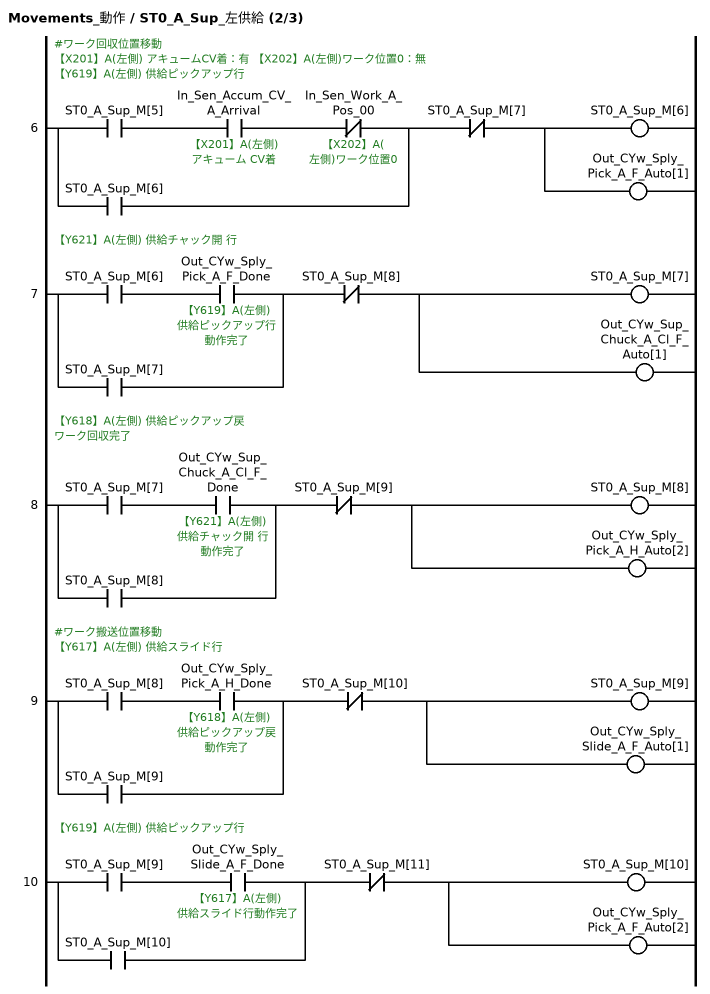
(* [picture p24: Movements_動作 / ST0_A_Sup_左供給, rungs 6-10] *)
(* Rung 6: #ワーク回収位置移動 / 【X201】A(左側) アキュームCV着：有 【X202】A(左側)ワーク位置0：無 / 【Y619】A(左側) 供給ピックアップ行 *)
_p20 := ((ST0_A_Sup_M[5] AND In_Sen_Accum_CV_A_Arrival AND NOT In_Sen_Work_A_Pos_00) OR ST0_A_Sup_M[6]) AND NOT ST0_A_Sup_M[7];
ST0_A_Sup_M[6] := _p20;
Out_CYw_Sply_Pick_A_F_Auto[1] := _p20;
(* Rung 7: 【Y621】A(左側) 供給チャック開 行 *)
_p21 := ((ST0_A_Sup_M[6] AND Out_CYw_Sply_Pick_A_F_Done) OR ST0_A_Sup_M[7]) AND NOT ST0_A_Sup_M[8];
ST0_A_Sup_M[7] := _p21;
Out_CYw_Sup_Chuck_A_Cl_F_Auto[1] := _p21;
(* Rung 8: 【Y618】A(左側) 供給ピックアップ戻 / ワーク回収完了 *)
_p22 := ((ST0_A_Sup_M[7] AND Out_CYw_Sup_Chuck_A_Cl_F_Done) OR ST0_A_Sup_M[8]) AND NOT ST0_A_Sup_M[9];
ST0_A_Sup_M[8] := _p22;
Out_CYw_Sply_Pick_A_H_Auto[2] := _p22;
(* Rung 9: #ワーク搬送位置移動 / 【Y617】A(左側) 供給スライド行 *)
_p23 := ((ST0_A_Sup_M[8] AND Out_CYw_Sply_Pick_A_H_Done) OR ST0_A_Sup_M[9]) AND NOT ST0_A_Sup_M[10];
ST0_A_Sup_M[9] := _p23;
Out_CYw_Sply_Slide_A_F_Auto[1] := _p23;
(* Rung 10: 【Y619】A(左側) 供給ピックアップ行 *)
_p24 := ((ST0_A_Sup_M[9] AND Out_CYw_Sply_Slide_A_F_Done) OR ST0_A_Sup_M[10]) AND NOT ST0_A_Sup_M[11];
ST0_A_Sup_M[10] := _p24;
Out_CYw_Sply_Pick_A_F_Auto[2] := _p24;

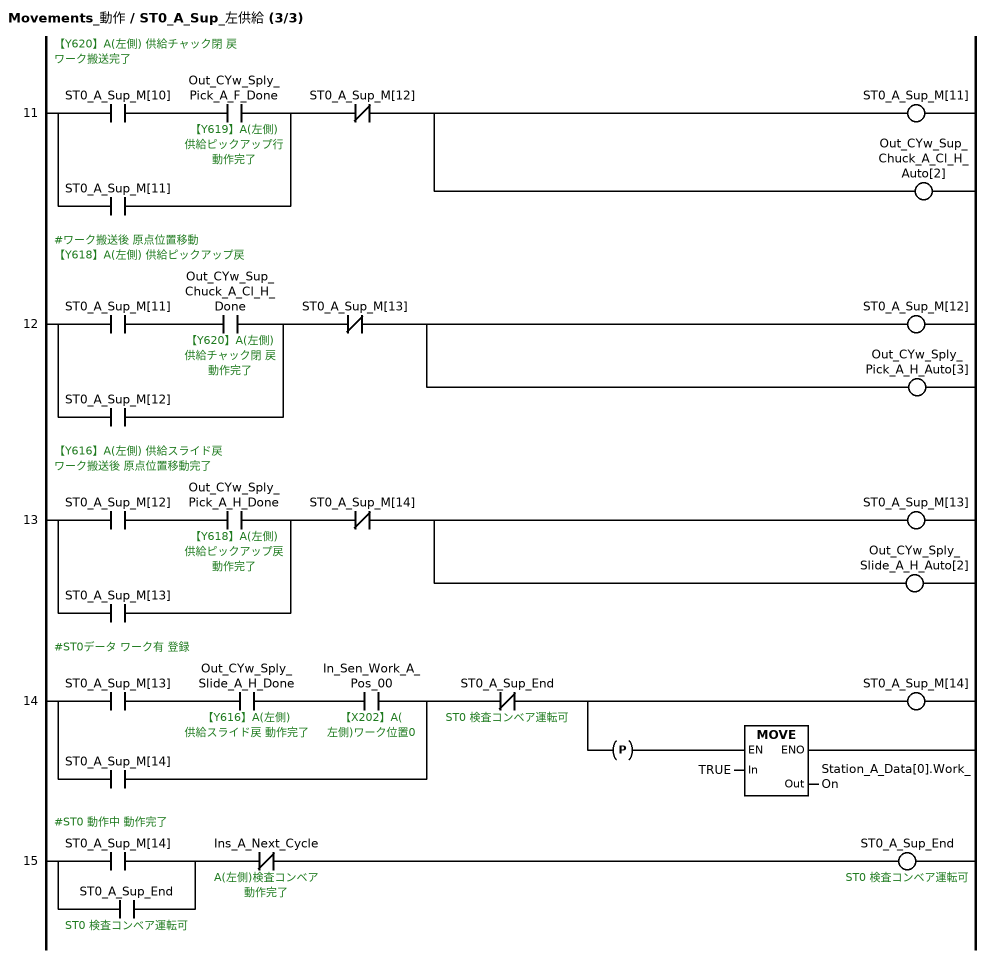
(* Rung 11: 【Y620】A(左側) 供給チャック閉 戻 / ワーク搬送完了 *)
_p25 := ((ST0_A_Sup_M[10] AND Out_CYw_Sply_Pick_A_F_Done) OR ST0_A_Sup_M[11]) AND NOT ST0_A_Sup_M[12];
ST0_A_Sup_M[11] := _p25;
Out_CYw_Sup_Chuck_A_Cl_H_Auto[2] := _p25;
(* Rung 12: #ワーク搬送後 原点位置移動 / 【Y618】A(左側) 供給ピックアップ戻 *)
_p26 := ((ST0_A_Sup_M[11] AND Out_CYw_Sup_Chuck_A_Cl_H_Done) OR ST0_A_Sup_M[12]) AND NOT ST0_A_Sup_M[13];
ST0_A_Sup_M[12] := _p26;
Out_CYw_Sply_Pick_A_H_Auto[3] := _p26;
(* Rung 13: 【Y616】A(左側) 供給スライド戻 / ワーク搬送後 原点位置移動完了 *)
_p27 := ((ST0_A_Sup_M[12] AND Out_CYw_Sply_Pick_A_H_Done) OR ST0_A_Sup_M[13]) AND NOT ST0_A_Sup_M[14];
ST0_A_Sup_M[13] := _p27;
Out_CYw_Sply_Slide_A_H_Auto[2] := _p27;
(* Rung 14: #ST0データ ワーク有 登録 *)
_p28 := ((ST0_A_Sup_M[13] AND Out_CYw_Sply_Slide_A_H_Done AND In_Sen_Work_A_Pos_00) OR ST0_A_Sup_M[14]) AND NOT ST0_A_Sup_End;
ST0_A_Sup_M[14] := _p28;
_e29(CLK := _p28);
IF _e29.Q THEN Station_A_Data[0].Work_On := TRUE; END_IF;
(* Rung 15: #ST0 動作中 動作完了 *)
ST0_A_Sup_End := (ST0_A_Sup_M[14] OR ST0_A_Sup_End) AND NOT Ins_A_Next_Cycle;

(* Section ST1_A_Ca1_左Ca1検査: ladder, written here as Structured Text *)

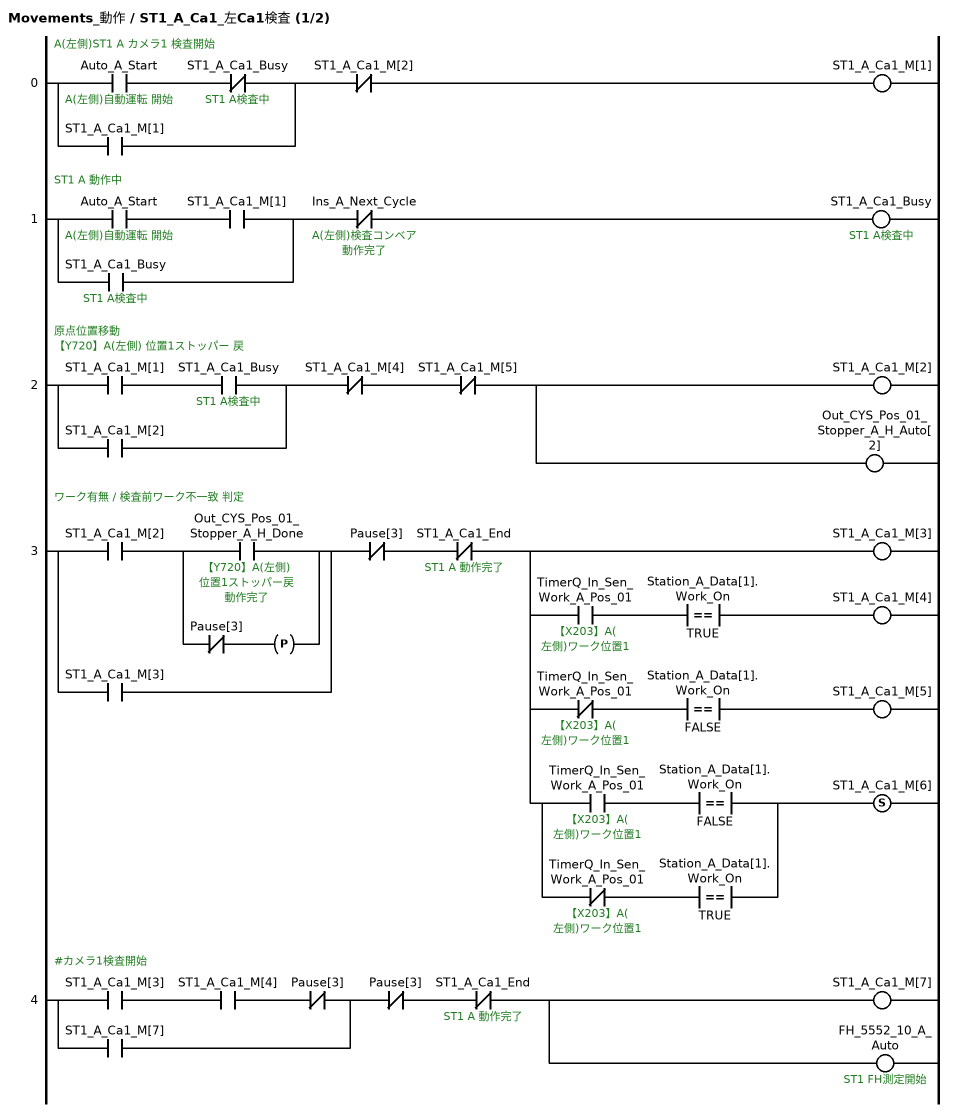
(* Rung 0: A(左側)ST1 A カメラ1 検査開始 *)
ST1_A_Ca1_M[1] := ((Auto_A_Start AND NOT ST1_A_Ca1_Busy) OR ST1_A_Ca1_M[1]) AND NOT ST1_A_Ca1_M[2];
(* Rung 1: ST1 A 動作中 *)
ST1_A_Ca1_Busy := ((Auto_A_Start AND ST1_A_Ca1_M[1]) OR ST1_A_Ca1_Busy) AND NOT Ins_A_Next_Cycle;
(* Rung 2: 原点位置移動 / 【Y720】A(左側) 位置1ストッパー 戻 *)
_p30 := ((ST1_A_Ca1_M[1] AND ST1_A_Ca1_Busy) OR ST1_A_Ca1_M[2]) AND NOT ST1_A_Ca1_M[4] AND NOT ST1_A_Ca1_M[5];
ST1_A_Ca1_M[2] := _p30;
Out_CYS_Pos_01_Stopper_A_H_Auto[2] := _p30;
(* Rung 3: ワーク有無 / 検査前ワーク不一致 判定 *)
_e31(CLK := ST1_A_Ca1_M[2] AND NOT Pause[3]);
_p32 := ((ST1_A_Ca1_M[2] AND Out_CYS_Pos_01_Stopper_A_H_Done) OR _e31.Q OR ST1_A_Ca1_M[3]) AND NOT Pause[3] AND NOT ST1_A_Ca1_End;
ST1_A_Ca1_M[3] := _p32;
ST1_A_Ca1_M[4] := _p32 AND TimerQ_In_Sen_Work_A_Pos_01 AND (Station_A_Data[1].Work_On = TRUE);
ST1_A_Ca1_M[5] := _p32 AND NOT TimerQ_In_Sen_Work_A_Pos_01 AND (Station_A_Data[1].Work_On = FALSE);
IF _p32 AND ((TimerQ_In_Sen_Work_A_Pos_01 AND (Station_A_Data[1].Work_On = FALSE)) OR (NOT TimerQ_In_Sen_Work_A_Pos_01 AND (Station_A_Data[1].Work_On = TRUE))) THEN
    ST1_A_Ca1_M[6] := TRUE;
END_IF;
(* Rung 4: #カメラ1検査開始 *)
_p33 := ((ST1_A_Ca1_M[3] AND ST1_A_Ca1_M[4] AND NOT Pause[3]) OR ST1_A_Ca1_M[7]) AND NOT Pause[3] AND NOT ST1_A_Ca1_End;
ST1_A_Ca1_M[7] := _p33;
FH_5552_10_A_Auto := _p33;

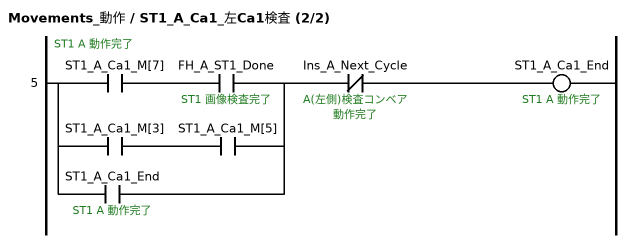
(* Rung 5: ST1 A 動作完了 *)
ST1_A_Ca1_End := ((ST1_A_Ca1_M[7] AND FH_A_ST1_Done) OR (ST1_A_Ca1_M[3] AND ST1_A_Ca1_M[5]) OR ST1_A_Ca1_End) AND NOT Ins_A_Next_Cycle;

(* Section ST2_A_Hgt_左高さ検査: ladder, written here as Structured Text *)

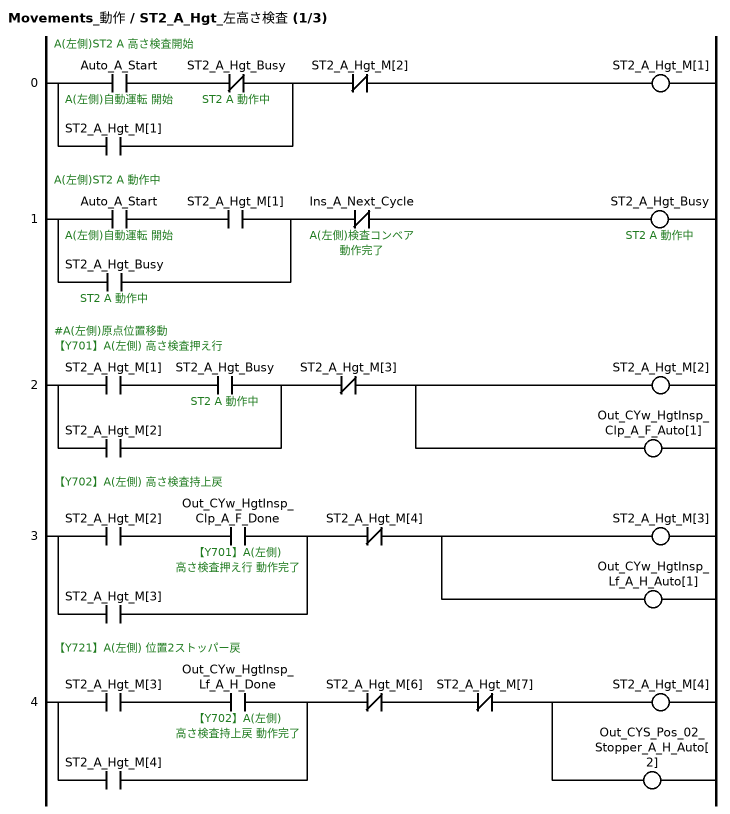
(* Rung 0: A(左側)ST2 A 高さ検査開始 *)
ST2_A_Hgt_M[1] := ((Auto_A_Start AND NOT ST2_A_Hgt_Busy) OR ST2_A_Hgt_M[1]) AND NOT ST2_A_Hgt_M[2];
(* Rung 1: A(左側)ST2 A 動作中 *)
ST2_A_Hgt_Busy := ((Auto_A_Start AND ST2_A_Hgt_M[1]) OR ST2_A_Hgt_Busy) AND NOT Ins_A_Next_Cycle;
(* Rung 2: #A(左側)原点位置移動 / 【Y701】A(左側) 高さ検査押え行 *)
_p34 := ((ST2_A_Hgt_M[1] AND ST2_A_Hgt_Busy) OR ST2_A_Hgt_M[2]) AND NOT ST2_A_Hgt_M[3];
ST2_A_Hgt_M[2] := _p34;
Out_CYw_HgtInsp_Clp_A_F_Auto[1] := _p34;
(* Rung 3: 【Y702】A(左側) 高さ検査持上戻 *)
_p35 := ((ST2_A_Hgt_M[2] AND Out_CYw_HgtInsp_Clp_A_F_Done) OR ST2_A_Hgt_M[3]) AND NOT ST2_A_Hgt_M[4];
ST2_A_Hgt_M[3] := _p35;
Out_CYw_HgtInsp_Lf_A_H_Auto[1] := _p35;
(* Rung 4: 【Y721】A(左側) 位置2ストッパー戻 *)
_p36 := ((ST2_A_Hgt_M[3] AND Out_CYw_HgtInsp_Lf_A_H_Done) OR ST2_A_Hgt_M[4]) AND NOT ST2_A_Hgt_M[6] AND NOT ST2_A_Hgt_M[7];
ST2_A_Hgt_M[4] := _p36;
Out_CYS_Pos_02_Stopper_A_H_Auto[2] := _p36;

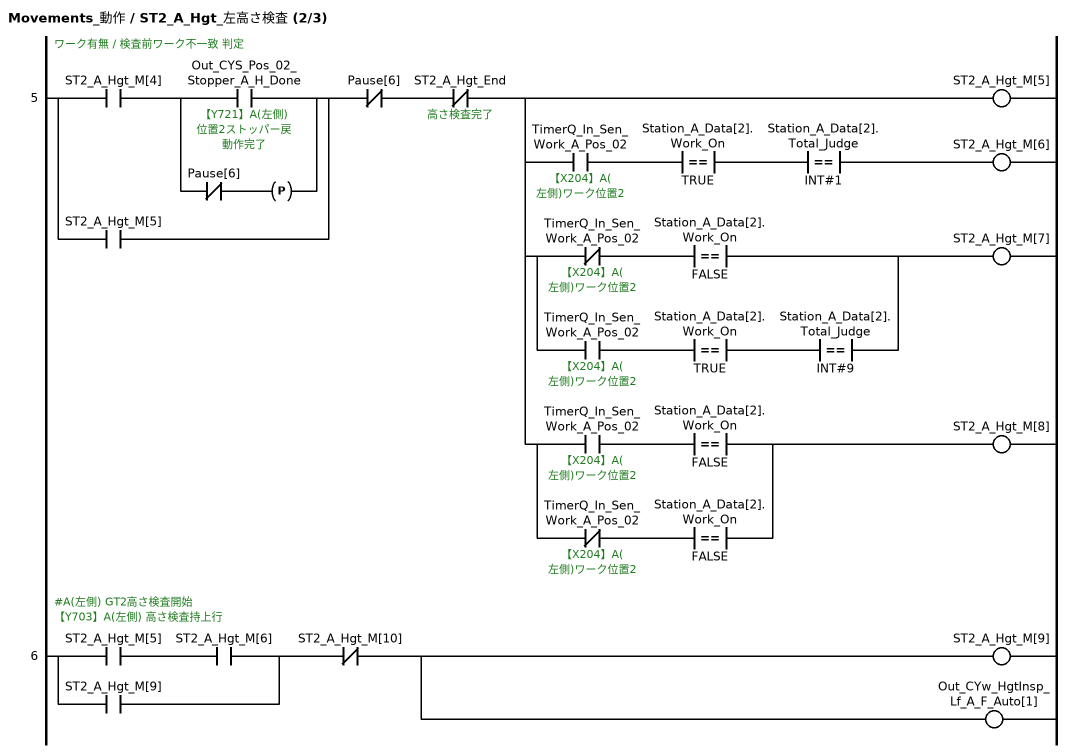
(* Rung 5: ワーク有無 / 検査前ワーク不一致 判定 *)
_e37(CLK := ST2_A_Hgt_M[4] AND NOT Pause[6]);
_p38 := ((ST2_A_Hgt_M[4] AND Out_CYS_Pos_02_Stopper_A_H_Done) OR _e37.Q OR ST2_A_Hgt_M[5]) AND NOT Pause[6] AND NOT ST2_A_Hgt_End;
ST2_A_Hgt_M[5] := _p38;
ST2_A_Hgt_M[6] := _p38 AND TimerQ_In_Sen_Work_A_Pos_02 AND (Station_A_Data[2].Work_On = TRUE) AND (Station_A_Data[2].Total_Judge = INT#1);
ST2_A_Hgt_M[7] := _p38 AND ((NOT TimerQ_In_Sen_Work_A_Pos_02 AND (Station_A_Data[2].Work_On = FALSE)) OR (TimerQ_In_Sen_Work_A_Pos_02 AND (Station_A_Data[2].Work_On = TRUE) AND (Station_A_Data[2].Total_Judge = INT#9)));
ST2_A_Hgt_M[8] := _p38 AND ((TimerQ_In_Sen_Work_A_Pos_02 AND (Station_A_Data[2].Work_On = FALSE)) OR (NOT TimerQ_In_Sen_Work_A_Pos_02 AND (Station_A_Data[2].Work_On = FALSE)));
(* Rung 6: #A(左側) GT2高さ検査開始 / 【Y703】A(左側) 高さ検査持上行 *)
_p39 := ((ST2_A_Hgt_M[5] AND ST2_A_Hgt_M[6]) OR ST2_A_Hgt_M[9]) AND NOT ST2_A_Hgt_M[10];
ST2_A_Hgt_M[9] := _p39;
Out_CYw_HgtInsp_Lf_A_F_Auto[1] := _p39;

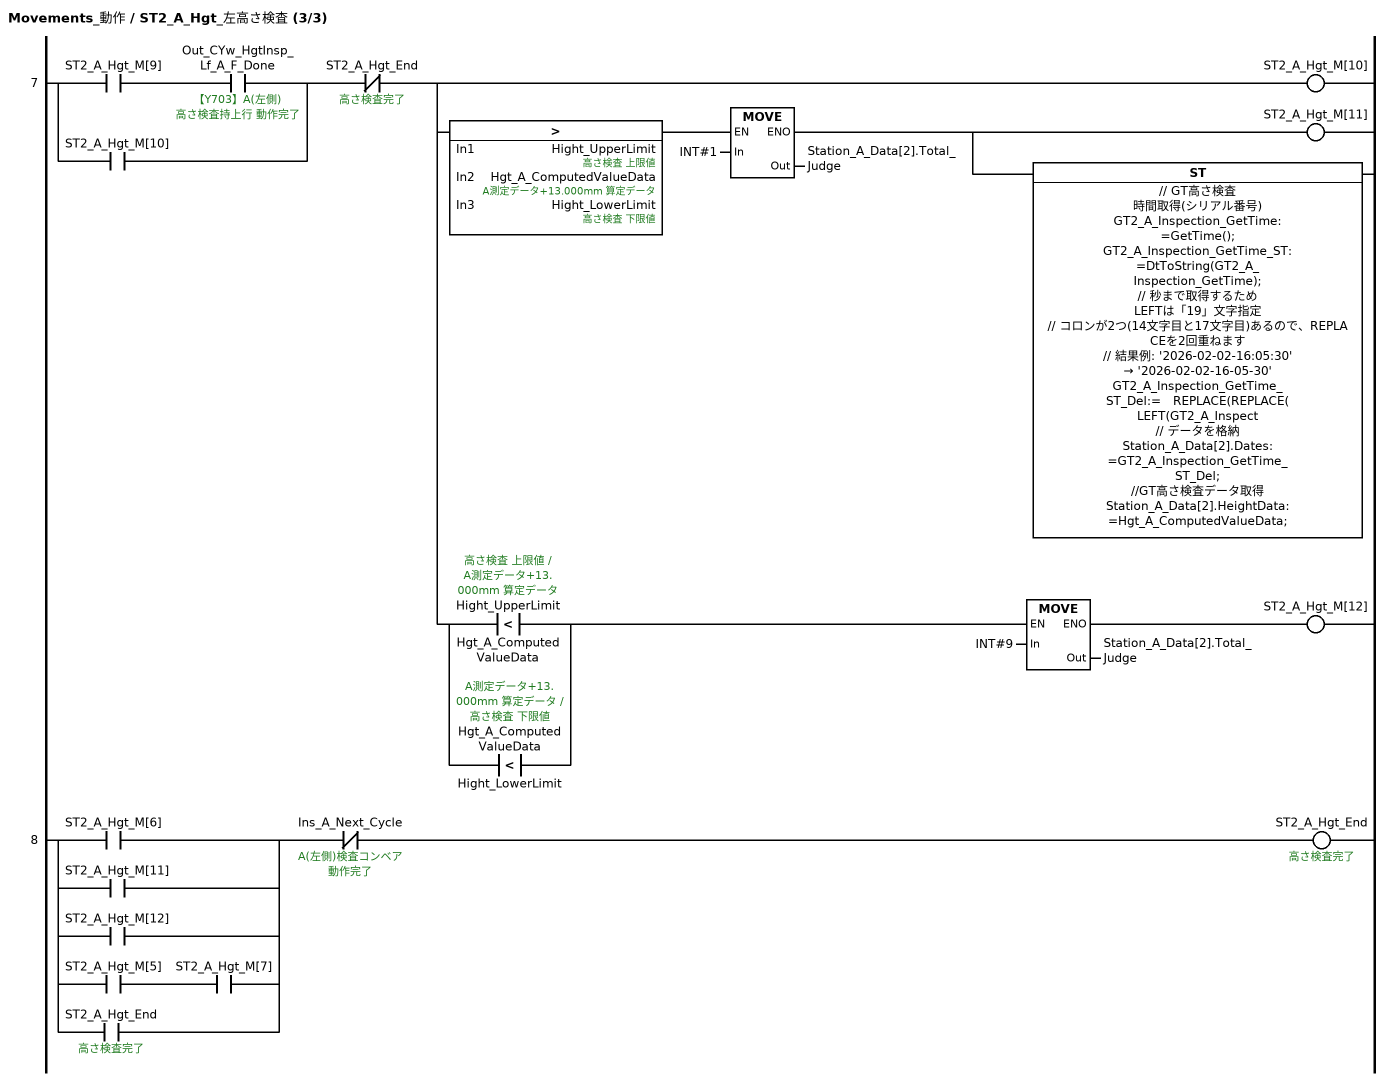
(* Rung 7 *)
_p40 := ((ST2_A_Hgt_M[9] AND Out_CYw_HgtInsp_Lf_A_F_Done) OR ST2_A_Hgt_M[10]) AND NOT ST2_A_Hgt_End;
ST2_A_Hgt_M[10] := _p40;
IF _p40 AND GT(Hight_UpperLimit, Hgt_A_ComputedValueData, Hight_LowerLimit) THEN
    Station_A_Data[2].Total_Judge := INT#1;
END_IF;
_p41 := _p40 AND GT(Hight_UpperLimit, Hgt_A_ComputedValueData, Hight_LowerLimit);
ST2_A_Hgt_M[11] := _p41;
IF _p41 THEN
    // GT高さ検査 時間取得(シリアル番号)
    GT2_A_Inspection_GetTime:=GetTime();
    GT2_A_Inspection_GetTime_ST:=DtToString(GT2_A_Inspection_GetTime);
    // 秒まで取得するため LEFTは「19」文字指定
    // コロンが2つ(14文字目と17文字目)あるので、REPLACEを2回重ねます
    // 結果例: '2026-02-02-16:05:30' → '2026-02-02-16-05-30'
    GT2_A_Inspection_GetTime_ST_Del:=   REPLACE(REPLACE(LEFT(GT2_A_Inspection_GetTime_ST, UINT#19), STRING#'-', UINT#1, UINT#17), STRING#'-', UINT#1, UINT#14);
    // データを格納
    Station_A_Data[2].Dates:=GT2_A_Inspection_GetTime_ST_Del;
    //GT高さ検査データ取得
    Station_A_Data[2].HeightData:=Hgt_A_ComputedValueData;
END_IF;
IF _p40 AND ((Hight_UpperLimit < Hgt_A_ComputedValueData) OR (Hgt_A_ComputedValueData < Hight_LowerLimit)) THEN
    Station_A_Data[2].Total_Judge := INT#9;
END_IF;
ST2_A_Hgt_M[12] := _p40 AND ((Hight_UpperLimit < Hgt_A_ComputedValueData) OR (Hgt_A_ComputedValueData < Hight_LowerLimit));
(* Rung 8 *)
ST2_A_Hgt_End := (ST2_A_Hgt_M[6] OR ST2_A_Hgt_M[11] OR ST2_A_Hgt_M[12] OR (ST2_A_Hgt_M[5] AND ST2_A_Hgt_M[7]) OR ST2_A_Hgt_End) AND NOT Ins_A_Next_Cycle;

(* Section ST3_A_Dis1_左NG1排出: ladder, written here as Structured Text *)

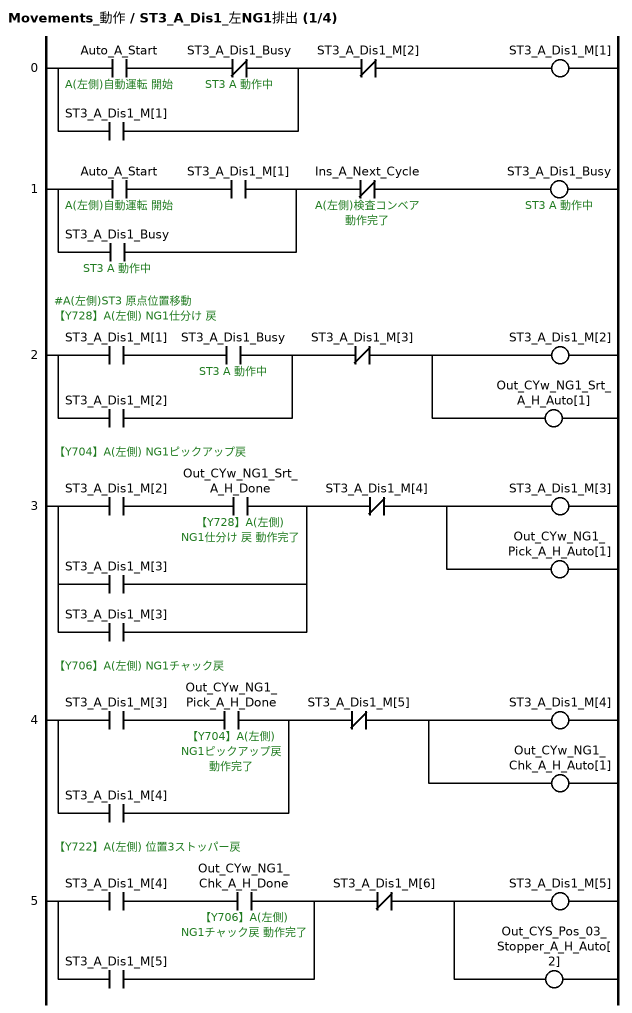
(* Rung 0 *)
ST3_A_Dis1_M[1] := ((Auto_A_Start AND NOT ST3_A_Dis1_Busy) OR ST3_A_Dis1_M[1]) AND NOT ST3_A_Dis1_M[2];
(* Rung 1 *)
ST3_A_Dis1_Busy := ((Auto_A_Start AND ST3_A_Dis1_M[1]) OR ST3_A_Dis1_Busy) AND NOT Ins_A_Next_Cycle;
(* Rung 2: #A(左側)ST3 原点位置移動 / 【Y728】A(左側) NG1仕分け 戻 *)
_p42 := ((ST3_A_Dis1_M[1] AND ST3_A_Dis1_Busy) OR ST3_A_Dis1_M[2]) AND NOT ST3_A_Dis1_M[3];
ST3_A_Dis1_M[2] := _p42;
Out_CYw_NG1_Srt_A_H_Auto[1] := _p42;
(* Rung 3: 【Y704】A(左側) NG1ピックアップ戻 *)
_p43 := ((ST3_A_Dis1_M[2] AND Out_CYw_NG1_Srt_A_H_Done) OR ST3_A_Dis1_M[3] OR ST3_A_Dis1_M[3]) AND NOT ST3_A_Dis1_M[4];
ST3_A_Dis1_M[3] := _p43;
Out_CYw_NG1_Pick_A_H_Auto[1] := _p43;
(* Rung 4: 【Y706】A(左側) NG1チャック戻 *)
_p44 := ((ST3_A_Dis1_M[3] AND Out_CYw_NG1_Pick_A_H_Done) OR ST3_A_Dis1_M[4]) AND NOT ST3_A_Dis1_M[5];
ST3_A_Dis1_M[4] := _p44;
Out_CYw_NG1_Chk_A_H_Auto[1] := _p44;
(* Rung 5: 【Y722】A(左側) 位置3ストッパー戻 *)
_p45 := ((ST3_A_Dis1_M[4] AND Out_CYw_NG1_Chk_A_H_Done) OR ST3_A_Dis1_M[5]) AND NOT ST3_A_Dis1_M[6];
ST3_A_Dis1_M[5] := _p45;
Out_CYS_Pos_03_Stopper_A_H_Auto[2] := _p45;

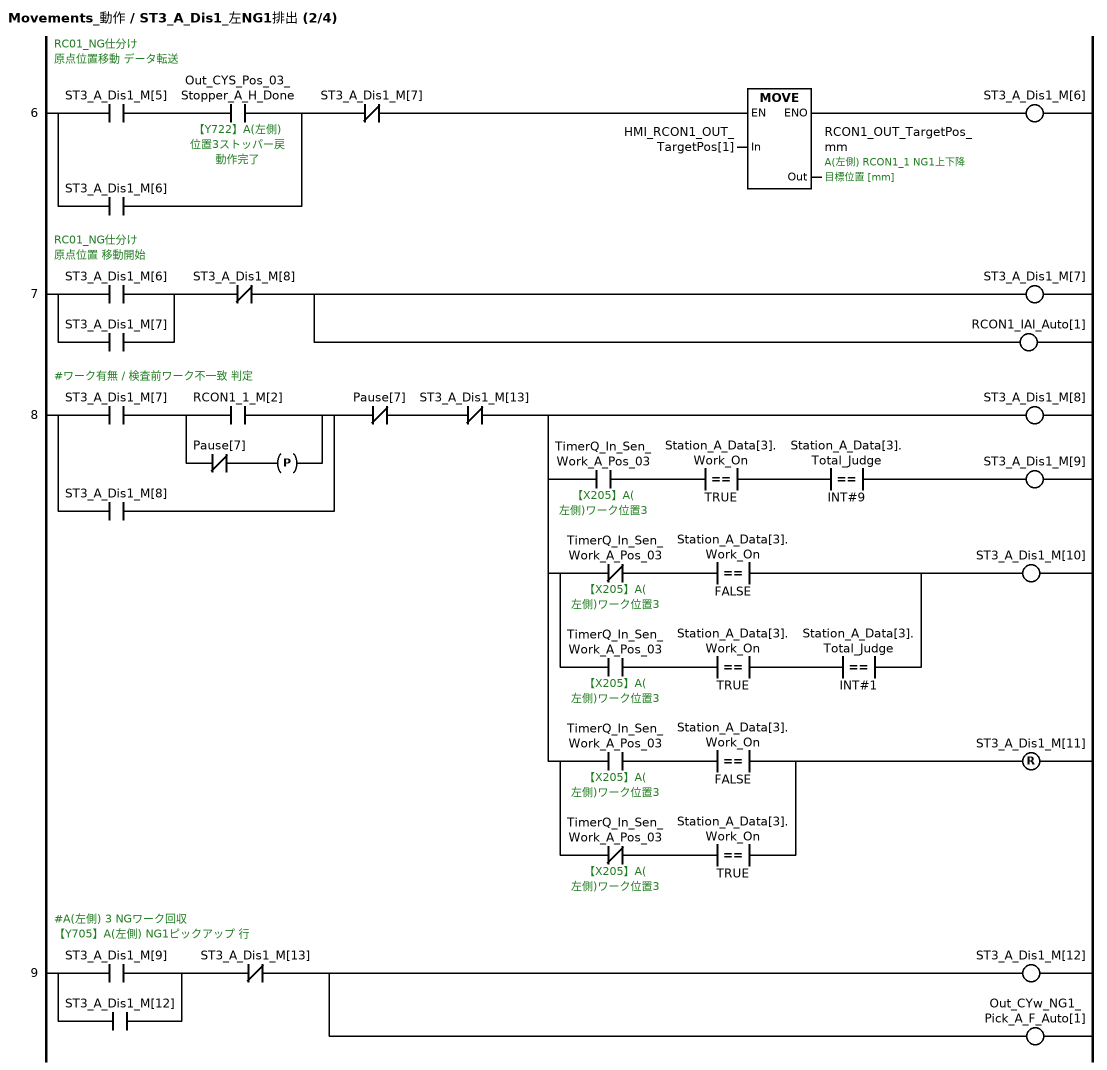
(* Rung 6: RC01_NG仕分け / 原点位置移動 データ転送 *)
IF ((ST3_A_Dis1_M[5] AND Out_CYS_Pos_03_Stopper_A_H_Done) OR ST3_A_Dis1_M[6]) AND NOT ST3_A_Dis1_M[7] THEN
    RCON1_OUT_TargetPos_mm := HMI_RCON1_OUT_TargetPos[1];
END_IF;
ST3_A_Dis1_M[6] := ((ST3_A_Dis1_M[5] AND Out_CYS_Pos_03_Stopper_A_H_Done) OR ST3_A_Dis1_M[6]) AND NOT ST3_A_Dis1_M[7];
(* Rung 7: RC01_NG仕分け / 原点位置 移動開始 *)
_p46 := (ST3_A_Dis1_M[6] OR ST3_A_Dis1_M[7]) AND NOT ST3_A_Dis1_M[8];
ST3_A_Dis1_M[7] := _p46;
RCON1_IAI_Auto[1] := _p46;
(* Rung 8: #ワーク有無 / 検査前ワーク不一致 判定 *)
_e47(CLK := ST3_A_Dis1_M[7] AND NOT Pause[7]);
_p48 := ((ST3_A_Dis1_M[7] AND RCON1_1_M[2]) OR _e47.Q OR ST3_A_Dis1_M[8]) AND NOT Pause[7] AND NOT ST3_A_Dis1_M[13];
ST3_A_Dis1_M[8] := _p48;
ST3_A_Dis1_M[9] := _p48 AND TimerQ_In_Sen_Work_A_Pos_03 AND (Station_A_Data[3].Work_On = TRUE) AND (Station_A_Data[3].Total_Judge = INT#9);
ST3_A_Dis1_M[10] := _p48 AND ((NOT TimerQ_In_Sen_Work_A_Pos_03 AND (Station_A_Data[3].Work_On = FALSE)) OR (TimerQ_In_Sen_Work_A_Pos_03 AND (Station_A_Data[3].Work_On = TRUE) AND (Station_A_Data[3].Total_Judge = INT#1)));
IF _p48 AND ((TimerQ_In_Sen_Work_A_Pos_03 AND (Station_A_Data[3].Work_On = FALSE)) OR (NOT TimerQ_In_Sen_Work_A_Pos_03 AND (Station_A_Data[3].Work_On = TRUE))) THEN
    ST3_A_Dis1_M[11] := FALSE;
END_IF;
(* Rung 9: #A(左側) 3 NGワーク回収 / 【Y705】A(左側) NG1ピックアップ 行 *)
_p49 := (ST3_A_Dis1_M[9] OR ST3_A_Dis1_M[12]) AND NOT ST3_A_Dis1_M[13];
ST3_A_Dis1_M[12] := _p49;
Out_CYw_NG1_Pick_A_F_Auto[1] := _p49;

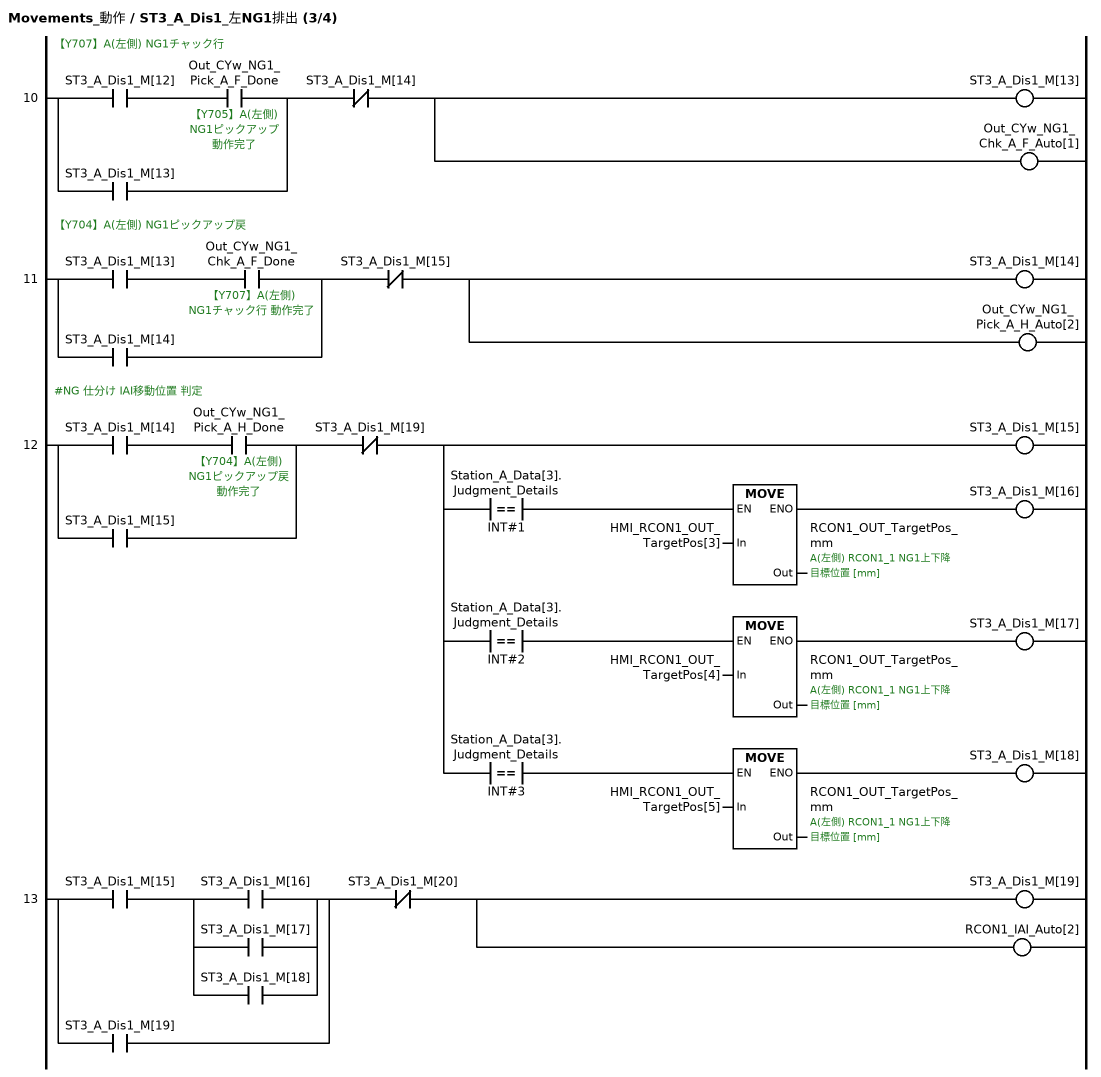
(* Rung 10: 【Y707】A(左側) NG1チャック行 *)
_p50 := ((ST3_A_Dis1_M[12] AND Out_CYw_NG1_Pick_A_F_Done) OR ST3_A_Dis1_M[13]) AND NOT ST3_A_Dis1_M[14];
ST3_A_Dis1_M[13] := _p50;
Out_CYw_NG1_Chk_A_F_Auto[1] := _p50;
(* Rung 11: 【Y704】A(左側) NG1ピックアップ戻 *)
_p51 := ((ST3_A_Dis1_M[13] AND Out_CYw_NG1_Chk_A_F_Done) OR ST3_A_Dis1_M[14]) AND NOT ST3_A_Dis1_M[15];
ST3_A_Dis1_M[14] := _p51;
Out_CYw_NG1_Pick_A_H_Auto[2] := _p51;
(* Rung 12: #NG 仕分け IAI移動位置 判定 *)
_p52 := ((ST3_A_Dis1_M[14] AND Out_CYw_NG1_Pick_A_H_Done) OR ST3_A_Dis1_M[15]) AND NOT ST3_A_Dis1_M[19];
ST3_A_Dis1_M[15] := _p52;
IF _p52 AND (Station_A_Data[3].Judgment_Details = INT#1) THEN
    RCON1_OUT_TargetPos_mm := HMI_RCON1_OUT_TargetPos[3];
END_IF;
ST3_A_Dis1_M[16] := _p52 AND (Station_A_Data[3].Judgment_Details = INT#1);
IF _p52 AND (Station_A_Data[3].Judgment_Details = INT#2) THEN
    RCON1_OUT_TargetPos_mm := HMI_RCON1_OUT_TargetPos[4];
END_IF;
ST3_A_Dis1_M[17] := _p52 AND (Station_A_Data[3].Judgment_Details = INT#2);
IF _p52 AND (Station_A_Data[3].Judgment_Details = INT#3) THEN
    RCON1_OUT_TargetPos_mm := HMI_RCON1_OUT_TargetPos[5];
END_IF;
ST3_A_Dis1_M[18] := _p52 AND (Station_A_Data[3].Judgment_Details = INT#3);
(* Rung 13 *)
_p53 := ((ST3_A_Dis1_M[15] AND (ST3_A_Dis1_M[16] OR ST3_A_Dis1_M[17] OR ST3_A_Dis1_M[18])) OR ST3_A_Dis1_M[19]) AND NOT ST3_A_Dis1_M[20];
ST3_A_Dis1_M[19] := _p53;
RCON1_IAI_Auto[2] := _p53;

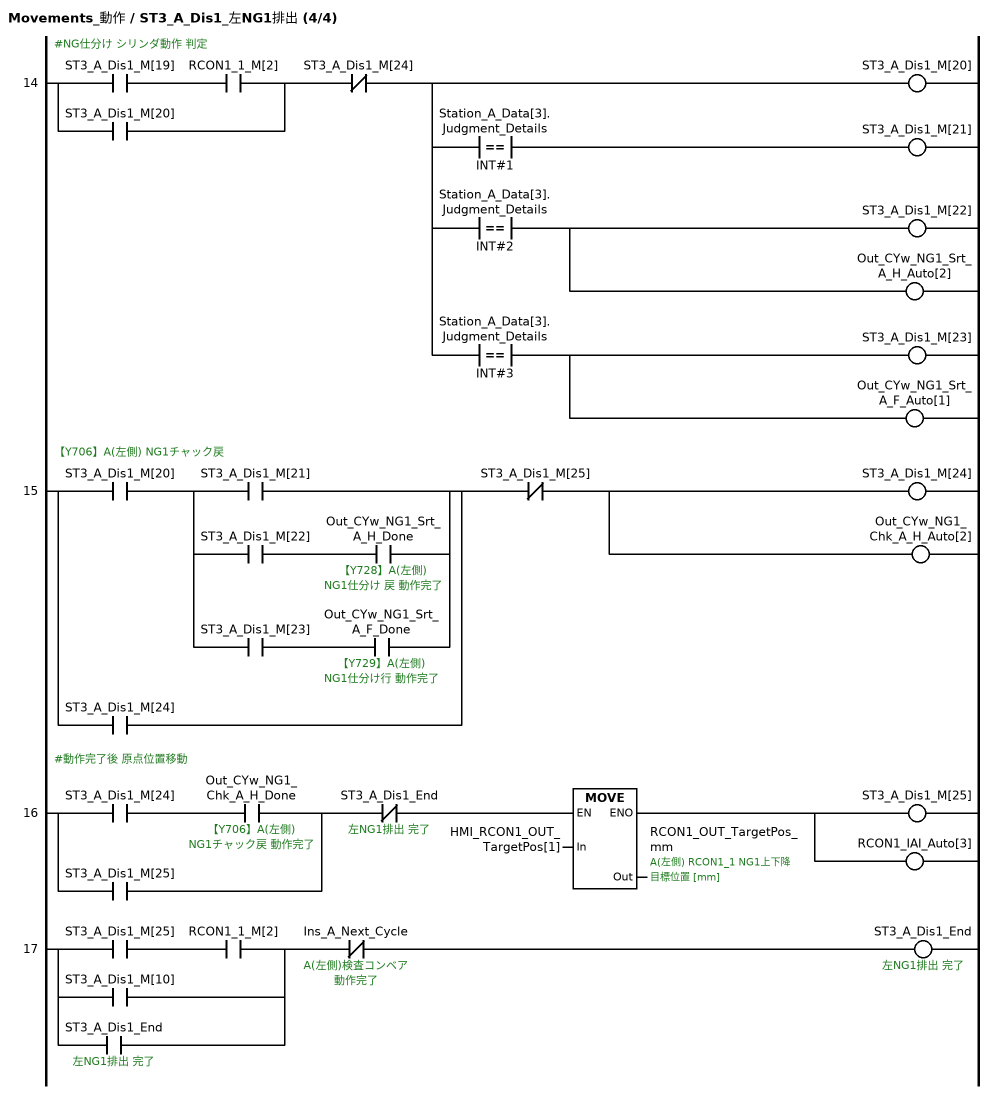
(* Rung 14: #NG仕分け シリンダ動作 判定 *)
_p54 := ((ST3_A_Dis1_M[19] AND RCON1_1_M[2]) OR ST3_A_Dis1_M[20]) AND NOT ST3_A_Dis1_M[24];
ST3_A_Dis1_M[20] := _p54;
ST3_A_Dis1_M[21] := _p54 AND (Station_A_Data[3].Judgment_Details = INT#1);
_p55 := _p54 AND (Station_A_Data[3].Judgment_Details = INT#2);
ST3_A_Dis1_M[22] := _p55;
Out_CYw_NG1_Srt_A_H_Auto[2] := _p55;
_p56 := _p54 AND (Station_A_Data[3].Judgment_Details = INT#3);
ST3_A_Dis1_M[23] := _p56;
Out_CYw_NG1_Srt_A_F_Auto[1] := _p56;
(* Rung 15: 【Y706】A(左側) NG1チャック戻 *)
_p57 := ((ST3_A_Dis1_M[20] AND (ST3_A_Dis1_M[21] OR (ST3_A_Dis1_M[22] AND Out_CYw_NG1_Srt_A_H_Done) OR (ST3_A_Dis1_M[23] AND Out_CYw_NG1_Srt_A_F_Done))) OR ST3_A_Dis1_M[24]) AND NOT ST3_A_Dis1_M[25];
ST3_A_Dis1_M[24] := _p57;
Out_CYw_NG1_Chk_A_H_Auto[2] := _p57;
(* Rung 16: #動作完了後 原点位置移動 *)
IF ((ST3_A_Dis1_M[24] AND Out_CYw_NG1_Chk_A_H_Done) OR ST3_A_Dis1_M[25]) AND NOT ST3_A_Dis1_End THEN
    RCON1_OUT_TargetPos_mm := HMI_RCON1_OUT_TargetPos[1];
END_IF;
_p58 := ((ST3_A_Dis1_M[24] AND Out_CYw_NG1_Chk_A_H_Done) OR ST3_A_Dis1_M[25]) AND NOT ST3_A_Dis1_End;
ST3_A_Dis1_M[25] := _p58;
RCON1_IAI_Auto[3] := _p58;
(* Rung 17 *)
ST3_A_Dis1_End := ((ST3_A_Dis1_M[25] AND RCON1_1_M[2]) OR ST3_A_Dis1_M[10] OR ST3_A_Dis1_End) AND NOT Ins_A_Next_Cycle;

(* Section ST4_A_Rev1_左反転1: ladder, written here as Structured Text *)

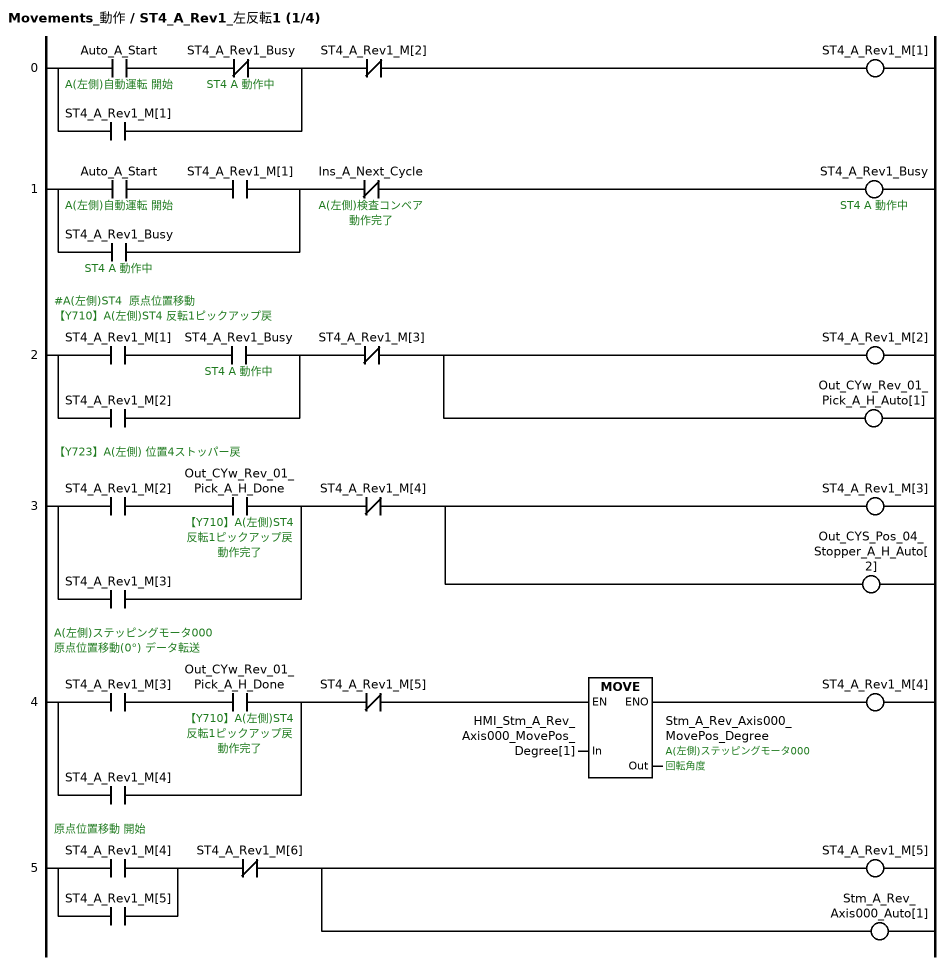
(* Rung 0 *)
ST4_A_Rev1_M[1] := ((Auto_A_Start AND NOT ST4_A_Rev1_Busy) OR ST4_A_Rev1_M[1]) AND NOT ST4_A_Rev1_M[2];
(* Rung 1 *)
ST4_A_Rev1_Busy := ((Auto_A_Start AND ST4_A_Rev1_M[1]) OR ST4_A_Rev1_Busy) AND NOT Ins_A_Next_Cycle;
(* Rung 2: #A(左側)ST4  原点位置移動 / 【Y710】A(左側)ST4 反転1ピックアップ戻 *)
_p59 := ((ST4_A_Rev1_M[1] AND ST4_A_Rev1_Busy) OR ST4_A_Rev1_M[2]) AND NOT ST4_A_Rev1_M[3];
ST4_A_Rev1_M[2] := _p59;
Out_CYw_Rev_01_Pick_A_H_Auto[1] := _p59;
(* Rung 3: 【Y723】A(左側) 位置4ストッパー戻 *)
_p60 := ((ST4_A_Rev1_M[2] AND Out_CYw_Rev_01_Pick_A_H_Done) OR ST4_A_Rev1_M[3]) AND NOT ST4_A_Rev1_M[4];
ST4_A_Rev1_M[3] := _p60;
Out_CYS_Pos_04_Stopper_A_H_Auto[2] := _p60;
(* Rung 4: A(左側)ステッピングモータ000 / 原点位置移動(0°) データ転送 *)
IF ((ST4_A_Rev1_M[3] AND Out_CYw_Rev_01_Pick_A_H_Done) OR ST4_A_Rev1_M[4]) AND NOT ST4_A_Rev1_M[5] THEN
    Stm_A_Rev_Axis000_MovePos_Degree := HMI_Stm_A_Rev_Axis000_MovePos_Degree[1];
END_IF;
ST4_A_Rev1_M[4] := ((ST4_A_Rev1_M[3] AND Out_CYw_Rev_01_Pick_A_H_Done) OR ST4_A_Rev1_M[4]) AND NOT ST4_A_Rev1_M[5];
(* Rung 5: 原点位置移動 開始 *)
_p61 := (ST4_A_Rev1_M[4] OR ST4_A_Rev1_M[5]) AND NOT ST4_A_Rev1_M[6];
ST4_A_Rev1_M[5] := _p61;
Stm_A_Rev_Axis000_Auto[1] := _p61;

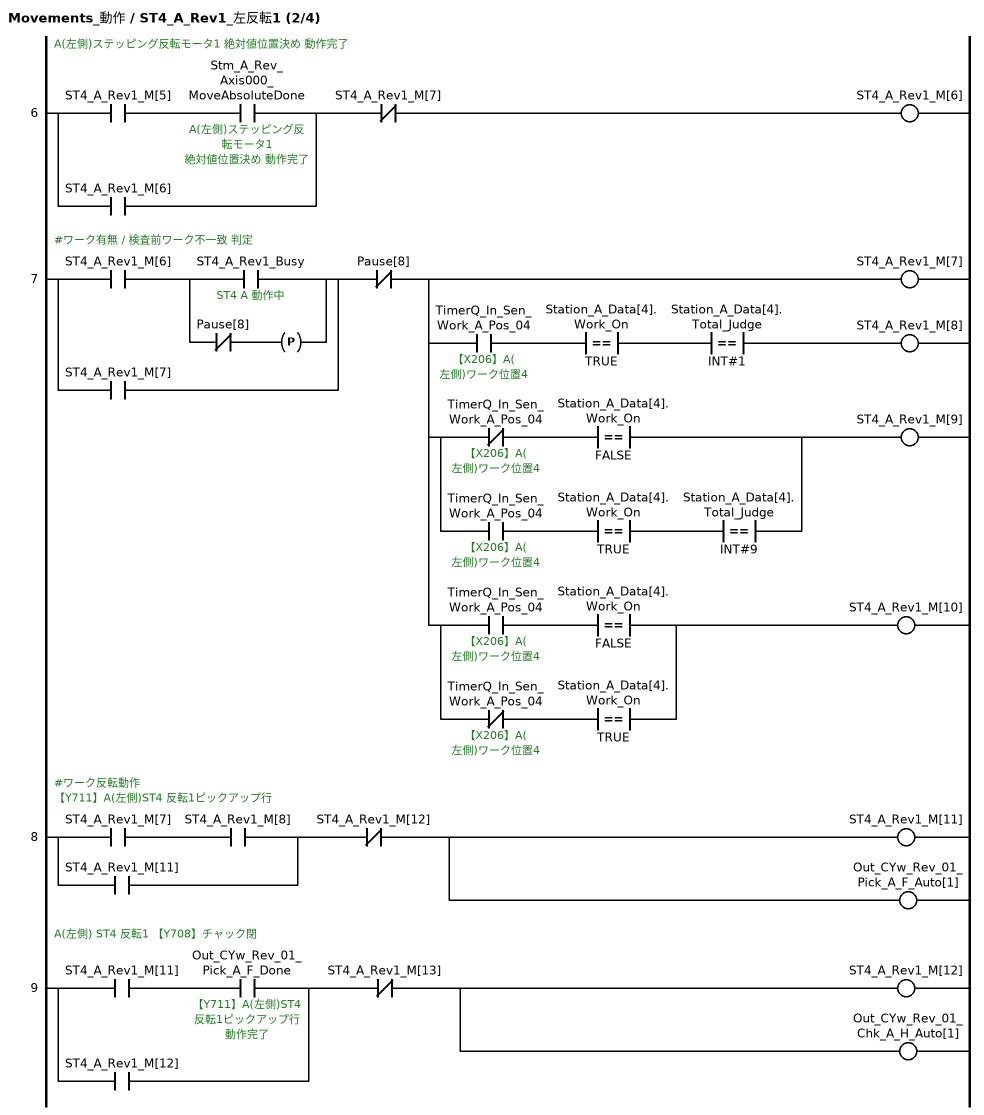
(* Rung 6: A(左側)ステッピング反転モータ1 絶対値位置決め 動作完了 *)
ST4_A_Rev1_M[6] := ((ST4_A_Rev1_M[5] AND Stm_A_Rev_Axis000_MoveAbsoluteDone) OR ST4_A_Rev1_M[6]) AND NOT ST4_A_Rev1_M[7];
(* Rung 7: #ワーク有無 / 検査前ワーク不一致 判定 *)
_e62(CLK := ST4_A_Rev1_M[6] AND NOT Pause[8]);
_p63 := ((ST4_A_Rev1_M[6] AND ST4_A_Rev1_Busy) OR _e62.Q OR ST4_A_Rev1_M[7]) AND NOT Pause[8];
ST4_A_Rev1_M[7] := _p63;
ST4_A_Rev1_M[8] := _p63 AND TimerQ_In_Sen_Work_A_Pos_04 AND (Station_A_Data[4].Work_On = TRUE) AND (Station_A_Data[4].Total_Judge = INT#1);
ST4_A_Rev1_M[9] := _p63 AND ((NOT TimerQ_In_Sen_Work_A_Pos_04 AND (Station_A_Data[4].Work_On = FALSE)) OR (TimerQ_In_Sen_Work_A_Pos_04 AND (Station_A_Data[4].Work_On = TRUE) AND (Station_A_Data[4].Total_Judge = INT#9)));
ST4_A_Rev1_M[10] := _p63 AND ((TimerQ_In_Sen_Work_A_Pos_04 AND (Station_A_Data[4].Work_On = FALSE)) OR (NOT TimerQ_In_Sen_Work_A_Pos_04 AND (Station_A_Data[4].Work_On = TRUE)));
(* Rung 8: #ワーク反転動作 / 【Y711】A(左側)ST4 反転1ピックアップ行 *)
_p64 := ((ST4_A_Rev1_M[7] AND ST4_A_Rev1_M[8]) OR ST4_A_Rev1_M[11]) AND NOT ST4_A_Rev1_M[12];
ST4_A_Rev1_M[11] := _p64;
Out_CYw_Rev_01_Pick_A_F_Auto[1] := _p64;
(* Rung 9: A(左側) ST4 反転1 【Y708】チャック閉 *)
_p65 := ((ST4_A_Rev1_M[11] AND Out_CYw_Rev_01_Pick_A_F_Done) OR ST4_A_Rev1_M[12]) AND NOT ST4_A_Rev1_M[13];
ST4_A_Rev1_M[12] := _p65;
Out_CYw_Rev_01_Chk_A_H_Auto[1] := _p65;

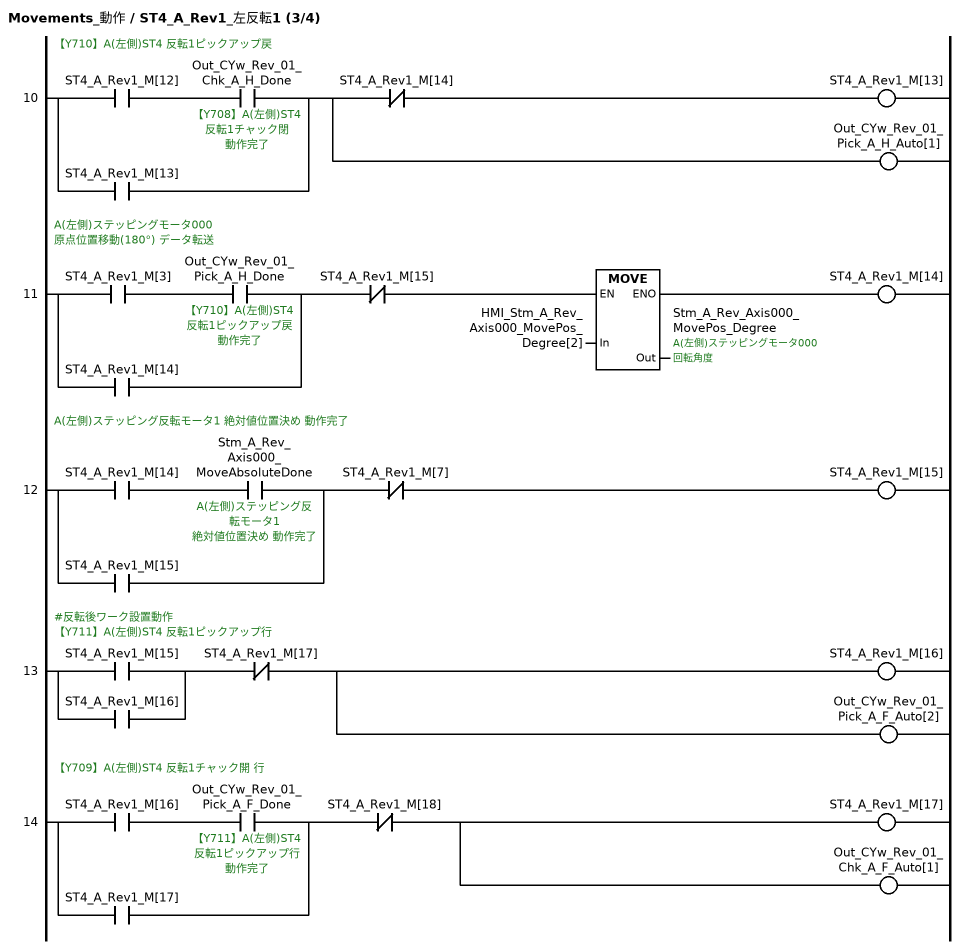
(* Rung 10: 【Y710】A(左側)ST4 反転1ピックアップ戻 *)
_p66 := (ST4_A_Rev1_M[12] AND Out_CYw_Rev_01_Chk_A_H_Done) OR ST4_A_Rev1_M[13];
ST4_A_Rev1_M[13] := _p66 AND NOT ST4_A_Rev1_M[14];
Out_CYw_Rev_01_Pick_A_H_Auto[1] := _p66;
(* Rung 11: A(左側)ステッピングモータ000 / 原点位置移動(180°) データ転送 *)
IF ((ST4_A_Rev1_M[3] AND Out_CYw_Rev_01_Pick_A_H_Done) OR ST4_A_Rev1_M[14]) AND NOT ST4_A_Rev1_M[15] THEN
    Stm_A_Rev_Axis000_MovePos_Degree := HMI_Stm_A_Rev_Axis000_MovePos_Degree[2];
END_IF;
ST4_A_Rev1_M[14] := ((ST4_A_Rev1_M[3] AND Out_CYw_Rev_01_Pick_A_H_Done) OR ST4_A_Rev1_M[14]) AND NOT ST4_A_Rev1_M[15];
(* Rung 12: A(左側)ステッピング反転モータ1 絶対値位置決め 動作完了 *)
ST4_A_Rev1_M[15] := ((ST4_A_Rev1_M[14] AND Stm_A_Rev_Axis000_MoveAbsoluteDone) OR ST4_A_Rev1_M[15]) AND NOT ST4_A_Rev1_M[7];
(* Rung 13: #反転後ワーク設置動作 / 【Y711】A(左側)ST4 反転1ピックアップ行 *)
_p67 := (ST4_A_Rev1_M[15] OR ST4_A_Rev1_M[16]) AND NOT ST4_A_Rev1_M[17];
ST4_A_Rev1_M[16] := _p67;
Out_CYw_Rev_01_Pick_A_F_Auto[2] := _p67;
(* Rung 14: 【Y709】A(左側)ST4 反転1チャック開 行 *)
_p68 := ((ST4_A_Rev1_M[16] AND Out_CYw_Rev_01_Pick_A_F_Done) OR ST4_A_Rev1_M[17]) AND NOT ST4_A_Rev1_M[18];
ST4_A_Rev1_M[17] := _p68;
Out_CYw_Rev_01_Chk_A_F_Auto[1] := _p68;

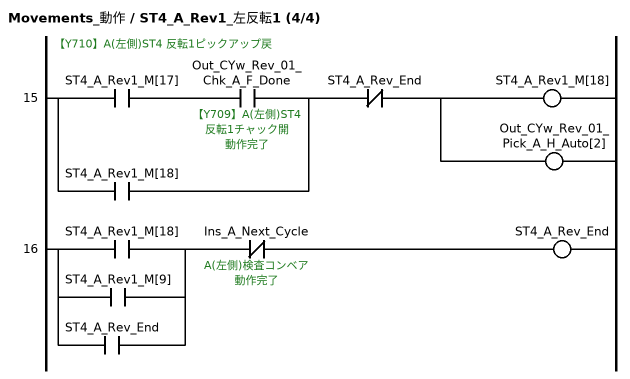
(* Rung 15: 【Y710】A(左側)ST4 反転1ピックアップ戻 *)
_p69 := ((ST4_A_Rev1_M[17] AND Out_CYw_Rev_01_Chk_A_F_Done) OR ST4_A_Rev1_M[18]) AND NOT ST4_A_Rev_End;
ST4_A_Rev1_M[18] := _p69;
Out_CYw_Rev_01_Pick_A_H_Auto[2] := _p69;
(* Rung 16 *)
ST4_A_Rev_End := (ST4_A_Rev1_M[18] OR ST4_A_Rev1_M[9] OR ST4_A_Rev_End) AND NOT Ins_A_Next_Cycle;

(* Section ST5_A_Ca2_左Ca2検査: ladder, written here as Structured Text *)

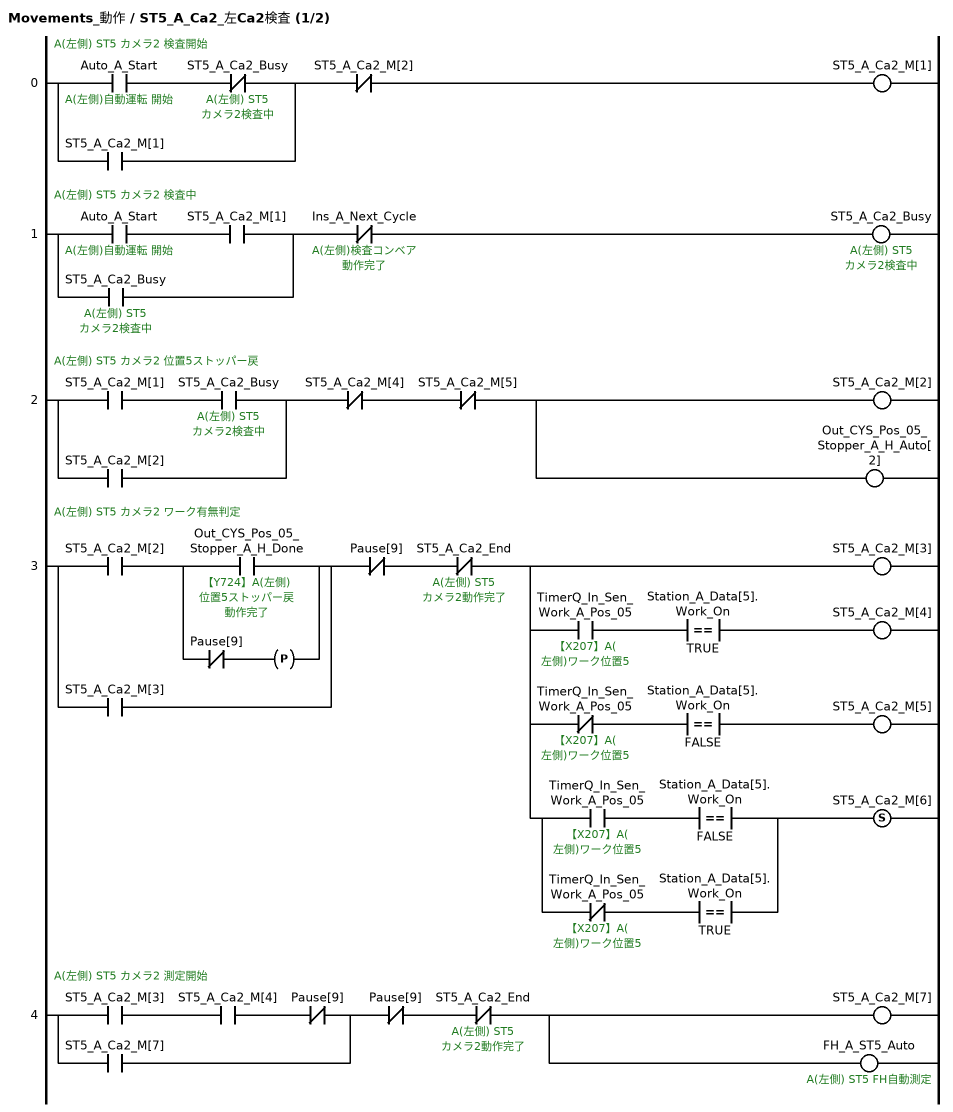
(* Rung 0: A(左側) ST5 カメラ2 検査開始 *)
ST5_A_Ca2_M[1] := ((Auto_A_Start AND NOT ST5_A_Ca2_Busy) OR ST5_A_Ca2_M[1]) AND NOT ST5_A_Ca2_M[2];
(* Rung 1: A(左側) ST5 カメラ2 検査中 *)
ST5_A_Ca2_Busy := ((Auto_A_Start AND ST5_A_Ca2_M[1]) OR ST5_A_Ca2_Busy) AND NOT Ins_A_Next_Cycle;
(* Rung 2: A(左側) ST5 カメラ2 位置5ストッパー戻 *)
_p70 := ((ST5_A_Ca2_M[1] AND ST5_A_Ca2_Busy) OR ST5_A_Ca2_M[2]) AND NOT ST5_A_Ca2_M[4] AND NOT ST5_A_Ca2_M[5];
ST5_A_Ca2_M[2] := _p70;
Out_CYS_Pos_05_Stopper_A_H_Auto[2] := _p70;
(* Rung 3: A(左側) ST5 カメラ2 ワーク有無判定 *)
_e71(CLK := ST5_A_Ca2_M[2] AND NOT Pause[9]);
_p72 := ((ST5_A_Ca2_M[2] AND Out_CYS_Pos_05_Stopper_A_H_Done) OR _e71.Q OR ST5_A_Ca2_M[3]) AND NOT Pause[9] AND NOT ST5_A_Ca2_End;
ST5_A_Ca2_M[3] := _p72;
ST5_A_Ca2_M[4] := _p72 AND TimerQ_In_Sen_Work_A_Pos_05 AND (Station_A_Data[5].Work_On = TRUE);
ST5_A_Ca2_M[5] := _p72 AND NOT TimerQ_In_Sen_Work_A_Pos_05 AND (Station_A_Data[5].Work_On = FALSE);
IF _p72 AND ((TimerQ_In_Sen_Work_A_Pos_05 AND (Station_A_Data[5].Work_On = FALSE)) OR (NOT TimerQ_In_Sen_Work_A_Pos_05 AND (Station_A_Data[5].Work_On = TRUE))) THEN
    ST5_A_Ca2_M[6] := TRUE;
END_IF;
(* Rung 4: A(左側) ST5 カメラ2 測定開始 *)
_p73 := ((ST5_A_Ca2_M[3] AND ST5_A_Ca2_M[4] AND NOT Pause[9]) OR ST5_A_Ca2_M[7]) AND NOT Pause[9] AND NOT ST5_A_Ca2_End;
ST5_A_Ca2_M[7] := _p73;
FH_A_ST5_Auto := _p73;

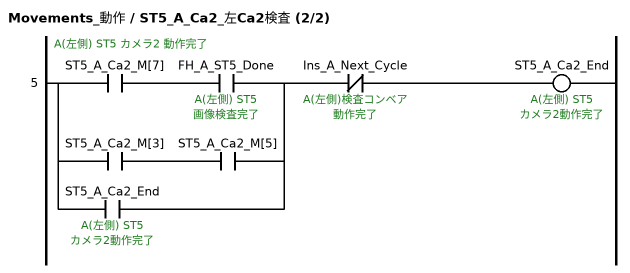
(* Rung 5: A(左側) ST5 カメラ2 動作完了 *)
ST5_A_Ca2_End := ((ST5_A_Ca2_M[7] AND FH_A_ST5_Done) OR (ST5_A_Ca2_M[3] AND ST5_A_Ca2_M[5]) OR ST5_A_Ca2_End) AND NOT Ins_A_Next_Cycle;

(* Section ST6_A_Rev2_左反転2: ladder, written here as Structured Text *)

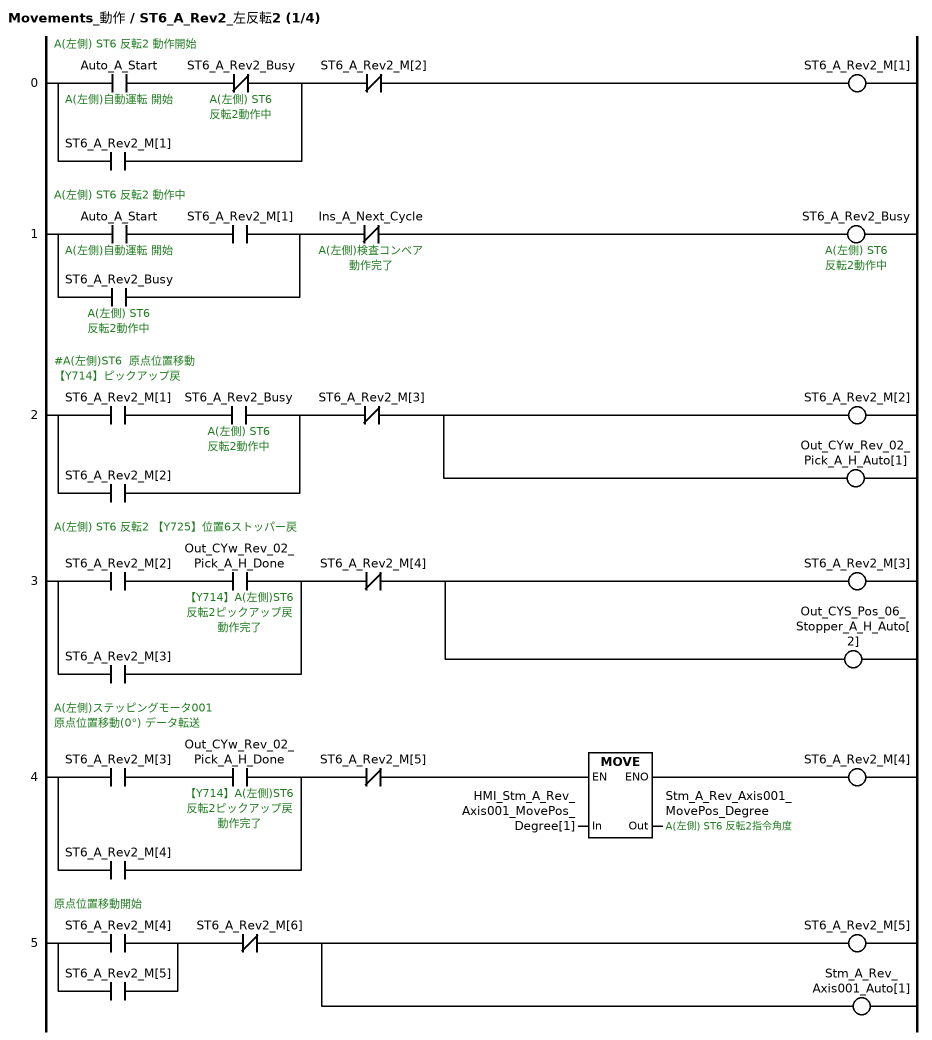
(* Rung 0: A(左側) ST6 反転2 動作開始 *)
ST6_A_Rev2_M[1] := ((Auto_A_Start AND NOT ST6_A_Rev2_Busy) OR ST6_A_Rev2_M[1]) AND NOT ST6_A_Rev2_M[2];
(* Rung 1: A(左側) ST6 反転2 動作中 *)
ST6_A_Rev2_Busy := ((Auto_A_Start AND ST6_A_Rev2_M[1]) OR ST6_A_Rev2_Busy) AND NOT Ins_A_Next_Cycle;
(* Rung 2: #A(左側)ST6  原点位置移動 / 【Y714】ピックアップ戻 *)
_p74 := ((ST6_A_Rev2_M[1] AND ST6_A_Rev2_Busy) OR ST6_A_Rev2_M[2]) AND NOT ST6_A_Rev2_M[3];
ST6_A_Rev2_M[2] := _p74;
Out_CYw_Rev_02_Pick_A_H_Auto[1] := _p74;
(* Rung 3: A(左側) ST6 反転2 【Y725】位置6ストッパー戻 *)
_p75 := ((ST6_A_Rev2_M[2] AND Out_CYw_Rev_02_Pick_A_H_Done) OR ST6_A_Rev2_M[3]) AND NOT ST6_A_Rev2_M[4];
ST6_A_Rev2_M[3] := _p75;
Out_CYS_Pos_06_Stopper_A_H_Auto[2] := _p75;
(* Rung 4: A(左側)ステッピングモータ001 / 原点位置移動(0°) データ転送 *)
IF ((ST6_A_Rev2_M[3] AND Out_CYw_Rev_02_Pick_A_H_Done) OR ST6_A_Rev2_M[4]) AND NOT ST6_A_Rev2_M[5] THEN
    Stm_A_Rev_Axis001_MovePos_Degree := HMI_Stm_A_Rev_Axis001_MovePos_Degree[1];
END_IF;
ST6_A_Rev2_M[4] := ((ST6_A_Rev2_M[3] AND Out_CYw_Rev_02_Pick_A_H_Done) OR ST6_A_Rev2_M[4]) AND NOT ST6_A_Rev2_M[5];
(* Rung 5: 原点位置移動開始 *)
_p76 := (ST6_A_Rev2_M[4] OR ST6_A_Rev2_M[5]) AND NOT ST6_A_Rev2_M[6];
ST6_A_Rev2_M[5] := _p76;
Stm_A_Rev_Axis001_Auto[1] := _p76;

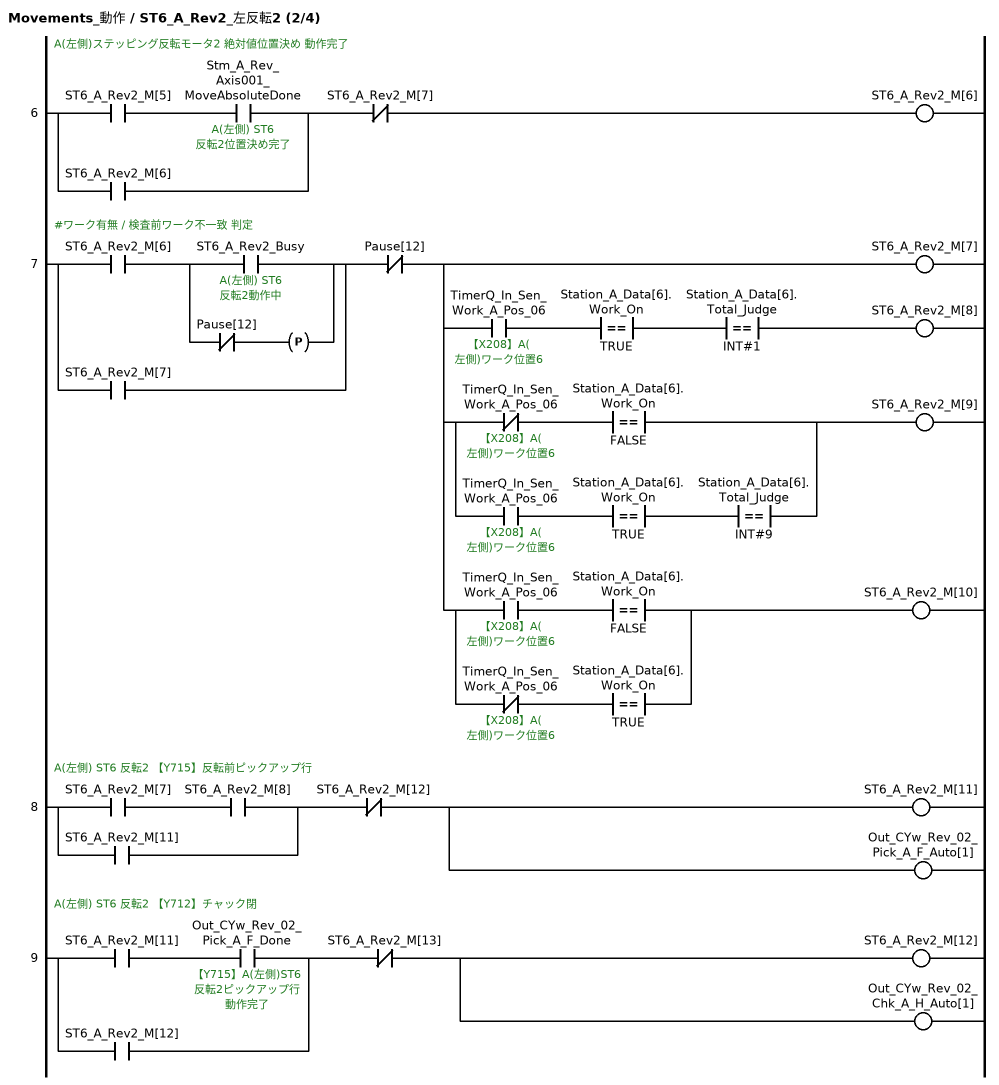
(* Rung 6: A(左側)ステッピング反転モータ2 絶対値位置決め 動作完了 *)
ST6_A_Rev2_M[6] := ((ST6_A_Rev2_M[5] AND Stm_A_Rev_Axis001_MoveAbsoluteDone) OR ST6_A_Rev2_M[6]) AND NOT ST6_A_Rev2_M[7];
(* Rung 7: #ワーク有無 / 検査前ワーク不一致 判定 *)
_e77(CLK := ST6_A_Rev2_M[6] AND NOT Pause[12]);
_p78 := ((ST6_A_Rev2_M[6] AND ST6_A_Rev2_Busy) OR _e77.Q OR ST6_A_Rev2_M[7]) AND NOT Pause[12];
ST6_A_Rev2_M[7] := _p78;
ST6_A_Rev2_M[8] := _p78 AND TimerQ_In_Sen_Work_A_Pos_06 AND (Station_A_Data[6].Work_On = TRUE) AND (Station_A_Data[6].Total_Judge = INT#1);
ST6_A_Rev2_M[9] := _p78 AND ((NOT TimerQ_In_Sen_Work_A_Pos_06 AND (Station_A_Data[6].Work_On = FALSE)) OR (TimerQ_In_Sen_Work_A_Pos_06 AND (Station_A_Data[6].Work_On = TRUE) AND (Station_A_Data[6].Total_Judge = INT#9)));
ST6_A_Rev2_M[10] := _p78 AND ((TimerQ_In_Sen_Work_A_Pos_06 AND (Station_A_Data[6].Work_On = FALSE)) OR (NOT TimerQ_In_Sen_Work_A_Pos_06 AND (Station_A_Data[6].Work_On = TRUE)));
(* Rung 8: A(左側) ST6 反転2 【Y715】反転前ピックアップ行 *)
_p79 := ((ST6_A_Rev2_M[7] AND ST6_A_Rev2_M[8]) OR ST6_A_Rev2_M[11]) AND NOT ST6_A_Rev2_M[12];
ST6_A_Rev2_M[11] := _p79;
Out_CYw_Rev_02_Pick_A_F_Auto[1] := _p79;
(* Rung 9: A(左側) ST6 反転2 【Y712】チャック閉 *)
_p80 := ((ST6_A_Rev2_M[11] AND Out_CYw_Rev_02_Pick_A_F_Done) OR ST6_A_Rev2_M[12]) AND NOT ST6_A_Rev2_M[13];
ST6_A_Rev2_M[12] := _p80;
Out_CYw_Rev_02_Chk_A_H_Auto[1] := _p80;

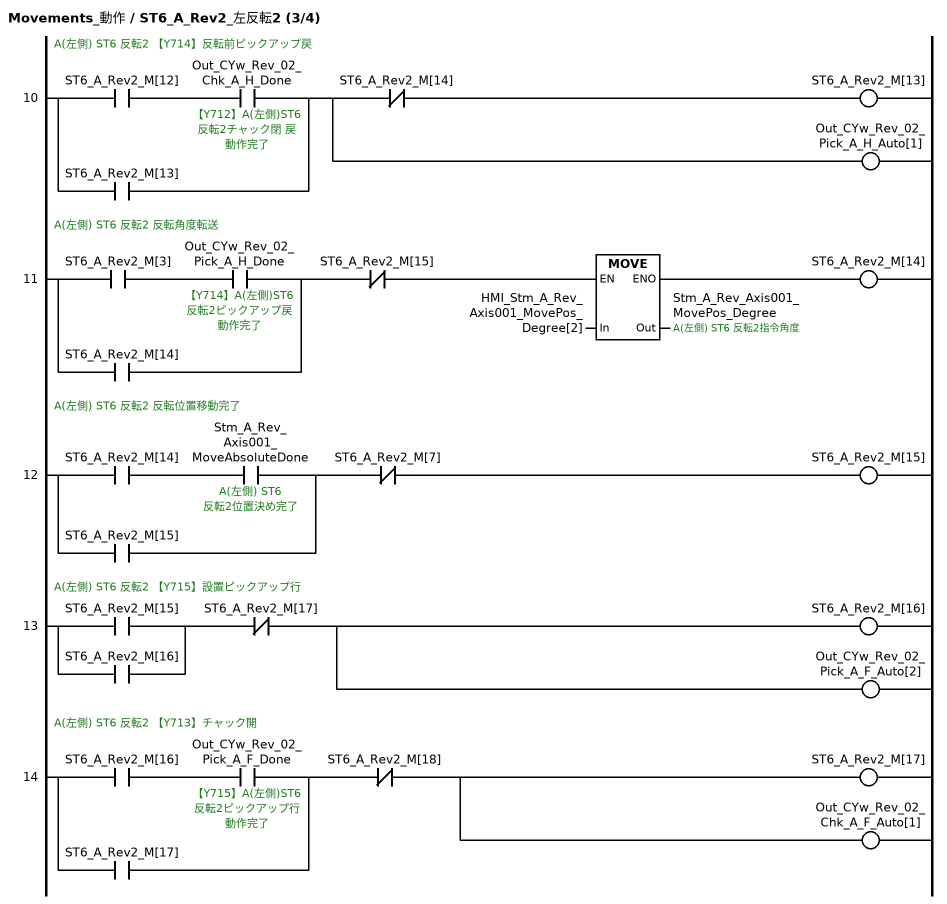
(* Rung 10: A(左側) ST6 反転2 【Y714】反転前ピックアップ戻 *)
_p81 := (ST6_A_Rev2_M[12] AND Out_CYw_Rev_02_Chk_A_H_Done) OR ST6_A_Rev2_M[13];
ST6_A_Rev2_M[13] := _p81 AND NOT ST6_A_Rev2_M[14];
Out_CYw_Rev_02_Pick_A_H_Auto[1] := _p81;
(* Rung 11: A(左側) ST6 反転2 反転角度転送 *)
IF ((ST6_A_Rev2_M[3] AND Out_CYw_Rev_02_Pick_A_H_Done) OR ST6_A_Rev2_M[14]) AND NOT ST6_A_Rev2_M[15] THEN
    Stm_A_Rev_Axis001_MovePos_Degree := HMI_Stm_A_Rev_Axis001_MovePos_Degree[2];
END_IF;
ST6_A_Rev2_M[14] := ((ST6_A_Rev2_M[3] AND Out_CYw_Rev_02_Pick_A_H_Done) OR ST6_A_Rev2_M[14]) AND NOT ST6_A_Rev2_M[15];
(* Rung 12: A(左側) ST6 反転2 反転位置移動完了 *)
ST6_A_Rev2_M[15] := ((ST6_A_Rev2_M[14] AND Stm_A_Rev_Axis001_MoveAbsoluteDone) OR ST6_A_Rev2_M[15]) AND NOT ST6_A_Rev2_M[7];
(* Rung 13: A(左側) ST6 反転2 【Y715】設置ピックアップ行 *)
_p82 := (ST6_A_Rev2_M[15] OR ST6_A_Rev2_M[16]) AND NOT ST6_A_Rev2_M[17];
ST6_A_Rev2_M[16] := _p82;
Out_CYw_Rev_02_Pick_A_F_Auto[2] := _p82;
(* Rung 14: A(左側) ST6 反転2 【Y713】チャック開 *)
_p83 := ((ST6_A_Rev2_M[16] AND Out_CYw_Rev_02_Pick_A_F_Done) OR ST6_A_Rev2_M[17]) AND NOT ST6_A_Rev2_M[18];
ST6_A_Rev2_M[17] := _p83;
Out_CYw_Rev_02_Chk_A_F_Auto[1] := _p83;

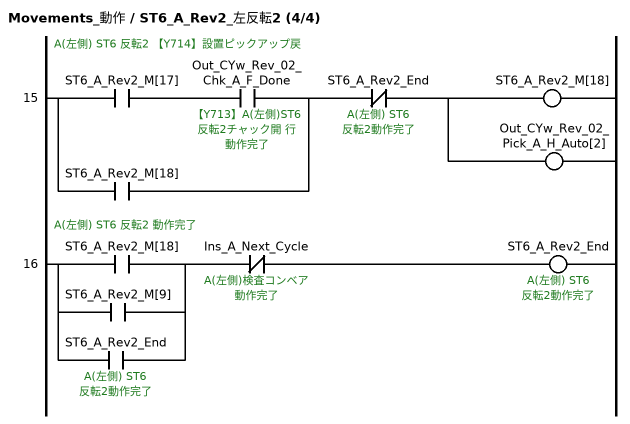
(* Rung 15: A(左側) ST6 反転2 【Y714】設置ピックアップ戻 *)
_p84 := ((ST6_A_Rev2_M[17] AND Out_CYw_Rev_02_Chk_A_F_Done) OR ST6_A_Rev2_M[18]) AND NOT ST6_A_Rev2_End;
ST6_A_Rev2_M[18] := _p84;
Out_CYw_Rev_02_Pick_A_H_Auto[2] := _p84;
(* Rung 16: A(左側) ST6 反転2 動作完了 *)
ST6_A_Rev2_End := (ST6_A_Rev2_M[18] OR ST6_A_Rev2_M[9] OR ST6_A_Rev2_End) AND NOT Ins_A_Next_Cycle;

(* Section ST7_A_Dis2_左SF排出: ladder, written here as Structured Text *)

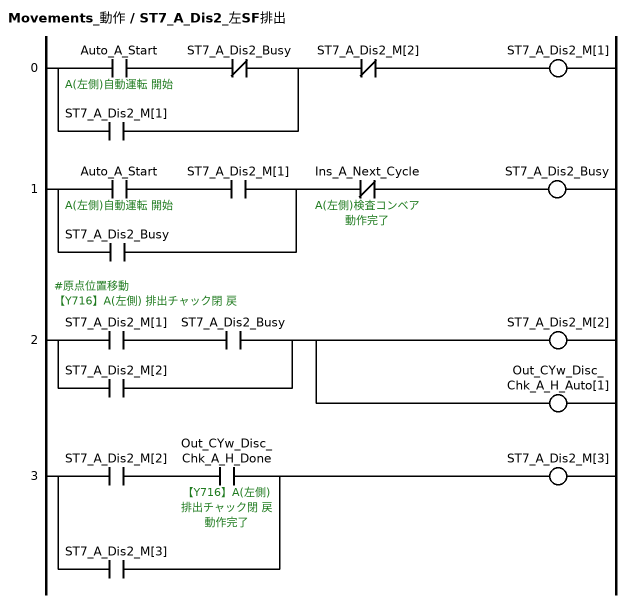
(* Rung 0 *)
ST7_A_Dis2_M[1] := ((Auto_A_Start AND NOT ST7_A_Dis2_Busy) OR ST7_A_Dis2_M[1]) AND NOT ST7_A_Dis2_M[2];
(* Rung 1 *)
ST7_A_Dis2_Busy := ((Auto_A_Start AND ST7_A_Dis2_M[1]) OR ST7_A_Dis2_Busy) AND NOT Ins_A_Next_Cycle;
(* Rung 2: #原点位置移動 / 【Y716】A(左側) 排出チャック閉 戻 *)
_p85 := (ST7_A_Dis2_M[1] AND ST7_A_Dis2_Busy) OR ST7_A_Dis2_M[2];
ST7_A_Dis2_M[2] := _p85;
Out_CYw_Disc_Chk_A_H_Auto[1] := _p85;
(* Rung 3 *)
ST7_A_Dis2_M[3] := (ST7_A_Dis2_M[2] AND Out_CYw_Disc_Chk_A_H_Done) OR ST7_A_Dis2_M[3];
END_PROGRAM

PROGRAM OtherDevice_外部機器
VAR
    FH_M : BOOL;
    GT2_M : BOOL;
    IAI_M : BOOL;  (* 旧ダミーマーカー（ST許可ではない） *)
    HMI_M : BOOL;
    FH_A_ST1_M : ARRAY[0..99] OF Bool;  (* [1] ST1 FH測定中; [5] ST1 測定完了 *)
    FH_A_ST1_OK : BOOL;  (* ST1 OK判定 *)
    FH_A_ST1_NG : BOOL;  (* ST1 NG 判定 *)
    FH_A_ST1_TON : ARRAY[0..99] OF TON;
    FH_A_ST1_TOF : ARRAY[0..99] OF TOF;
    ４ : UINT;
    ConvWordIndex : INT;  (* 作業用 ワード番号 *)
    ConvAxisIndex : INT;  (* 作業用 軸番号（RCON1:1～6／RCON2:1～5） *)
    ConvBase : INT;  (* 作業用 軸先頭ワード番号 *)
    ConvDWord : DWORD;  (* 作業用 32bit分割・結合 *)
    ConvPos : DINT;  (* 作業用 目標位置 [0.01mm・符号付き] *)
    ConvBand : UDINT;  (* 作業用 位置決め幅 [0.01mm] *)
    ConvSpeed : UINT;  (* 作業用 速度送信値 *)
    ConvAccDec : UINT;  (* 作業用 共通加減速 [0.01G] *)
    ConvPush : UINT;  (* 作業用 押付け制限 [255=100%] *)
    ConvScaled : LREAL;  (* 作業用 換算後の小数値 *)
    ConvWord : WORD;  (* 作業用 16bitワード *)
    ConvUnitOK : BOOL;  (* 作業用 速度単位正常 *)
    RCON1_1_TOF : ARRAY[0..99] OF TOF;  (* A(左側) RCON1_1 NG1上下降 開始要求100ms保持; [1] A(左側) RCON1_1 NG1上下降 開始要求100ms保持 *)
    RCON1_1_TON : ARRAY[0..99] OF TON;  (* A(左側) RCON1_1 NG1上下降 準備・完了タイマー; [1] A(左側) RCON1_1 NG1上下降準備100ms確認; [2] A(左側) RCON1_1 NG1上下降 動作完了100ms保持 *)
    Stm_A_Rev_Axis000_ZeroSet : MC_SetPosition;
    Stm_A_Rev_Axis000_HomeWithParameter : MC_HomeWithParameter;
    Stm_A_Rev_Axis000_Power : MC_Power;  (* A(左側)ステッピングモータ000 電源ON状態 *)
    Stm_A_Rev_Axis000_MoveAbsolute : MC_MoveAbsolute;
    Stm_A_Rev_Axis000_MoveVel : LREAL;  (* 動作速度 *)
    Stm_A_Rev_Axis000_MoveAcc : LREAL;  (* 動作加速度 *)
    Stm_A_Rev_Axis000_MoveDec : LREAL;  (* 動作減速度 *)
    Stm_A_Rev_Axis000_MoveBusy : BOOL;  (* 動作中 *)
    Stm_A_Rev_Axis000_MoveError : BOOL;  (* 動作エラー *)
    Stm_A_Rev_Axis000_TON : ARRAY[0..99] OF TON;
    FH_A_ST5_M : ARRAY[0..99] OF Bool;  (* A(左側) ST5 FH工程; [1] A(左側) ST5 測定要求; [2] A(左側) ST5 シーン切替; [3] A(左側) ST5 コマンド完了; [4] A(左側) ST5 測定トリガー; [5] A(左側) ST5 測定完了; [6] A(左側) ST5 OK保持; [7] A(左側) ST5 NG／完了保持 *)
    FH_A_ST5_OK : BOOL;  (* A(左側) ST5 OK判定 *)
    FH_A_ST5_NG : BOOL;  (* A(左側) ST5 NG判定 *)
    FH_A_ST5_TON : ARRAY[0..99] OF TON;  (* A(左側) ST5 FH遅延タイマー *)
    FH_A_ST5_TOF : ARRAY[0..99] OF TOF;  (* A(左側) ST5 FHトリガ保持; [1] A(左側) ST5 トリガー100ms *)
    Stm_A_Rev_Axis001_ZeroSet : MC_SetPosition;  (* A(左側) ST6 反転2 位置ゼロ設定 *)
    Stm_A_Rev_Axis001_HomeWithParameter : MC_HomeWithParameter;  (* A(左側) ST6 反転2 原点復帰FB *)
    Stm_A_Rev_Axis001_Power : MC_Power;  (* A(左側) ST6 反転2 電源ON状態 *)
    Stm_A_Rev_Axis001_MoveAbsolute : MC_MoveAbsolute;  (* A(左側) ST6 反転2 絶対位置決めFB *)
    Stm_A_Rev_Axis001_MoveVel : LREAL;  (* A(左側) ST6 反転2 速度 *)
    Stm_A_Rev_Axis001_MoveAcc : LREAL;  (* A(左側) ST6 反転2 加速度 *)
    Stm_A_Rev_Axis001_MoveDec : LREAL;  (* A(左側) ST6 反転2 減速度 *)
    Stm_A_Rev_Axis001_MoveBusy : BOOL;  (* A(左側) ST6 反転2 移動中 *)
    Stm_A_Rev_Axis001_MoveError : BOOL;  (* A(左側) ST6 反転2 移動エラー *)
    Stm_A_Rev_Axis001_TON : ARRAY[0..99] OF TON;  (* A(左側) ST6 反転2 完了保持タイマー *)
    RCON1_2_TOF : ARRAY[0..99] OF TOF;  (* B(右側) RCON1_2 NG1上下降 開始要求100ms保持; [1] B(右側) RCON1_2 NG1上下降 開始要求100ms保持 *)
    RCON1_2_TON : ARRAY[0..99] OF TON;  (* B(右側) RCON1_2 NG1上下降 準備・完了タイマー; [1] B(右側) RCON1_2 NG1上下降準備100ms確認; [2] B(右側) RCON1_2 NG1上下降 動作完了100ms保持 *)
    RCON1_3_TOF : ARRAY[0..99] OF TOF;  (* A(左側) RCON1_3 SF/NG2送り 開始要求100ms保持; [1] A(左側) RCON1_3 SF/NG2送り 開始要求100ms保持 *)
    RCON1_3_TON : ARRAY[0..99] OF TON;  (* A(左側) RCON1_3 SF/NG2送り 準備・完了タイマー; [1] A(左側) RCON1_3 SF/NG2送り準備100ms確認; [2] A(左側) RCON1_3 SF/NG2送り 動作完了100ms保持 *)
    RCON1_4_TOF : ARRAY[0..99] OF TOF;  (* B(右側) RCON1_4 SF/NG2送り 開始要求100ms保持; [1] B(右側) RCON1_4 SF/NG2送り 開始要求100ms保持 *)
    RCON1_4_TON : ARRAY[0..99] OF TON;  (* B(右側) RCON1_4 SF/NG2送り 準備・完了タイマー; [1] B(右側) RCON1_4 SF/NG2送り準備100ms確認; [2] B(右側) RCON1_4 SF/NG2送り 動作完了100ms保持 *)
    RCON1_5_TOF : ARRAY[0..99] OF TOF;  (* A(左側) RCON1_5 SF/NG2上下降 開始要求100ms保持; [1] A(左側) RCON1_5 SF/NG2上下降 開始要求100ms保持 *)
    RCON1_5_TON : ARRAY[0..99] OF TON;  (* A(左側) RCON1_5 SF/NG2上下降 準備・完了タイマー; [1] A(左側) RCON1_5 SF/NG2上下降準備100ms確認; [2] A(左側) RCON1_5 SF/NG2上下降 動作完了100ms保持 *)
    RCON1_6_TOF : ARRAY[0..99] OF TOF;  (* B(右側) RCON1_6 SF/NG2上下降 開始要求100ms保持; [1] B(右側) RCON1_6 SF/NG2上下降 開始要求100ms保持 *)
    RCON1_6_TON : ARRAY[0..99] OF TON;  (* B(右側) RCON1_6 SF/NG2上下降 準備・完了タイマー; [1] B(右側) RCON1_6 SF/NG2上下降準備100ms確認; [2] B(右側) RCON1_6 SF/NG2上下降 動作完了100ms保持 *)
END_VAR
VAR_EXTERNAL
    HMI_MessageNo : ARRAY[0..9] OF UINT;
    HMI_Message : ARRAY[0..9] OF String[256];
    HMI_Language : BOOL;
    FH_Line0_Trigger_Ready_1 : BOOL;
    FH_Line0_Trigger_1 : BOOL;
    M9999 : BOOL;
    FH_Line0_Busy_1 : BOOL;
    FH_Line0_Result_Notification_1 : BOOL;
    FH_Line0_DINT_Result_Data_0_1 : DINT;
    FH_Line0_DINT_Result_Data_1_1 : DINT;
    FH_Line0_DINT_Result_Data_2_1 : DINT;
    FH_Line0_Command_Code_1 : DWORD;
    FH_Line0_Command_Request_1 : BOOL;
    FH_Line0_Command_Completion_1 : BOOL;
    MdlChg : BOOL;  (* 機種切替：ON【GA120】 OFF【GA90】 *)
    FH_Line0_Error_Status_1 : BOOL;
    FH_5552_10_A_Auto : BOOL;  (* ST1 FH測定開始 *)
    FH_A_ST1_Manual : BOOL;  (* ST1 *)
    Pause : ARRAY[0..99] OF Bool;  (* [3] FH A(左側) ST1; [9] FH A(左側) ST5; [10] FH B(右側) ST1; [11] FH B(右側) ST5; [12] A(左側) ST6 反転2 ワーク不一致 *)
    FH_A_ST1_Done : BOOL;  (* ST1 画像検査完了 *)
    Station_A_Data : ARRAY[0..8] OF sData;
    DLEP1_OUT : ARRAY[0..79] OF BOOL;
    DLEP2_OUT : ARRAY[0..79] OF BOOL;
    DLEP1_IN : ARRAY[0..167] OF byte;
    DLEP2_IN : ARRAY[0..167] OF byte;
    DLEP2_IN_Error : BOOL;  (* B(右側)センサエラー *)
    DLEP1_IN_Error : BOOL;  (* A(右側)センサエラー *)
    GT2_A_CurrentVal : INT;  (* A(左側) 測定値 *)
    GT2_B_CurrentVal : INT;  (* B(右側) 測定値 *)
    Hgt_A_Ins_Data : LREAL;  (* A測定データに変換 *)
    Hgt_B_Ins_Data : LREAL;
    Hgt_A_ComputedValueData : LREAL;  (* A測定データ+13.000mm 算定データ *)
    Hgt_B_ComputedValueData : LREAL;  (* B測定データ+13.000mm 算定データ *)
    E001_In_IN00_2004_01 : UINT;  (* RCON1 IN00 GW状態 *)
    E001_In_IN01_2004_02 : UINT;  (* RCON1 IN01 軸リンク状態 *)
    E001_In_IN02_2004_03 : UINT;  (* RCON1 IN02 電源状態0 *)
    E001_In_IN03_2004_04 : UINT;  (* RCON1 IN03 電源状態1 *)
    E001_In_IN04_2004_05 : UINT;  (* RCON1 IN04 電源状態2 *)
    E001_In_IN05_2004_06 : UINT;  (* RCON1 IN05 電源状態3 *)
    E001_In_IN06_2004_07 : UINT;  (* RCON1 IN06 電源状態4（構成依存） *)
    E001_In_IN07_2004_08 : UINT;  (* RCON1 IN07 予約（使用禁止） *)
    E001_In_IN08_2004_09 : UINT;  (* A(左側) RCON1_1 NG1上下降 IN08 現在位置 下位 [0.01mm] *)
    E001_In_IN09_2004_0A : UINT;  (* A(左側) RCON1_1 NG1上下降 IN09 現在位置 上位 [0.01mm] *)
    E001_In_IN10_2004_0B : UINT;  (* A(左側) RCON1_1 NG1上下降 IN10 指令電流 下位 [mA] *)
    E001_In_IN11_2004_0C : UINT;  (* A(左側) RCON1_1 NG1上下降 IN11 指令電流 上位 [mA] *)
    E001_In_IN12_2004_0D : UINT;  (* A(左側) RCON1_1 NG1上下降 IN12 現在速度 [実機単位・符号付き] *)
    E001_In_IN13_2004_0E : UINT;  (* A(左側) RCON1_1 NG1上下降 IN13 予約（使用禁止） *)
    E001_In_IN14_2004_0F : UINT;  (* A(左側) RCON1_1 NG1上下降 IN14 軸異常コード *)
    E001_In_IN15_2004_10 : UINT;  (* A(左側) RCON1_1 NG1上下降 IN15 状態信号（PEND/SV等） *)
    E001_In_IN16_2004_11 : UINT;  (* B(右側) RCON1_2 NG1上下降 IN16 現在位置 下位 [0.01mm] *)
    E001_In_IN17_2004_12 : UINT;  (* B(右側) RCON1_2 NG1上下降 IN17 現在位置 上位 [0.01mm] *)
    E001_In_IN18_2004_13 : UINT;  (* B(右側) RCON1_2 NG1上下降 IN18 指令電流 下位 [mA] *)
    E001_In_IN19_2004_14 : UINT;  (* B(右側) RCON1_2 NG1上下降 IN19 指令電流 上位 [mA] *)
    E001_In_IN20_2004_15 : UINT;  (* B(右側) RCON1_2 NG1上下降 IN20 現在速度 [実機単位・符号付き] *)
    E001_In_IN21_2004_16 : UINT;  (* B(右側) RCON1_2 NG1上下降 IN21 予約（使用禁止） *)
    E001_In_IN22_2004_17 : UINT;  (* B(右側) RCON1_2 NG1上下降 IN22 軸異常コード *)
    E001_In_IN23_2004_18 : UINT;  (* B(右側) RCON1_2 NG1上下降 IN23 状態信号（PEND/SV等） *)
    E001_In_IN24_2004_19 : UINT;  (* A(左側) RCON1_3 SF/NG2送り IN24 現在位置 下位 [0.01mm] *)
    E001_In_IN25_2004_1A : UINT;  (* A(左側) RCON1_3 SF/NG2送り IN25 現在位置 上位 [0.01mm] *)
    E001_In_IN26_2004_1B : UINT;  (* A(左側) RCON1_3 SF/NG2送り IN26 指令電流 下位 [mA] *)
    E001_In_IN27_2004_1C : UINT;  (* A(左側) RCON1_3 SF/NG2送り IN27 指令電流 上位 [mA] *)
    E001_In_IN28_2004_1D : UINT;  (* A(左側) RCON1_3 SF/NG2送り IN28 現在速度 [実機単位・符号付き] *)
    E001_In_IN29_2004_1E : UINT;  (* A(左側) RCON1_3 SF/NG2送り IN29 予約（使用禁止） *)
    E001_In_IN30_2004_1F : UINT;  (* A(左側) RCON1_3 SF/NG2送り IN30 軸異常コード *)
    E001_In_IN31_2004_20 : UINT;  (* A(左側) RCON1_3 SF/NG2送り IN31 状態信号（PEND/SV等） *)
    E001_In_IN32_2004_21 : UINT;  (* B(右側) RCON1_4 SF/NG2送り IN32 現在位置 下位 [0.01mm] *)
    E001_In_IN33_2004_22 : UINT;  (* B(右側) RCON1_4 SF/NG2送り IN33 現在位置 上位 [0.01mm] *)
    E001_In_IN34_2004_23 : UINT;  (* B(右側) RCON1_4 SF/NG2送り IN34 指令電流 下位 [mA] *)
    E001_In_IN35_2004_24 : UINT;  (* B(右側) RCON1_4 SF/NG2送り IN35 指令電流 上位 [mA] *)
    E001_In_IN36_2004_25 : UINT;  (* B(右側) RCON1_4 SF/NG2送り IN36 現在速度 [実機単位・符号付き] *)
    E001_In_IN37_2004_26 : UINT;  (* B(右側) RCON1_4 SF/NG2送り IN37 予約（使用禁止） *)
    E001_In_IN38_2004_27 : UINT;  (* B(右側) RCON1_4 SF/NG2送り IN38 軸異常コード *)
    E001_In_IN39_2004_28 : UINT;  (* B(右側) RCON1_4 SF/NG2送り IN39 状態信号（PEND/SV等） *)
    E001_In_IN40_2004_29 : UINT;  (* A(左側) RCON1_5 SF/NG2上下降 IN40 現在位置 下位 [0.01mm] *)
    E001_In_IN41_2004_2A : UINT;  (* A(左側) RCON1_5 SF/NG2上下降 IN41 現在位置 上位 [0.01mm] *)
    E001_In_IN42_2004_2B : UINT;  (* A(左側) RCON1_5 SF/NG2上下降 IN42 指令電流 下位 [mA] *)
    E001_In_IN43_2004_2C : UINT;  (* A(左側) RCON1_5 SF/NG2上下降 IN43 指令電流 上位 [mA] *)
    E001_In_IN44_2004_2D : UINT;  (* A(左側) RCON1_5 SF/NG2上下降 IN44 現在速度 [実機単位・符号付き] *)
    E001_In_IN45_2004_2E : UINT;  (* A(左側) RCON1_5 SF/NG2上下降 IN45 予約（使用禁止） *)
    E001_In_IN46_2004_2F : UINT;  (* A(左側) RCON1_5 SF/NG2上下降 IN46 軸異常コード *)
    E001_In_IN47_2004_30 : UINT;  (* A(左側) RCON1_5 SF/NG2上下降 IN47 状態信号（PEND/SV等） *)
    E001_In_IN48_2004_31 : UINT;  (* B(右側) RCON1_6 SF/NG2上下降 IN48 現在位置 下位 [0.01mm] *)
    E001_In_IN49_2004_32 : UINT;  (* B(右側) RCON1_6 SF/NG2上下降 IN49 現在位置 上位 [0.01mm] *)
    E001_In_IN50_2004_33 : UINT;  (* B(右側) RCON1_6 SF/NG2上下降 IN50 指令電流 下位 [mA] *)
    E001_In_IN51_2004_34 : UINT;  (* B(右側) RCON1_6 SF/NG2上下降 IN51 指令電流 上位 [mA] *)
    E001_In_IN52_2004_35 : UINT;  (* B(右側) RCON1_6 SF/NG2上下降 IN52 現在速度 [実機単位・符号付き] *)
    E001_In_IN53_2004_36 : UINT;  (* B(右側) RCON1_6 SF/NG2上下降 IN53 予約（使用禁止） *)
    E001_In_IN54_2004_37 : UINT;  (* B(右側) RCON1_6 SF/NG2上下降 IN54 軸異常コード *)
    E001_In_IN55_2004_38 : UINT;  (* B(右側) RCON1_6 SF/NG2上下降 IN55 状態信号（PEND/SV等） *)
    E001_In_IN56_2004_39 : UINT;  (* RCON1 IN56 112Byte範囲外（未割付・不使用） *)
    E001_In_IN57_2004_3A : UINT;  (* RCON1 IN57 112Byte範囲外（未割付・不使用） *)
    E001_In_IN58_2004_3B : UINT;  (* RCON1 IN58 112Byte範囲外（未割付・不使用） *)
    E001_In_IN59_2004_3C : UINT;  (* RCON1 IN59 112Byte範囲外（未割付・不使用） *)
    E001_In_IN60_2004_3D : UINT;  (* RCON1 IN60 112Byte範囲外（未割付・不使用） *)
    E001_In_IN61_2004_3E : UINT;  (* RCON1 IN61 112Byte範囲外（未割付・不使用） *)
    E001_In_IN62_2004_3F : UINT;  (* RCON1 IN62 112Byte範囲外（未割付・不使用） *)
    E001_In_IN63_2004_40 : UINT;  (* RCON1 IN63 112Byte範囲外（未割付・不使用） *)
    E001_In_IN64_2004_41 : UINT;  (* RCON1 IN64 112Byte範囲外（未割付・不使用） *)
    E001_In_IN65_2004_42 : UINT;  (* RCON1 IN65 112Byte範囲外（未割付・不使用） *)
    E001_In_IN66_2004_43 : UINT;  (* RCON1 IN66 112Byte範囲外（未割付・不使用） *)
    E001_In_IN67_2004_44 : UINT;  (* RCON1 IN67 112Byte範囲外（未割付・不使用） *)
    E001_In_IN68_2004_45 : UINT;  (* RCON1 IN68 112Byte範囲外（未割付・不使用） *)
    E001_In_IN69_2004_46 : UINT;  (* RCON1 IN69 112Byte範囲外（未割付・不使用） *)
    E001_In_IN70_2004_47 : UINT;  (* RCON1 IN70 112Byte範囲外（未割付・不使用） *)
    E001_In_IN71_2004_48 : UINT;  (* RCON1 IN71 112Byte範囲外（未割付・不使用） *)
    E001_Out_OUT00_2003_01 : UINT;  (* RCON1 OUT00 共通制御（MON/RTE） *)
    E001_Out_OUT08_2003_09 : UINT;  (* A(左側) RCON1_1 NG1上下降 OUT08 目標位置 下位 [0.01mm] *)
    E001_Out_OUT09_2003_0A : UINT;  (* A(左側) RCON1_1 NG1上下降 OUT09 目標位置 上位 [0.01mm] *)
    E001_Out_OUT10_2003_0B : UINT;  (* A(左側) RCON1_1 NG1上下降 OUT10 位置決め幅 下位 [0.01mm] *)
    E001_Out_OUT11_2003_0C : UINT;  (* A(左側) RCON1_1 NG1上下降 OUT11 位置決め幅 上位 [0.01mm] *)
    E001_Out_OUT12_2003_0D : UINT;  (* A(左側) RCON1_1 NG1上下降 OUT12 速度指令 [実機単位] *)
    E001_Out_OUT13_2003_0E : UINT;  (* A(左側) RCON1_1 NG1上下降 OUT13 共通加減速 [0.01G] *)
    E001_Out_OUT14_2003_0F : UINT;  (* A(左側) RCON1_1 NG1上下降 OUT14 押付け制限 [255=100%] *)
    E001_Out_OUT15_2003_10 : UINT;  (* A(左側) RCON1_1 NG1上下降 OUT15 制御信号（DSTR/SON等） *)
    E001_Out_OUT16_2003_11 : UINT;  (* B(右側) RCON1_2 NG1上下降 OUT16 目標位置 下位 [0.01mm] *)
    E001_Out_OUT17_2003_12 : UINT;  (* B(右側) RCON1_2 NG1上下降 OUT17 目標位置 上位 [0.01mm] *)
    E001_Out_OUT18_2003_13 : UINT;  (* B(右側) RCON1_2 NG1上下降 OUT18 位置決め幅 下位 [0.01mm] *)
    E001_Out_OUT19_2003_14 : UINT;  (* B(右側) RCON1_2 NG1上下降 OUT19 位置決め幅 上位 [0.01mm] *)
    E001_Out_OUT20_2003_15 : UINT;  (* B(右側) RCON1_2 NG1上下降 OUT20 速度指令 [実機単位] *)
    E001_Out_OUT21_2003_16 : UINT;  (* B(右側) RCON1_2 NG1上下降 OUT21 共通加減速 [0.01G] *)
    E001_Out_OUT22_2003_17 : UINT;  (* B(右側) RCON1_2 NG1上下降 OUT22 押付け制限 [255=100%] *)
    E001_Out_OUT23_2003_18 : UINT;  (* B(右側) RCON1_2 NG1上下降 OUT23 制御信号（DSTR/SON等） *)
    E001_Out_OUT24_2003_19 : UINT;  (* A(左側) RCON1_3 SF/NG2送り OUT24 目標位置 下位 [0.01mm] *)
    E001_Out_OUT25_2003_1A : UINT;  (* A(左側) RCON1_3 SF/NG2送り OUT25 目標位置 上位 [0.01mm] *)
    E001_Out_OUT26_2003_1B : UINT;  (* A(左側) RCON1_3 SF/NG2送り OUT26 位置決め幅 下位 [0.01mm] *)
    E001_Out_OUT27_2003_1C : UINT;  (* A(左側) RCON1_3 SF/NG2送り OUT27 位置決め幅 上位 [0.01mm] *)
    E001_Out_OUT28_2003_1D : UINT;  (* A(左側) RCON1_3 SF/NG2送り OUT28 速度指令 [実機単位] *)
    E001_Out_OUT29_2003_1E : UINT;  (* A(左側) RCON1_3 SF/NG2送り OUT29 共通加減速 [0.01G] *)
    E001_Out_OUT30_2003_1F : UINT;  (* A(左側) RCON1_3 SF/NG2送り OUT30 押付け制限 [255=100%] *)
    E001_Out_OUT31_2003_20 : UINT;  (* A(左側) RCON1_3 SF/NG2送り OUT31 制御信号（DSTR/SON等） *)
    E001_Out_OUT32_2003_21 : UINT;  (* B(右側) RCON1_4 SF/NG2送り OUT32 目標位置 下位 [0.01mm] *)
    E001_Out_OUT33_2003_22 : UINT;  (* B(右側) RCON1_4 SF/NG2送り OUT33 目標位置 上位 [0.01mm] *)
    E001_Out_OUT34_2003_23 : UINT;  (* B(右側) RCON1_4 SF/NG2送り OUT34 位置決め幅 下位 [0.01mm] *)
    E001_Out_OUT35_2003_24 : UINT;  (* B(右側) RCON1_4 SF/NG2送り OUT35 位置決め幅 上位 [0.01mm] *)
    E001_Out_OUT36_2003_25 : UINT;  (* B(右側) RCON1_4 SF/NG2送り OUT36 速度指令 [実機単位] *)
    E001_Out_OUT37_2003_26 : UINT;  (* B(右側) RCON1_4 SF/NG2送り OUT37 共通加減速 [0.01G] *)
    E001_Out_OUT38_2003_27 : UINT;  (* B(右側) RCON1_4 SF/NG2送り OUT38 押付け制限 [255=100%] *)
    E001_Out_OUT39_2003_28 : UINT;  (* B(右側) RCON1_4 SF/NG2送り OUT39 制御信号（DSTR/SON等） *)
    E001_Out_OUT40_2003_29 : UINT;  (* A(左側) RCON1_5 SF/NG2上下降 OUT40 目標位置 下位 [0.01mm] *)
    E001_Out_OUT41_2003_2A : UINT;  (* A(左側) RCON1_5 SF/NG2上下降 OUT41 目標位置 上位 [0.01mm] *)
    E001_Out_OUT42_2003_2B : UINT;  (* A(左側) RCON1_5 SF/NG2上下降 OUT42 位置決め幅 下位 [0.01mm] *)
    E001_Out_OUT43_2003_2C : UINT;  (* A(左側) RCON1_5 SF/NG2上下降 OUT43 位置決め幅 上位 [0.01mm] *)
    E001_Out_OUT44_2003_2D : UINT;  (* A(左側) RCON1_5 SF/NG2上下降 OUT44 速度指令 [実機単位] *)
    E001_Out_OUT45_2003_2E : UINT;  (* A(左側) RCON1_5 SF/NG2上下降 OUT45 共通加減速 [0.01G] *)
    E001_Out_OUT46_2003_2F : UINT;  (* A(左側) RCON1_5 SF/NG2上下降 OUT46 押付け制限 [255=100%] *)
    E001_Out_OUT47_2003_30 : UINT;  (* A(左側) RCON1_5 SF/NG2上下降 OUT47 制御信号（DSTR/SON等） *)
    E001_Out_OUT48_2003_31 : UINT;  (* B(右側) RCON1_6 SF/NG2上下降 OUT48 目標位置 下位 [0.01mm] *)
    E001_Out_OUT49_2003_32 : UINT;  (* B(右側) RCON1_6 SF/NG2上下降 OUT49 目標位置 上位 [0.01mm] *)
    E001_Out_OUT50_2003_33 : UINT;  (* B(右側) RCON1_6 SF/NG2上下降 OUT50 位置決め幅 下位 [0.01mm] *)
    E001_Out_OUT51_2003_34 : UINT;  (* B(右側) RCON1_6 SF/NG2上下降 OUT51 位置決め幅 上位 [0.01mm] *)
    E001_Out_OUT52_2003_35 : UINT;  (* B(右側) RCON1_6 SF/NG2上下降 OUT52 速度指令 [実機単位] *)
    E001_Out_OUT53_2003_36 : UINT;  (* B(右側) RCON1_6 SF/NG2上下降 OUT53 共通加減速 [0.01G] *)
    E001_Out_OUT54_2003_37 : UINT;  (* B(右側) RCON1_6 SF/NG2上下降 OUT54 押付け制限 [255=100%] *)
    E001_Out_OUT55_2003_38 : UINT;  (* B(右側) RCON1_6 SF/NG2上下降 OUT55 制御信号（DSTR/SON等） *)
    E005_In_IN00_2004_01_1 : UINT;  (* RCON2 IN00 GW状態 *)
    E005_In_IN01_2004_02_1 : UINT;  (* RCON2 IN01 軸リンク状態 *)
    E005_In_IN02_2004_03_1 : UINT;  (* RCON2 IN02 電源状態0 *)
    E005_In_IN03_2004_04_1 : UINT;  (* RCON2 IN03 電源状態1 *)
    E005_In_IN04_2004_05_1 : UINT;  (* RCON2 IN04 電源状態2 *)
    E005_In_IN05_2004_06_1 : UINT;  (* RCON2 IN05 電源状態3 *)
    E005_In_IN06_2004_07_1 : UINT;  (* RCON2 IN06 電源状態4（構成依存） *)
    E005_In_IN07_2004_08_1 : UINT;  (* RCON2 IN07 予約（使用禁止） *)
    E005_In_IN08_2004_09_1 : UINT;  (* RCON2 IN08 1軸目 現在位置 下位 [0.01mm] *)
    E005_In_IN09_2004_0A_1 : UINT;  (* RCON2 IN09 1軸目 現在位置 上位 [0.01mm] *)
    E005_In_IN10_2004_0B_1 : UINT;  (* RCON2 IN10 1軸目 指令電流 下位 [mA] *)
    E005_In_IN11_2004_0C_1 : UINT;  (* RCON2 IN11 1軸目 指令電流 上位 [mA] *)
    E005_In_IN12_2004_0D_1 : UINT;  (* RCON2 IN12 1軸目 現在速度 [実機単位・符号付き] *)
    E005_In_IN13_2004_0E_1 : UINT;  (* RCON2 IN13 1軸目 予約（使用禁止） *)
    E005_In_IN14_2004_0F_1 : UINT;  (* RCON2 IN14 1軸目 軸異常コード *)
    E005_In_IN15_2004_10_1 : UINT;  (* RCON2 IN15 1軸目 状態信号（PEND/SV等） *)
    E005_In_IN16_2004_11_1 : UINT;  (* RCON2 IN16 2軸目 現在位置 下位 [0.01mm] *)
    E005_In_IN17_2004_12_1 : UINT;  (* RCON2 IN17 2軸目 現在位置 上位 [0.01mm] *)
    E005_In_IN18_2004_13_1 : UINT;  (* RCON2 IN18 2軸目 指令電流 下位 [mA] *)
    E005_In_IN19_2004_14_1 : UINT;  (* RCON2 IN19 2軸目 指令電流 上位 [mA] *)
    E005_In_IN20_2004_15_1 : UINT;  (* RCON2 IN20 2軸目 現在速度 [実機単位・符号付き] *)
    E005_In_IN21_2004_16_1 : UINT;  (* RCON2 IN21 2軸目 予約（使用禁止） *)
    E005_In_IN22_2004_17_1 : UINT;  (* RCON2 IN22 2軸目 軸異常コード *)
    E005_In_IN23_2004_18_1 : UINT;  (* RCON2 IN23 2軸目 状態信号（PEND/SV等） *)
    E005_In_IN24_2004_19_1 : UINT;  (* RCON2 IN24 3軸目 現在位置 下位 [0.01mm] *)
    E005_In_IN25_2004_1A_1 : UINT;  (* RCON2 IN25 3軸目 現在位置 上位 [0.01mm] *)
    E005_In_IN26_2004_1B_1 : UINT;  (* RCON2 IN26 3軸目 指令電流 下位 [mA] *)
    E005_In_IN27_2004_1C_1 : UINT;  (* RCON2 IN27 3軸目 指令電流 上位 [mA] *)
    E005_In_IN28_2004_1D_1 : UINT;  (* RCON2 IN28 3軸目 現在速度 [実機単位・符号付き] *)
    E005_In_IN29_2004_1E_1 : UINT;  (* RCON2 IN29 3軸目 予約（使用禁止） *)
    E005_In_IN30_2004_1F_1 : UINT;  (* RCON2 IN30 3軸目 軸異常コード *)
    E005_In_IN31_2004_20_1 : UINT;  (* RCON2 IN31 3軸目 状態信号（PEND/SV等） *)
    E005_In_IN32_2004_21_1 : UINT;  (* RCON2 IN32 4軸目 現在位置 下位 [0.01mm] *)
    E005_In_IN33_2004_22_1 : UINT;  (* RCON2 IN33 4軸目 現在位置 上位 [0.01mm] *)
    E005_In_IN34_2004_23_1 : UINT;  (* RCON2 IN34 4軸目 指令電流 下位 [mA] *)
    E005_In_IN35_2004_24_1 : UINT;  (* RCON2 IN35 4軸目 指令電流 上位 [mA] *)
    E005_In_IN36_2004_25_1 : UINT;  (* RCON2 IN36 4軸目 現在速度 [実機単位・符号付き] *)
    E005_In_IN37_2004_26_1 : UINT;  (* RCON2 IN37 4軸目 予約（使用禁止） *)
    E005_In_IN38_2004_27_1 : UINT;  (* RCON2 IN38 4軸目 軸異常コード *)
    E005_In_IN39_2004_28_1 : UINT;  (* RCON2 IN39 4軸目 状態信号（PEND/SV等） *)
    E005_In_IN40_2004_29_1 : UINT;  (* RCON2 IN40 5軸目 現在位置 下位 [0.01mm] *)
    E005_In_IN41_2004_2A_1 : UINT;  (* RCON2 IN41 5軸目 現在位置 上位 [0.01mm] *)
    E005_In_IN42_2004_2B_1 : UINT;  (* RCON2 IN42 5軸目 指令電流 下位 [mA] *)
    E005_In_IN43_2004_2C_1 : UINT;  (* RCON2 IN43 5軸目 指令電流 上位 [mA] *)
    E005_In_IN44_2004_2D_1 : UINT;  (* RCON2 IN44 5軸目 現在速度 [実機単位・符号付き] *)
    E005_In_IN45_2004_2E_1 : UINT;  (* RCON2 IN45 5軸目 予約（使用禁止） *)
    E005_In_IN46_2004_2F_1 : UINT;  (* RCON2 IN46 5軸目 軸異常コード *)
    E005_In_IN47_2004_30_1 : UINT;  (* RCON2 IN47 5軸目 状態信号（PEND/SV等） *)
    E005_In_IN48_2004_31_1 : UINT;  (* RCON2 IN48 用途未確認（今回未使用） *)
    E005_In_IN49_2004_32_1 : UINT;  (* RCON2 IN49 用途未確認（今回未使用） *)
    E005_In_IN50_2004_33_1 : UINT;  (* RCON2 IN50 用途未確認（今回未使用） *)
    E005_In_IN51_2004_34_1 : UINT;  (* RCON2 IN51 用途未確認（今回未使用） *)
    E005_In_IN52_2004_35_1 : UINT;  (* RCON2 IN52 用途未確認（今回未使用） *)
    E005_In_IN53_2004_36_1 : UINT;  (* RCON2 IN53 用途未確認（今回未使用） *)
    E005_In_IN54_2004_37_1 : UINT;  (* RCON2 IN54 用途未確認（今回未使用） *)
    E005_In_IN55_2004_38_1 : UINT;  (* RCON2 IN55 用途未確認（今回未使用） *)
    E005_Out_OUT00_2003_01_1 : UINT;  (* RCON2 OUT00 共通制御（MON/RTE） *)
    E005_Out_OUT08_2003_09_1 : UINT;  (* RCON2 OUT08 1軸目 目標位置 下位 [0.01mm] *)
    E005_Out_OUT09_2003_0A_1 : UINT;  (* RCON2 OUT09 1軸目 目標位置 上位 [0.01mm] *)
    E005_Out_OUT10_2003_0B_1 : UINT;  (* RCON2 OUT10 1軸目 位置決め幅 下位 [0.01mm] *)
    E005_Out_OUT11_2003_0C_1 : UINT;  (* RCON2 OUT11 1軸目 位置決め幅 上位 [0.01mm] *)
    E005_Out_OUT12_2003_0D_1 : UINT;  (* RCON2 OUT12 1軸目 速度指令 [実機単位] *)
    E005_Out_OUT13_2003_0E_1 : UINT;  (* RCON2 OUT13 1軸目 共通加減速 [0.01G] *)
    E005_Out_OUT14_2003_0F_1 : UINT;  (* RCON2 OUT14 1軸目 押付け制限 [255=100%] *)
    E005_Out_OUT15_2003_10_1 : UINT;  (* RCON2 OUT15 1軸目 制御信号（DSTR/SON等） *)
    E005_Out_OUT16_2003_11_1 : UINT;  (* RCON2 OUT16 2軸目 目標位置 下位 [0.01mm] *)
    E005_Out_OUT17_2003_12_1 : UINT;  (* RCON2 OUT17 2軸目 目標位置 上位 [0.01mm] *)
    E005_Out_OUT18_2003_13_1 : UINT;  (* RCON2 OUT18 2軸目 位置決め幅 下位 [0.01mm] *)
    E005_Out_OUT19_2003_14_1 : UINT;  (* RCON2 OUT19 2軸目 位置決め幅 上位 [0.01mm] *)
    E005_Out_OUT20_2003_15_1 : UINT;  (* RCON2 OUT20 2軸目 速度指令 [実機単位] *)
    E005_Out_OUT21_2003_16_1 : UINT;  (* RCON2 OUT21 2軸目 共通加減速 [0.01G] *)
    E005_Out_OUT22_2003_17_1 : UINT;  (* RCON2 OUT22 2軸目 押付け制限 [255=100%] *)
    E005_Out_OUT23_2003_18_1 : UINT;  (* RCON2 OUT23 2軸目 制御信号（DSTR/SON等） *)
    E005_Out_OUT24_2003_19_1 : UINT;  (* RCON2 OUT24 3軸目 目標位置 下位 [0.01mm] *)
    E005_Out_OUT25_2003_1A_1 : UINT;  (* RCON2 OUT25 3軸目 目標位置 上位 [0.01mm] *)
    E005_Out_OUT26_2003_1B_1 : UINT;  (* RCON2 OUT26 3軸目 位置決め幅 下位 [0.01mm] *)
    E005_Out_OUT27_2003_1C_1 : UINT;  (* RCON2 OUT27 3軸目 位置決め幅 上位 [0.01mm] *)
    E005_Out_OUT28_2003_1D_1 : UINT;  (* RCON2 OUT28 3軸目 速度指令 [実機単位] *)
    E005_Out_OUT29_2003_1E_1 : UINT;  (* RCON2 OUT29 3軸目 共通加減速 [0.01G] *)
    E005_Out_OUT30_2003_1F_1 : UINT;  (* RCON2 OUT30 3軸目 押付け制限 [255=100%] *)
    E005_Out_OUT31_2003_20_1 : UINT;  (* RCON2 OUT31 3軸目 制御信号（DSTR/SON等） *)
    E005_Out_OUT32_2003_21_1 : UINT;  (* RCON2 OUT32 4軸目 目標位置 下位 [0.01mm] *)
    E005_Out_OUT33_2003_22_1 : UINT;  (* RCON2 OUT33 4軸目 目標位置 上位 [0.01mm] *)
    E005_Out_OUT34_2003_23_1 : UINT;  (* RCON2 OUT34 4軸目 位置決め幅 下位 [0.01mm] *)
    E005_Out_OUT35_2003_24_1 : UINT;  (* RCON2 OUT35 4軸目 位置決め幅 上位 [0.01mm] *)
    E005_Out_OUT36_2003_25_1 : UINT;  (* RCON2 OUT36 4軸目 速度指令 [実機単位] *)
    E005_Out_OUT37_2003_26_1 : UINT;  (* RCON2 OUT37 4軸目 共通加減速 [0.01G] *)
    E005_Out_OUT38_2003_27_1 : UINT;  (* RCON2 OUT38 4軸目 押付け制限 [255=100%] *)
    E005_Out_OUT39_2003_28_1 : UINT;  (* RCON2 OUT39 4軸目 制御信号（DSTR/SON等） *)
    E005_Out_OUT40_2003_29_1 : UINT;  (* RCON2 OUT40 5軸目 目標位置 下位 [0.01mm] *)
    E005_Out_OUT41_2003_2A_1 : UINT;  (* RCON2 OUT41 5軸目 目標位置 上位 [0.01mm] *)
    E005_Out_OUT42_2003_2B_1 : UINT;  (* RCON2 OUT42 5軸目 位置決め幅 下位 [0.01mm] *)
    E005_Out_OUT43_2003_2C_1 : UINT;  (* RCON2 OUT43 5軸目 位置決め幅 上位 [0.01mm] *)
    E005_Out_OUT44_2003_2D_1 : UINT;  (* RCON2 OUT44 5軸目 速度指令 [実機単位] *)
    E005_Out_OUT45_2003_2E_1 : UINT;  (* RCON2 OUT45 5軸目 共通加減速 [0.01G] *)
    E005_Out_OUT46_2003_2F_1 : UINT;  (* RCON2 OUT46 5軸目 押付け制限 [255=100%] *)
    E005_Out_OUT47_2003_30_1 : UINT;  (* RCON2 OUT47 5軸目 制御信号（DSTR/SON等） *)
    RCON1_AxisApply : ARRAY[1..6] OF BOOL;  (* RCON1 軸別出力更新許可（OFF=前値保持）; [1] A(左側) RCON1_1 NG1上下降 出力更新許可（OFF=前値保持）; [2] B(右側) RCON1_2 NG1上下降 出力更新許可（OFF=前値保持）; [3] A(左側) RCON1_3 SF/NG2送り 出力更新許可（OFF=前値保持）; [4] B(右側) RCON1_4 SF/NG2送り 出力更新許可（OFF=前値保持）; [5] A(左側) RCON1_5 SF/NG2上下降 出力更新許可（OFF=前値保持）; [6] B(右側) RCON1_6 SF/NG2上下降 出力更新許可（OFF=前値保持） *)
    RCON1_AxisLinked : ARRAY[1..6] OF BOOL;  (* RCON1 軸別リンク状態; [1] A(左側) RCON1_1 NG1上下降 リンク状態; [2] B(右側) RCON1_2 NG1上下降 リンク状態; [3] A(左側) RCON1_3 SF/NG2送り リンク状態; [4] B(右側) RCON1_4 SF/NG2送り リンク状態; [5] A(左側) RCON1_5 SF/NG2上下降 リンク状態; [6] B(右側) RCON1_6 SF/NG2上下降 リンク状態 *)
    RCON1_AxisWritten : ARRAY[1..6] OF BOOL;  (* RCON1 軸別出力代入済み（RCON受付とは別）; [1] A(左側) RCON1_1 NG1上下降 出力代入済み（RCON受付とは別）; [2] B(右側) RCON1_2 NG1上下降 出力代入済み（RCON受付とは別）; [3] A(左側) RCON1_3 SF/NG2送り 出力代入済み（RCON受付とは別）; [4] B(右側) RCON1_4 SF/NG2送り 出力代入済み（RCON受付とは別）; [5] A(左側) RCON1_5 SF/NG2上下降 出力代入済み（RCON受付とは別）; [6] B(右側) RCON1_6 SF/NG2上下降 出力代入済み（RCON受付とは別） *)
    RCON1_ByteOrderConfirmed : BOOL;  (* RCON1 ワード・バイト順確認済み（初期OFF） *)
    RCON1_CommOK : BOOL;  (* RCON1 通信正常（外部判定・固定ON不可） *)
    RCON1_EncodeError : ARRAY[1..6] OF UINT;  (* RCON1 軸別変換エラー番号（0=正常）; [1] A(左側) RCON1_1 NG1上下降 変換エラー番号; [2] B(右側) RCON1_2 NG1上下降 変換エラー番号; [3] A(左側) RCON1_3 SF/NG2送り 変換エラー番号; [4] B(右側) RCON1_4 SF/NG2送り 変換エラー番号; [5] A(左側) RCON1_5 SF/NG2上下降 変換エラー番号; [6] B(右側) RCON1_6 SF/NG2上下降 変換エラー番号 *)
    RCON1_EncodeOK : ARRAY[1..6] OF BOOL;  (* RCON1 軸別変換正常（運転許可とは別）; [1] A(左側) RCON1_1 NG1上下降 変換正常; [2] B(右側) RCON1_2 NG1上下降 変換正常; [3] A(左側) RCON1_3 SF/NG2送り 変換正常; [4] B(右側) RCON1_4 SF/NG2送り 変換正常; [5] A(左側) RCON1_5 SF/NG2上下降 変換正常; [6] B(右側) RCON1_6 SF/NG2上下降 変換正常 *)
    RCON1_GwAlarmCode : UINT;  (* RCON1 GW異常コード（ALMC/b0～7） *)
    RCON1_GwApply : BOOL;  (* RCON1 共通出力更新許可（OFF=前値保持） *)
    RCON1_GwAxisCommError : BOOL;  (* RCON1 GW－軸 通信異常（ERRT/b13） *)
    RCON1_GwControllerCommLatch : BOOL;  (* RCON1 GW通信異常保持（LERC/b14） *)
    RCON1_GwHeavyAlarm : BOOL;  (* RCON1 GW重故障（ALMH/b11） *)
    RCON1_GwLightAlarm : BOOL;  (* RCON1 GW軽故障（ALML/b10） *)
    RCON1_GwMON_Request : BOOL;  (* RCON1 MON要求（b15） *)
    RCON1_GwManual : BOOL;  (* RCON1 手動モード（MOD/b12） *)
    RCON1_GwRTE_Request : BOOL;  (* RCON1 通信異常ラッチ解除要求（b13） *)
    RCON1_GwRun : BOOL;  (* RCON1 GW動作中（RUN/b15） *)
    RCON1_GwSystemStop : BOOL;  (* RCON1 システム停止状態（SEMG/b8・監視用） *)
    RCON1_GwWritten : BOOL;  (* RCON1 共通出力代入済み（RCON受付とは別） *)
    RCON1_IN : ARRAY[1..6] OF ST_RCON_Direct_IN_Axis;  (* RCON1/Node1 6軸 入力（RCON→PLC）; [1] A(左側) RCON1_1 NG1排出(上下降); [2] B(右側) RCON1_2 NG1排出(上下降); [3] A(左側) RCON1_3 ストックフォルダ(SF)／NG2排出(送り); [4] B(右側) RCON1_4 ストックフォルダ(SF)／NG2排出(送り); [5] A(左側) RCON1_5 ストックフォルダ(SF)／NG2排出(上下降); [6] B(右側) RCON1_6 ストックフォルダ(SF)／NG2排出(上下降); [1].ActualPos_mm A(左側) RCON1_1 NG1上下降 現在位置 [mm]; [1].Current_mA A(左側) RCON1_1 NG1上下降 指令電流 [mA]（監視値）; [1].ActualSpeed_mm_s A(左側) RCON1_1 NG1上下降 現在速度 [mm/s・符号付き]; [1].AlarmCode A(左側) RCON1_1 NG1上下降 軸異常コード; [1].DataValid A(左側) RCON1_1 NG1上下降 入力有効（安全許可ではない）; [1].Status.PositionDone A(左側) RCON1_1 NG1上下降 位置決め完了; [1].Status.HomeDone A(左側) RCON1_1 NG1上下降 原点復帰完了; [1].Status.Moving A(左側) RCON1_1 NG1上下降 移動中; [1].Status.Alarm A(左側) RCON1_1 NG1上下降 軸異常; [1].Status.ServoReady A(左側) RCON1_1 NG1上下降 サーボON状態; [1].Status.PushMiss A(左側) RCON1_1 NG1上下降 押付け空振り（未使用）; [1].Status.OverloadWarning A(左側) RCON1_1 NG1上下降 過負荷警告; [1].Status.CommandDone A(左側) RCON1_1 NG1上下降 指令完了; [1].Status.Zone1 A(左側) RCON1_1 NG1上下降 ゾーン1内; [1].Status.Zone2 A(左側) RCON1_1 NG1上下降 ゾーン2内; [1].Status.ControllerReady A(左側) RCON1_1 NG1上下降 コントローラ準備完了; [1].Status.EmergencyStop A(左側) RCON1_1 NG1上下降 非常停止状態（入力）; [2].ActualPos_mm B(右側) RCON1_2 NG1上下降 現在位置 [mm]; [2].Current_mA B(右側) RCON1_2 NG1上下降 指令電流 [mA]（監視値）; [2].ActualSpeed_mm_s B(右側) RCON1_2 NG1上下降 現在速度 [mm/s・符号付き]; [2].AlarmCode B(右側) RCON1_2 NG1上下降 軸異常コード; [2].DataValid B(右側) RCON1_2 NG1上下降 入力有効（安全許可ではない）; [2].Status.PositionDone B(右側) RCON1_2 NG1上下降 位置決め完了; [2].Status.HomeDone B(右側) RCON1_2 NG1上下降 原点復帰完了; [2].Status.Moving B(右側) RCON1_2 NG1上下降 移動中; [2].Status.Alarm B(右側) RCON1_2 NG1上下降 軸異常; [2].Status.ServoReady B(右側) RCON1_2 NG1上下降 サーボON状態; [2].Status.PushMiss B(右側) RCON1_2 NG1上下降 押付け空振り（未使用）; [2].Status.OverloadWarning B(右側) RCON1_2 NG1上下降 過負荷警告; [2].Status.CommandDone B(右側) RCON1_2 NG1上下降 指令完了; [2].Status.Zone1 B(右側) RCON1_2 NG1上下降 ゾーン1内; [2].Status.Zone2 B(右側) RCON1_2 NG1上下降 ゾーン2内; [2].Status.ControllerReady B(右側) RCON1_2 NG1上下降 コントローラ準備完了; [2].Status.EmergencyStop B(右側) RCON1_2 NG1上下降 非常停止状態（入力）; [3].ActualPos_mm A(左側) RCON1_3 SF/NG2送り 現在位置 [mm]; [3].Current_mA A(左側) RCON1_3 SF/NG2送り 指令電流 [mA]（監視値）; [3].ActualSpeed_mm_s A(左側) RCON1_3 SF/NG2送り 現在速度 [mm/s・符号付き]; [3].AlarmCode A(左側) RCON1_3 SF/NG2送り 軸異常コード; [3].DataValid A(左側) RCON1_3 SF/NG2送り 入力有効（安全許可ではない）; [3].Status.PositionDone A(左側) RCON1_3 SF/NG2送り 位置決め完了; [3].Status.HomeDone A(左側) RCON1_3 SF/NG2送り 原点復帰完了; [3].Status.Moving A(左側) RCON1_3 SF/NG2送り 移動中; [3].Status.Alarm A(左側) RCON1_3 SF/NG2送り 軸異常; [3].Status.ServoReady A(左側) RCON1_3 SF/NG2送り サーボON状態; [3].Status.PushMiss A(左側) RCON1_3 SF/NG2送り 押付け空振り（未使用）; [3].Status.OverloadWarning A(左側) RCON1_3 SF/NG2送り 過負荷警告; [3].Status.CommandDone A(左側) RCON1_3 SF/NG2送り 指令完了; [3].Status.Zone1 A(左側) RCON1_3 SF/NG2送り ゾーン1内; [3].Status.Zone2 A(左側) RCON1_3 SF/NG2送り ゾーン2内; [3].Status.ControllerReady A(左側) RCON1_3 SF/NG2送り コントローラ準備完了; [3].Status.EmergencyStop A(左側) RCON1_3 SF/NG2送り 非常停止状態（入力）; [4].ActualPos_mm B(右側) RCON1_4 SF/NG2送り 現在位置 [mm]; [4].Current_mA B(右側) RCON1_4 SF/NG2送り 指令電流 [mA]（監視値）; [4].ActualSpeed_mm_s B(右側) RCON1_4 SF/NG2送り 現在速度 [mm/s・符号付き]; [4].AlarmCode B(右側) RCON1_4 SF/NG2送り 軸異常コード; [4].DataValid B(右側) RCON1_4 SF/NG2送り 入力有効（安全許可ではない）; [4].Status.PositionDone B(右側) RCON1_4 SF/NG2送り 位置決め完了; [4].Status.HomeDone B(右側) RCON1_4 SF/NG2送り 原点復帰完了; [4].Status.Moving B(右側) RCON1_4 SF/NG2送り 移動中; [4].Status.Alarm B(右側) RCON1_4 SF/NG2送り 軸異常; [4].Status.ServoReady B(右側) RCON1_4 SF/NG2送り サーボON状態; [4].Status.PushMiss B(右側) RCON1_4 SF/NG2送り 押付け空振り（未使用）; [4].Status.OverloadWarning B(右側) RCON1_4 SF/NG2送り 過負荷警告; [4].Status.CommandDone B(右側) RCON1_4 SF/NG2送り 指令完了; [4].Status.Zone1 B(右側) RCON1_4 SF/NG2送り ゾーン1内; [4].Status.Zone2 B(右側) RCON1_4 SF/NG2送り ゾーン2内; [4].Status.ControllerReady B(右側) RCON1_4 SF/NG2送り コントローラ準備完了; [4].Status.EmergencyStop B(右側) RCON1_4 SF/NG2送り 非常停止状態（入力）; [5].ActualPos_mm A(左側) RCON1_5 SF/NG2上下降 現在位置 [mm]; [5].Current_mA A(左側) RCON1_5 SF/NG2上下降 指令電流 [mA]（監視値）; [5].ActualSpeed_mm_s A(左側) RCON1_5 SF/NG2上下降 現在速度 [mm/s・符号付き]; [5].AlarmCode A(左側) RCON1_5 SF/NG2上下降 軸異常コード; [5].DataValid A(左側) RCON1_5 SF/NG2上下降 入力有効（安全許可ではない）; [5].Status.PositionDone A(左側) RCON1_5 SF/NG2上下降 位置決め完了; [5].Status.HomeDone A(左側) RCON1_5 SF/NG2上下降 原点復帰完了; [5].Status.Moving A(左側) RCON1_5 SF/NG2上下降 移動中; [5].Status.Alarm A(左側) RCON1_5 SF/NG2上下降 軸異常; [5].Status.ServoReady A(左側) RCON1_5 SF/NG2上下降 サーボON状態; [5].Status.PushMiss A(左側) RCON1_5 SF/NG2上下降 押付け空振り（未使用）; [5].Status.OverloadWarning A(左側) RCON1_5 SF/NG2上下降 過負荷警告; [5].Status.CommandDone A(左側) RCON1_5 SF/NG2上下降 指令完了; [5].Status.Zone1 A(左側) RCON1_5 SF/NG2上下降 ゾーン1内; [5].Status.Zone2 A(左側) RCON1_5 SF/NG2上下降 ゾーン2内; [5].Status.ControllerReady A(左側) RCON1_5 SF/NG2上下降 コントローラ準備完了; [5].Status.EmergencyStop A(左側) RCON1_5 SF/NG2上下降 非常停止状態（入力）; [6].ActualPos_mm B(右側) RCON1_6 SF/NG2上下降 現在位置 [mm]; [6].Current_mA B(右側) RCON1_6 SF/NG2上下降 指令電流 [mA]（監視値）; [6].ActualSpeed_mm_s B(右側) RCON1_6 SF/NG2上下降 現在速度 [mm/s・符号付き]; [6].AlarmCode B(右側) RCON1_6 SF/NG2上下降 軸異常コード; [6].DataValid B(右側) RCON1_6 SF/NG2上下降 入力有効（安全許可ではない）; [6].Status.PositionDone B(右側) RCON1_6 SF/NG2上下降 位置決め完了; [6].Status.HomeDone B(右側) RCON1_6 SF/NG2上下降 原点復帰完了; [6].Status.Moving B(右側) RCON1_6 SF/NG2上下降 移動中; [6].Status.Alarm B(右側) RCON1_6 SF/NG2上下降 軸異常; [6].Status.ServoReady B(右側) RCON1_6 SF/NG2上下降 サーボON状態; [6].Status.PushMiss B(右側) RCON1_6 SF/NG2上下降 押付け空振り（未使用）; [6].Status.OverloadWarning B(右側) RCON1_6 SF/NG2上下降 過負荷警告; [6].Status.CommandDone B(右側) RCON1_6 SF/NG2上下降 指令完了; [6].Status.Zone1 B(右側) RCON1_6 SF/NG2上下降 ゾーン1内; [6].Status.Zone2 B(右側) RCON1_6 SF/NG2上下降 ゾーン2内; [6].Status.ControllerReady B(右側) RCON1_6 SF/NG2上下降 コントローラ準備完了; [6].Status.EmergencyStop B(右側) RCON1_6 SF/NG2上下降 非常停止状態（入力） *)
    RCON1_LayoutConfirmed : BOOL;  (* RCON1 I/O配置確認済み（初期OFF） *)
    RCON1_MotionPermit : ARRAY[1..6] OF BOOL;  (* RCON1 軸別運転許可（外部判定・初期OFF）; [1] A(左側) RCON1_1 NG1上下降 運転許可（外部判定）; [2] B(右側) RCON1_2 NG1上下降 運転許可（外部判定）; [3] A(左側) RCON1_3 SF/NG2送り 運転許可（外部判定）; [4] B(右側) RCON1_4 SF/NG2送り 運転許可（外部判定）; [5] A(左側) RCON1_5 SF/NG2上下降 運転許可（外部判定）; [6] B(右側) RCON1_6 SF/NG2上下降 運転許可（外部判定） *)
    RCON1_OUT : ARRAY[1..6] OF ST_RCON_Direct_OUT_Axis;  (* RCON1/Node1 6軸 出力（PLC→RCON）; [2] B(右側) RCON1_2 NG1排出(上下降); [3] A(左側) RCON1_3 ストックフォルダ(SF)／NG2排出(送り); [4] B(右側) RCON1_4 ストックフォルダ(SF)／NG2排出(送り); [5] A(左側) RCON1_5 ストックフォルダ(SF)／NG2排出(上下降); [6] B(右側) RCON1_6 ストックフォルダ(SF)／NG2排出(上下降); [1].Control.Pause A(左側) RCON1_1 NG1上下降 一時停止要求（未接続）; [1] A(左側) RCON1_1 NG1排出(上下降); [1].TargetPos_mm A(左側) RCON1_1 NG1上下降 目標位置 [mm]; [1].PositionBand_mm A(左側) RCON1_1 NG1上下降 位置決め幅 [mm]; [1].Speed_mm_s A(左側) RCON1_1 NG1上下降 指令速度 [mm/s]; [1].AccDec_G A(左側) RCON1_1 NG1上下降 共通加減速度 [G]; [1].PushLimit_pct A(左側) RCON1_1 NG1上下降 押付け制限 [%]（未使用）; [1].Control.Start A(左側) RCON1_1 NG1上下降 移動開始要求（100ms保持）; [1].Control.Home A(左側) RCON1_1 NG1上下降 原点復帰要求（未接続）; [1].Control.Reset A(左側) RCON1_1 NG1上下降 異常リセット要求; [1].Control.ServoOn A(左側) RCON1_1 NG1上下降 サーボON要求（非常停止時OFF）; [1].Control.InchingSelect A(左側) RCON1_1 NG1上下降 インチング選択（OFF=ジョグ）; [1].Control.JogSpeedSelect A(左側) RCON1_1 NG1上下降 ジョグ速度切替（未接続）; [1].Control.JogMinus A(左側) RCON1_1 NG1上下降 原点方向ジョグ（未接続）; [1].Control.JogPlus A(左側) RCON1_1 NG1上下降 反原点方向ジョグ（未接続）; [1].Control.GainSelect0 A(左側) RCON1_1 NG1上下降 ゲイン選択下位（未使用）; [1].Control.GainSelect1 A(左側) RCON1_1 NG1上下降 ゲイン選択上位（未使用）; [1].Control.PushEnable A(左側) RCON1_1 NG1上下降 押付け選択（未使用・OFF=位置決め）; [1].Control.PushDirection A(左側) RCON1_1 NG1上下降 押付け方向（未使用）; [1].Control.RelativeMove A(左側) RCON1_1 NG1上下降 相対移動選択（未使用・OFF=絶対）; [1].Control.BrakeRelease A(左側) RCON1_1 NG1上下降 ブレーキ強制解除要求（非常停止でない間ON）; [2].TargetPos_mm B(右側) RCON1_2 NG1上下降 目標位置 [mm]; [2].PositionBand_mm B(右側) RCON1_2 NG1上下降 位置決め幅 [mm]; [2].Speed_mm_s B(右側) RCON1_2 NG1上下降 指令速度 [mm/s]; [2].AccDec_G B(右側) RCON1_2 NG1上下降 共通加減速度 [G]; [2].PushLimit_pct B(右側) RCON1_2 NG1上下降 押付け制限 [%]（未使用）; [2].Control.Start B(右側) RCON1_2 NG1上下降 移動開始要求（100ms保持）; [2].Control.Home B(右側) RCON1_2 NG1上下降 原点復帰要求（未接続）; [2].Control.Pause B(右側) RCON1_2 NG1上下降 一時停止要求（未接続）; [2].Control.Reset B(右側) RCON1_2 NG1上下降 異常リセット要求; [2].Control.ServoOn B(右側) RCON1_2 NG1上下降 サーボON要求（非常停止時OFF）; [2].Control.InchingSelect B(右側) RCON1_2 NG1上下降 インチング選択（OFF=ジョグ）; [2].Control.JogSpeedSelect B(右側) RCON1_2 NG1上下降 ジョグ速度切替（未接続）; [2].Control.JogMinus B(右側) RCON1_2 NG1上下降 原点方向ジョグ（未接続）; [2].Control.JogPlus B(右側) RCON1_2 NG1上下降 反原点方向ジョグ（未接続）; [2].Control.GainSelect0 B(右側) RCON1_2 NG1上下降 ゲイン選択下位（未使用）; [2].Control.GainSelect1 B(右側) RCON1_2 NG1上下降 ゲイン選択上位（未使用）; [2].Control.PushEnable B(右側) RCON1_2 NG1上下降 押付け選択（未使用・OFF=位置決め）; [2].Control.PushDirection B(右側) RCON1_2 NG1上下降 押付け方向（未使用）; [2].Control.RelativeMove B(右側) RCON1_2 NG1上下降 相対移動選択（未使用・OFF=絶対）; [2].Control.BrakeRelease B(右側) RCON1_2 NG1上下降 ブレーキ強制解除要求（非常停止でない間ON）; [3].TargetPos_mm A(左側) RCON1_3 SF/NG2送り 目標位置 [mm]; [3].PositionBand_mm A(左側) RCON1_3 SF/NG2送り 位置決め幅 [mm]; [3].Speed_mm_s A(左側) RCON1_3 SF/NG2送り 指令速度 [mm/s]; [3].AccDec_G A(左側) RCON1_3 SF/NG2送り 共通加減速度 [G]; [3].PushLimit_pct A(左側) RCON1_3 SF/NG2送り 押付け制限 [%]（未使用）; [3].Control.Start A(左側) RCON1_3 SF/NG2送り 移動開始要求（100ms保持）; [3].Control.Home A(左側) RCON1_3 SF/NG2送り 原点復帰要求（未接続）; [3].Control.Pause A(左側) RCON1_3 SF/NG2送り 一時停止要求（未接続）; [3].Control.Reset A(左側) RCON1_3 SF/NG2送り 異常リセット要求; [3].Control.ServoOn A(左側) RCON1_3 SF/NG2送り サーボON要求（非常停止時OFF）; [3].Control.InchingSelect A(左側) RCON1_3 SF/NG2送り インチング選択（OFF=ジョグ）; [3].Control.JogSpeedSelect A(左側) RCON1_3 SF/NG2送り ジョグ速度切替（未接続）; [3].Control.JogMinus A(左側) RCON1_3 SF/NG2送り 原点方向ジョグ（未接続）; [3].Control.JogPlus A(左側) RCON1_3 SF/NG2送り 反原点方向ジョグ（未接続）; [3].Control.GainSelect0 A(左側) RCON1_3 SF/NG2送り ゲイン選択下位（未使用）; [3].Control.GainSelect1 A(左側) RCON1_3 SF/NG2送り ゲイン選択上位（未使用）; [3].Control.PushEnable A(左側) RCON1_3 SF/NG2送り 押付け選択（未使用・OFF=位置決め）; [3].Control.PushDirection A(左側) RCON1_3 SF/NG2送り 押付け方向（未使用）; [3].Control.RelativeMove A(左側) RCON1_3 SF/NG2送り 相対移動選択（未使用・OFF=絶対）; [3].Control.BrakeRelease A(左側) RCON1_3 SF/NG2送り ブレーキ強制解除要求（非常停止でない間ON）; [4].TargetPos_mm B(右側) RCON1_4 SF/NG2送り 目標位置 [mm]; [4].PositionBand_mm B(右側) RCON1_4 SF/NG2送り 位置決め幅 [mm]; [4].Speed_mm_s B(右側) RCON1_4 SF/NG2送り 指令速度 [mm/s]; [4].AccDec_G B(右側) RCON1_4 SF/NG2送り 共通加減速度 [G]; [4].PushLimit_pct B(右側) RCON1_4 SF/NG2送り 押付け制限 [%]（未使用）; [4].Control.Start B(右側) RCON1_4 SF/NG2送り 移動開始要求（100ms保持）; [4].Control.Home B(右側) RCON1_4 SF/NG2送り 原点復帰要求（未接続）; [4].Control.Pause B(右側) RCON1_4 SF/NG2送り 一時停止要求（未接続）; [4].Control.Reset B(右側) RCON1_4 SF/NG2送り 異常リセット要求; [4].Control.ServoOn B(右側) RCON1_4 SF/NG2送り サーボON要求（非常停止時OFF）; [4].Control.InchingSelect B(右側) RCON1_4 SF/NG2送り インチング選択（OFF=ジョグ）; [4].Control.JogSpeedSelect B(右側) RCON1_4 SF/NG2送り ジョグ速度切替（未接続）; [4].Control.JogMinus B(右側) RCON1_4 SF/NG2送り 原点方向ジョグ（未接続）; [4].Control.JogPlus B(右側) RCON1_4 SF/NG2送り 反原点方向ジョグ（未接続）; [4].Control.GainSelect0 B(右側) RCON1_4 SF/NG2送り ゲイン選択下位（未使用）; [4].Control.GainSelect1 B(右側) RCON1_4 SF/NG2送り ゲイン選択上位（未使用）; [4].Control.PushEnable B(右側) RCON1_4 SF/NG2送り 押付け選択（未使用・OFF=位置決め）; [4].Control.PushDirection B(右側) RCON1_4 SF/NG2送り 押付け方向（未使用）; [4].Control.RelativeMove B(右側) RCON1_4 SF/NG2送り 相対移動選択（未使用・OFF=絶対）; [4].Control.BrakeRelease B(右側) RCON1_4 SF/NG2送り ブレーキ強制解除要求（非常停止でない間ON）; [5].TargetPos_mm A(左側) RCON1_5 SF/NG2上下降 目標位置 [mm]; [5].PositionBand_mm A(左側) RCON1_5 SF/NG2上下降 位置決め幅 [mm]; [5].Speed_mm_s A(左側) RCON1_5 SF/NG2上下降 指令速度 [mm/s]; [5].AccDec_G A(左側) RCON1_5 SF/NG2上下降 共通加減速度 [G]; [5].PushLimit_pct A(左側) RCON1_5 SF/NG2上下降 押付け制限 [%]（未使用）; [5].Control.Start A(左側) RCON1_5 SF/NG2上下降 移動開始要求（100ms保持）; [5].Control.Home A(左側) RCON1_5 SF/NG2上下降 原点復帰要求（未接続）; [5].Control.Pause A(左側) RCON1_5 SF/NG2上下降 一時停止要求（未接続）; [5].Control.Reset A(左側) RCON1_5 SF/NG2上下降 異常リセット要求; [5].Control.ServoOn A(左側) RCON1_5 SF/NG2上下降 サーボON要求（非常停止時OFF）; [5].Control.InchingSelect A(左側) RCON1_5 SF/NG2上下降 インチング選択（OFF=ジョグ）; [5].Control.JogSpeedSelect A(左側) RCON1_5 SF/NG2上下降 ジョグ速度切替（未接続）; [5].Control.JogMinus A(左側) RCON1_5 SF/NG2上下降 原点方向ジョグ（未接続）; [5].Control.JogPlus A(左側) RCON1_5 SF/NG2上下降 反原点方向ジョグ（未接続）; [5].Control.GainSelect0 A(左側) RCON1_5 SF/NG2上下降 ゲイン選択下位（未使用）; [5].Control.GainSelect1 A(左側) RCON1_5 SF/NG2上下降 ゲイン選択上位（未使用）; [5].Control.PushEnable A(左側) RCON1_5 SF/NG2上下降 押付け選択（未使用・OFF=位置決め）; [5].Control.PushDirection A(左側) RCON1_5 SF/NG2上下降 押付け方向（未使用）; [5].Control.RelativeMove A(左側) RCON1_5 SF/NG2上下降 相対移動選択（未使用・OFF=絶対）; [5].Control.BrakeRelease A(左側) RCON1_5 SF/NG2上下降 ブレーキ強制解除要求（非常停止でない間ON）; [6].TargetPos_mm B(右側) RCON1_6 SF/NG2上下降 目標位置 [mm]; [6].PositionBand_mm B(右側) RCON1_6 SF/NG2上下降 位置決め幅 [mm]; [6].Speed_mm_s B(右側) RCON1_6 SF/NG2上下降 指令速度 [mm/s]; [6].AccDec_G B(右側) RCON1_6 SF/NG2上下降 共通加減速度 [G]; [6].PushLimit_pct B(右側) RCON1_6 SF/NG2上下降 押付け制限 [%]（未使用）; [6].Control.Start B(右側) RCON1_6 SF/NG2上下降 移動開始要求（100ms保持）; [6].Control.Home B(右側) RCON1_6 SF/NG2上下降 原点復帰要求（未接続）; [6].Control.Pause B(右側) RCON1_6 SF/NG2上下降 一時停止要求（未接続）; [6].Control.Reset B(右側) RCON1_6 SF/NG2上下降 異常リセット要求; [6].Control.ServoOn B(右側) RCON1_6 SF/NG2上下降 サーボON要求（非常停止時OFF）; [6].Control.InchingSelect B(右側) RCON1_6 SF/NG2上下降 インチング選択（OFF=ジョグ）; [6].Control.JogSpeedSelect B(右側) RCON1_6 SF/NG2上下降 ジョグ速度切替（未接続）; [6].Control.JogMinus B(右側) RCON1_6 SF/NG2上下降 原点方向ジョグ（未接続）; [6].Control.JogPlus B(右側) RCON1_6 SF/NG2上下降 反原点方向ジョグ（未接続）; [6].Control.GainSelect0 B(右側) RCON1_6 SF/NG2上下降 ゲイン選択下位（未使用）; [6].Control.GainSelect1 B(右側) RCON1_6 SF/NG2上下降 ゲイン選択上位（未使用）; [6].Control.PushEnable B(右側) RCON1_6 SF/NG2上下降 押付け選択（未使用・OFF=位置決め）; [6].Control.PushDirection B(右側) RCON1_6 SF/NG2上下降 押付け方向（未使用）; [6].Control.RelativeMove B(右側) RCON1_6 SF/NG2上下降 相対移動選択（未使用・OFF=絶対）; [6].Control.BrakeRelease B(右側) RCON1_6 SF/NG2上下降 ブレーキ強制解除要求（非常停止でない間ON） *)
    RCON1_PowerStateRaw : ARRAY[0..4] OF WORD;  (* RCON1 電源状態ワード（詳細未確認）; [0] IN02 電源状態0（詳細未確認）; [1] IN03 電源状態1（詳細未確認）; [2] IN04 電源状態2（詳細未確認）; [3] IN05 電源状態3（詳細未確認）; [4] IN06 電源状態4（詳細未確認） *)
    RCON1_RxRaw : ARRAY[0..55] OF UINT;  (* RCON1 受信値（バイト交換前）; [0] IN00 GW状態; [1] IN01 軸リンク状態; [2] IN02 電源状態0; [3] IN03 電源状態1; [4] IN04 電源状態2; [5] IN05 電源状態3; [6] IN06 電源状態4（構成依存）; [7] IN07 予約（使用禁止）; [8] IN08 A(左側) RCON1_1 NG1上下降 現在位置 下位 [0.01mm]; [9] IN09 A(左側) RCON1_1 NG1上下降 現在位置 上位 [0.01mm]; [10] IN10 A(左側) RCON1_1 NG1上下降 指令電流 下位 [mA]; [11] IN11 A(左側) RCON1_1 NG1上下降 指令電流 上位 [mA]; [12] IN12 A(左側) RCON1_1 NG1上下降 現在速度 [実機単位・符号付き]; [13] IN13 A(左側) RCON1_1 NG1上下降 予約（使用禁止）; [14] IN14 A(左側) RCON1_1 NG1上下降 軸異常コード; [15] IN15 A(左側) RCON1_1 NG1上下降 状態信号（PEND/SV等）; [16] IN16 B(右側) RCON1_2 NG1上下降 現在位置 下位 [0.01mm]; [17] IN17 B(右側) RCON1_2 NG1上下降 現在位置 上位 [0.01mm]; [18] IN18 B(右側) RCON1_2 NG1上下降 指令電流 下位 [mA]; [19] IN19 B(右側) RCON1_2 NG1上下降 指令電流 上位 [mA]; [20] IN20 B(右側) RCON1_2 NG1上下降 現在速度 [実機単位・符号付き]; [21] IN21 B(右側) RCON1_2 NG1上下降 予約（使用禁止）; [22] IN22 B(右側) RCON1_2 NG1上下降 軸異常コード; [23] IN23 B(右側) RCON1_2 NG1上下降 状態信号（PEND/SV等）; [24] IN24 A(左側) RCON1_3 SF/NG2送り 現在位置 下位 [0.01mm]; [25] IN25 A(左側) RCON1_3 SF/NG2送り 現在位置 上位 [0.01mm]; [26] IN26 A(左側) RCON1_3 SF/NG2送り 指令電流 下位 [mA]; [27] IN27 A(左側) RCON1_3 SF/NG2送り 指令電流 上位 [mA]; [28] IN28 A(左側) RCON1_3 SF/NG2送り 現在速度 [実機単位・符号付き]; [29] IN29 A(左側) RCON1_3 SF/NG2送り 予約（使用禁止）; [30] IN30 A(左側) RCON1_3 SF/NG2送り 軸異常コード; [31] IN31 A(左側) RCON1_3 SF/NG2送り 状態信号（PEND/SV等）; [32] IN32 B(右側) RCON1_4 SF/NG2送り 現在位置 下位 [0.01mm]; [33] IN33 B(右側) RCON1_4 SF/NG2送り 現在位置 上位 [0.01mm]; [34] IN34 B(右側) RCON1_4 SF/NG2送り 指令電流 下位 [mA]; [35] IN35 B(右側) RCON1_4 SF/NG2送り 指令電流 上位 [mA]; [36] IN36 B(右側) RCON1_4 SF/NG2送り 現在速度 [実機単位・符号付き]; [37] IN37 B(右側) RCON1_4 SF/NG2送り 予約（使用禁止）; [38] IN38 B(右側) RCON1_4 SF/NG2送り 軸異常コード; [39] IN39 B(右側) RCON1_4 SF/NG2送り 状態信号（PEND/SV等）; [40] IN40 A(左側) RCON1_5 SF/NG2上下降 現在位置 下位 [0.01mm]; [41] IN41 A(左側) RCON1_5 SF/NG2上下降 現在位置 上位 [0.01mm]; [42] IN42 A(左側) RCON1_5 SF/NG2上下降 指令電流 下位 [mA]; [43] IN43 A(左側) RCON1_5 SF/NG2上下降 指令電流 上位 [mA]; [44] IN44 A(左側) RCON1_5 SF/NG2上下降 現在速度 [実機単位・符号付き]; [45] IN45 A(左側) RCON1_5 SF/NG2上下降 予約（使用禁止）; [46] IN46 A(左側) RCON1_5 SF/NG2上下降 軸異常コード; [47] IN47 A(左側) RCON1_5 SF/NG2上下降 状態信号（PEND/SV等）; [48] IN48 B(右側) RCON1_6 SF/NG2上下降 現在位置 下位 [0.01mm]; [49] IN49 B(右側) RCON1_6 SF/NG2上下降 現在位置 上位 [0.01mm]; [50] IN50 B(右側) RCON1_6 SF/NG2上下降 指令電流 下位 [mA]; [51] IN51 B(右側) RCON1_6 SF/NG2上下降 指令電流 上位 [mA]; [52] IN52 B(右側) RCON1_6 SF/NG2上下降 現在速度 [実機単位・符号付き]; [53] IN53 B(右側) RCON1_6 SF/NG2上下降 予約（使用禁止）; [54] IN54 B(右側) RCON1_6 SF/NG2上下降 軸異常コード; [55] IN55 B(右側) RCON1_6 SF/NG2上下降 状態信号（PEND/SV等） *)
    RCON1_RxWord : ARRAY[0..55] OF WORD;  (* RCON1 受信ワード（正規化後）; [0] IN00 GW状態; [1] IN01 軸リンク状態; [2] IN02 電源状態0; [3] IN03 電源状態1; [4] IN04 電源状態2; [5] IN05 電源状態3; [6] IN06 電源状態4（構成依存）; [7] IN07 予約（使用禁止）; [8] IN08 A(左側) RCON1_1 NG1上下降 現在位置 下位 [0.01mm]; [9] IN09 A(左側) RCON1_1 NG1上下降 現在位置 上位 [0.01mm]; [10] IN10 A(左側) RCON1_1 NG1上下降 指令電流 下位 [mA]; [11] IN11 A(左側) RCON1_1 NG1上下降 指令電流 上位 [mA]; [12] IN12 A(左側) RCON1_1 NG1上下降 現在速度 [実機単位・符号付き]; [13] IN13 A(左側) RCON1_1 NG1上下降 予約（使用禁止）; [14] IN14 A(左側) RCON1_1 NG1上下降 軸異常コード; [15] IN15 A(左側) RCON1_1 NG1上下降 状態信号（PEND/SV等）; [16] IN16 B(右側) RCON1_2 NG1上下降 現在位置 下位 [0.01mm]; [17] IN17 B(右側) RCON1_2 NG1上下降 現在位置 上位 [0.01mm]; [18] IN18 B(右側) RCON1_2 NG1上下降 指令電流 下位 [mA]; [19] IN19 B(右側) RCON1_2 NG1上下降 指令電流 上位 [mA]; [20] IN20 B(右側) RCON1_2 NG1上下降 現在速度 [実機単位・符号付き]; [21] IN21 B(右側) RCON1_2 NG1上下降 予約（使用禁止）; [22] IN22 B(右側) RCON1_2 NG1上下降 軸異常コード; [23] IN23 B(右側) RCON1_2 NG1上下降 状態信号（PEND/SV等）; [24] IN24 A(左側) RCON1_3 SF/NG2送り 現在位置 下位 [0.01mm]; [25] IN25 A(左側) RCON1_3 SF/NG2送り 現在位置 上位 [0.01mm]; [26] IN26 A(左側) RCON1_3 SF/NG2送り 指令電流 下位 [mA]; [27] IN27 A(左側) RCON1_3 SF/NG2送り 指令電流 上位 [mA]; [28] IN28 A(左側) RCON1_3 SF/NG2送り 現在速度 [実機単位・符号付き]; [29] IN29 A(左側) RCON1_3 SF/NG2送り 予約（使用禁止）; [30] IN30 A(左側) RCON1_3 SF/NG2送り 軸異常コード; [31] IN31 A(左側) RCON1_3 SF/NG2送り 状態信号（PEND/SV等）; [32] IN32 B(右側) RCON1_4 SF/NG2送り 現在位置 下位 [0.01mm]; [33] IN33 B(右側) RCON1_4 SF/NG2送り 現在位置 上位 [0.01mm]; [34] IN34 B(右側) RCON1_4 SF/NG2送り 指令電流 下位 [mA]; [35] IN35 B(右側) RCON1_4 SF/NG2送り 指令電流 上位 [mA]; [36] IN36 B(右側) RCON1_4 SF/NG2送り 現在速度 [実機単位・符号付き]; [37] IN37 B(右側) RCON1_4 SF/NG2送り 予約（使用禁止）; [38] IN38 B(右側) RCON1_4 SF/NG2送り 軸異常コード; [39] IN39 B(右側) RCON1_4 SF/NG2送り 状態信号（PEND/SV等）; [40] IN40 A(左側) RCON1_5 SF/NG2上下降 現在位置 下位 [0.01mm]; [41] IN41 A(左側) RCON1_5 SF/NG2上下降 現在位置 上位 [0.01mm]; [42] IN42 A(左側) RCON1_5 SF/NG2上下降 指令電流 下位 [mA]; [43] IN43 A(左側) RCON1_5 SF/NG2上下降 指令電流 上位 [mA]; [44] IN44 A(左側) RCON1_5 SF/NG2上下降 現在速度 [実機単位・符号付き]; [45] IN45 A(左側) RCON1_5 SF/NG2上下降 予約（使用禁止）; [46] IN46 A(左側) RCON1_5 SF/NG2上下降 軸異常コード; [47] IN47 A(左側) RCON1_5 SF/NG2上下降 状態信号（PEND/SV等）; [48] IN48 B(右側) RCON1_6 SF/NG2上下降 現在位置 下位 [0.01mm]; [49] IN49 B(右側) RCON1_6 SF/NG2上下降 現在位置 上位 [0.01mm]; [50] IN50 B(右側) RCON1_6 SF/NG2上下降 指令電流 下位 [mA]; [51] IN51 B(右側) RCON1_6 SF/NG2上下降 指令電流 上位 [mA]; [52] IN52 B(右側) RCON1_6 SF/NG2上下降 現在速度 [実機単位・符号付き]; [53] IN53 B(右側) RCON1_6 SF/NG2上下降 予約（使用禁止）; [54] IN54 B(右側) RCON1_6 SF/NG2上下降 軸異常コード; [55] IN55 B(右側) RCON1_6 SF/NG2上下降 状態信号（PEND/SV等） *)
    RCON1_SpeedUnit_mm_s : LREAL;  (* RCON1 速度単位 [mm/s/カウント]（1.0/0.1） *)
    RCON1_SwapBytes : BOOL;  (* RCON1 上下バイト交換設定（ON=交換） *)
    RCON1_TxUInt : ARRAY[0..55] OF UINT;  (* RCON1 送信UINT候補（実I/Oではない）; [0] OUT00 共通制御（MON/RTE）; [1] OUT01 予約（書込禁止）; [2] OUT02 予約（書込禁止）; [3] OUT03 予約（書込禁止）; [4] OUT04 予約（書込禁止）; [5] OUT05 予約（書込禁止）; [6] OUT06 予約（書込禁止）; [7] OUT07 予約（書込禁止）; [8] OUT08 A(左側) RCON1_1 NG1上下降 目標位置 下位 [0.01mm]; [9] OUT09 A(左側) RCON1_1 NG1上下降 目標位置 上位 [0.01mm]; [10] OUT10 A(左側) RCON1_1 NG1上下降 位置決め幅 下位 [0.01mm]; [11] OUT11 A(左側) RCON1_1 NG1上下降 位置決め幅 上位 [0.01mm]; [12] OUT12 A(左側) RCON1_1 NG1上下降 速度指令 [実機単位]; [13] OUT13 A(左側) RCON1_1 NG1上下降 共通加減速 [0.01G]; [14] OUT14 A(左側) RCON1_1 NG1上下降 押付け制限 [255=100%]; [15] OUT15 A(左側) RCON1_1 NG1上下降 制御信号（DSTR/SON等）; [16] OUT16 B(右側) RCON1_2 NG1上下降 目標位置 下位 [0.01mm]; [17] OUT17 B(右側) RCON1_2 NG1上下降 目標位置 上位 [0.01mm]; [18] OUT18 B(右側) RCON1_2 NG1上下降 位置決め幅 下位 [0.01mm]; [19] OUT19 B(右側) RCON1_2 NG1上下降 位置決め幅 上位 [0.01mm]; [20] OUT20 B(右側) RCON1_2 NG1上下降 速度指令 [実機単位]; [21] OUT21 B(右側) RCON1_2 NG1上下降 共通加減速 [0.01G]; [22] OUT22 B(右側) RCON1_2 NG1上下降 押付け制限 [255=100%]; [23] OUT23 B(右側) RCON1_2 NG1上下降 制御信号（DSTR/SON等）; [24] OUT24 A(左側) RCON1_3 SF/NG2送り 目標位置 下位 [0.01mm]; [25] OUT25 A(左側) RCON1_3 SF/NG2送り 目標位置 上位 [0.01mm]; [26] OUT26 A(左側) RCON1_3 SF/NG2送り 位置決め幅 下位 [0.01mm]; [27] OUT27 A(左側) RCON1_3 SF/NG2送り 位置決め幅 上位 [0.01mm]; [28] OUT28 A(左側) RCON1_3 SF/NG2送り 速度指令 [実機単位]; [29] OUT29 A(左側) RCON1_3 SF/NG2送り 共通加減速 [0.01G]; [30] OUT30 A(左側) RCON1_3 SF/NG2送り 押付け制限 [255=100%]; [31] OUT31 A(左側) RCON1_3 SF/NG2送り 制御信号（DSTR/SON等）; [32] OUT32 B(右側) RCON1_4 SF/NG2送り 目標位置 下位 [0.01mm]; [33] OUT33 B(右側) RCON1_4 SF/NG2送り 目標位置 上位 [0.01mm]; [34] OUT34 B(右側) RCON1_4 SF/NG2送り 位置決め幅 下位 [0.01mm]; [35] OUT35 B(右側) RCON1_4 SF/NG2送り 位置決め幅 上位 [0.01mm]; [36] OUT36 B(右側) RCON1_4 SF/NG2送り 速度指令 [実機単位]; [37] OUT37 B(右側) RCON1_4 SF/NG2送り 共通加減速 [0.01G]; [38] OUT38 B(右側) RCON1_4 SF/NG2送り 押付け制限 [255=100%]; [39] OUT39 B(右側) RCON1_4 SF/NG2送り 制御信号（DSTR/SON等）; [40] OUT40 A(左側) RCON1_5 SF/NG2上下降 目標位置 下位 [0.01mm]; [41] OUT41 A(左側) RCON1_5 SF/NG2上下降 目標位置 上位 [0.01mm]; [42] OUT42 A(左側) RCON1_5 SF/NG2上下降 位置決め幅 下位 [0.01mm]; [43] OUT43 A(左側) RCON1_5 SF/NG2上下降 位置決め幅 上位 [0.01mm]; [44] OUT44 A(左側) RCON1_5 SF/NG2上下降 速度指令 [実機単位]; [45] OUT45 A(左側) RCON1_5 SF/NG2上下降 共通加減速 [0.01G]; [46] OUT46 A(左側) RCON1_5 SF/NG2上下降 押付け制限 [255=100%]; [47] OUT47 A(左側) RCON1_5 SF/NG2上下降 制御信号（DSTR/SON等）; [48] OUT48 B(右側) RCON1_6 SF/NG2上下降 目標位置 下位 [0.01mm]; [49] OUT49 B(右側) RCON1_6 SF/NG2上下降 目標位置 上位 [0.01mm]; [50] OUT50 B(右側) RCON1_6 SF/NG2上下降 位置決め幅 下位 [0.01mm]; [51] OUT51 B(右側) RCON1_6 SF/NG2上下降 位置決め幅 上位 [0.01mm]; [52] OUT52 B(右側) RCON1_6 SF/NG2上下降 速度指令 [実機単位]; [53] OUT53 B(右側) RCON1_6 SF/NG2上下降 共通加減速 [0.01G]; [54] OUT54 B(右側) RCON1_6 SF/NG2上下降 押付け制限 [255=100%]; [55] OUT55 B(右側) RCON1_6 SF/NG2上下降 制御信号（DSTR/SON等） *)
    RCON1_TxWord : ARRAY[0..55] OF WORD;  (* RCON1 送信ワード候補; [0] OUT00 共通制御（MON/RTE）; [1] OUT01 予約（書込禁止）; [2] OUT02 予約（書込禁止）; [3] OUT03 予約（書込禁止）; [4] OUT04 予約（書込禁止）; [5] OUT05 予約（書込禁止）; [6] OUT06 予約（書込禁止）; [7] OUT07 予約（書込禁止）; [8] OUT08 A(左側) RCON1_1 NG1上下降 目標位置 下位 [0.01mm]; [9] OUT09 A(左側) RCON1_1 NG1上下降 目標位置 上位 [0.01mm]; [10] OUT10 A(左側) RCON1_1 NG1上下降 位置決め幅 下位 [0.01mm]; [11] OUT11 A(左側) RCON1_1 NG1上下降 位置決め幅 上位 [0.01mm]; [12] OUT12 A(左側) RCON1_1 NG1上下降 速度指令 [実機単位]; [13] OUT13 A(左側) RCON1_1 NG1上下降 共通加減速 [0.01G]; [14] OUT14 A(左側) RCON1_1 NG1上下降 押付け制限 [255=100%]; [15] OUT15 A(左側) RCON1_1 NG1上下降 制御信号（DSTR/SON等）; [16] OUT16 B(右側) RCON1_2 NG1上下降 目標位置 下位 [0.01mm]; [17] OUT17 B(右側) RCON1_2 NG1上下降 目標位置 上位 [0.01mm]; [18] OUT18 B(右側) RCON1_2 NG1上下降 位置決め幅 下位 [0.01mm]; [19] OUT19 B(右側) RCON1_2 NG1上下降 位置決め幅 上位 [0.01mm]; [20] OUT20 B(右側) RCON1_2 NG1上下降 速度指令 [実機単位]; [21] OUT21 B(右側) RCON1_2 NG1上下降 共通加減速 [0.01G]; [22] OUT22 B(右側) RCON1_2 NG1上下降 押付け制限 [255=100%]; [23] OUT23 B(右側) RCON1_2 NG1上下降 制御信号（DSTR/SON等）; [24] OUT24 A(左側) RCON1_3 SF/NG2送り 目標位置 下位 [0.01mm]; [25] OUT25 A(左側) RCON1_3 SF/NG2送り 目標位置 上位 [0.01mm]; [26] OUT26 A(左側) RCON1_3 SF/NG2送り 位置決め幅 下位 [0.01mm]; [27] OUT27 A(左側) RCON1_3 SF/NG2送り 位置決め幅 上位 [0.01mm]; [28] OUT28 A(左側) RCON1_3 SF/NG2送り 速度指令 [実機単位]; [29] OUT29 A(左側) RCON1_3 SF/NG2送り 共通加減速 [0.01G]; [30] OUT30 A(左側) RCON1_3 SF/NG2送り 押付け制限 [255=100%]; [31] OUT31 A(左側) RCON1_3 SF/NG2送り 制御信号（DSTR/SON等）; [32] OUT32 B(右側) RCON1_4 SF/NG2送り 目標位置 下位 [0.01mm]; [33] OUT33 B(右側) RCON1_4 SF/NG2送り 目標位置 上位 [0.01mm]; [34] OUT34 B(右側) RCON1_4 SF/NG2送り 位置決め幅 下位 [0.01mm]; [35] OUT35 B(右側) RCON1_4 SF/NG2送り 位置決め幅 上位 [0.01mm]; [36] OUT36 B(右側) RCON1_4 SF/NG2送り 速度指令 [実機単位]; [37] OUT37 B(右側) RCON1_4 SF/NG2送り 共通加減速 [0.01G]; [38] OUT38 B(右側) RCON1_4 SF/NG2送り 押付け制限 [255=100%]; [39] OUT39 B(右側) RCON1_4 SF/NG2送り 制御信号（DSTR/SON等）; [40] OUT40 A(左側) RCON1_5 SF/NG2上下降 目標位置 下位 [0.01mm]; [41] OUT41 A(左側) RCON1_5 SF/NG2上下降 目標位置 上位 [0.01mm]; [42] OUT42 A(左側) RCON1_5 SF/NG2上下降 位置決め幅 下位 [0.01mm]; [43] OUT43 A(左側) RCON1_5 SF/NG2上下降 位置決め幅 上位 [0.01mm]; [44] OUT44 A(左側) RCON1_5 SF/NG2上下降 速度指令 [実機単位]; [45] OUT45 A(左側) RCON1_5 SF/NG2上下降 共通加減速 [0.01G]; [46] OUT46 A(左側) RCON1_5 SF/NG2上下降 押付け制限 [255=100%]; [47] OUT47 A(左側) RCON1_5 SF/NG2上下降 制御信号（DSTR/SON等）; [48] OUT48 B(右側) RCON1_6 SF/NG2上下降 目標位置 下位 [0.01mm]; [49] OUT49 B(右側) RCON1_6 SF/NG2上下降 目標位置 上位 [0.01mm]; [50] OUT50 B(右側) RCON1_6 SF/NG2上下降 位置決め幅 下位 [0.01mm]; [51] OUT51 B(右側) RCON1_6 SF/NG2上下降 位置決め幅 上位 [0.01mm]; [52] OUT52 B(右側) RCON1_6 SF/NG2上下降 速度指令 [実機単位]; [53] OUT53 B(右側) RCON1_6 SF/NG2上下降 共通加減速 [0.01G]; [54] OUT54 B(右側) RCON1_6 SF/NG2上下降 押付け制限 [255=100%]; [55] OUT55 B(右側) RCON1_6 SF/NG2上下降 制御信号（DSTR/SON等） *)
    RCON1_WriteEnable : BOOL;  (* RCON1 実出力書込み許可（OFF=前値保持・停止不可） *)
    RCON2_AxisApply : ARRAY[1..5] OF BOOL;  (* RCON2 軸別出力更新許可（OFF=前値保持）; [1] 1軸目（No.0）出力更新許可（OFF=前値保持）; [2] 2軸目（No.1）出力更新許可（OFF=前値保持）; [3] 3軸目（No.2）出力更新許可（OFF=前値保持）; [4] 4軸目（No.3）出力更新許可（OFF=前値保持）; [5] 5軸目（No.4）出力更新許可（OFF=前値保持） *)
    RCON2_AxisLinked : ARRAY[1..5] OF BOOL;  (* RCON2 軸別リンク状態; [1] 1軸目（No.0）リンク状態; [2] 2軸目（No.1）リンク状態; [3] 3軸目（No.2）リンク状態; [4] 4軸目（No.3）リンク状態; [5] 5軸目（No.4）リンク状態 *)
    RCON2_AxisWritten : ARRAY[1..5] OF BOOL;  (* RCON2 軸別出力代入済み（RCON受付とは別）; [1] 1軸目（No.0）出力代入済み（RCON受付とは別）; [2] 2軸目（No.1）出力代入済み（RCON受付とは別）; [3] 3軸目（No.2）出力代入済み（RCON受付とは別）; [4] 4軸目（No.3）出力代入済み（RCON受付とは別）; [5] 5軸目（No.4）出力代入済み（RCON受付とは別） *)
    RCON2_ByteOrderConfirmed : BOOL;  (* RCON2 ワード・バイト順確認済み（初期OFF） *)
    RCON2_CommOK : BOOL;  (* RCON2 通信正常（外部判定・固定ON不可） *)
    RCON2_EncodeError : ARRAY[1..5] OF UINT;  (* RCON2 軸別変換エラー番号（0=正常）; [1] 1軸目（No.0）変換エラー番号; [2] 2軸目（No.1）変換エラー番号; [3] 3軸目（No.2）変換エラー番号; [4] 4軸目（No.3）変換エラー番号; [5] 5軸目（No.4）変換エラー番号 *)
    RCON2_EncodeOK : ARRAY[1..5] OF BOOL;  (* RCON2 軸別変換正常（運転許可とは別）; [1] 1軸目（No.0）変換正常; [2] 2軸目（No.1）変換正常; [3] 3軸目（No.2）変換正常; [4] 4軸目（No.3）変換正常; [5] 5軸目（No.4）変換正常 *)
    RCON2_GwAlarmCode : UINT;  (* RCON2 GW異常コード（ALMC/b0～7） *)
    RCON2_GwApply : BOOL;  (* RCON2 共通出力更新許可（OFF=前値保持） *)
    RCON2_GwAxisCommError : BOOL;  (* RCON2 GW－軸 通信異常（ERRT/b13） *)
    RCON2_GwControllerCommLatch : BOOL;  (* RCON2 GW通信異常保持（LERC/b14） *)
    RCON2_GwHeavyAlarm : BOOL;  (* RCON2 GW重故障（ALMH/b11） *)
    RCON2_GwLightAlarm : BOOL;  (* RCON2 GW軽故障（ALML/b10） *)
    RCON2_GwMON_Request : BOOL;  (* RCON2 MON要求（b15） *)
    RCON2_GwManual : BOOL;  (* RCON2 手動モード（MOD/b12） *)
    RCON2_GwRTE_Request : BOOL;  (* RCON2 通信異常ラッチ解除要求（b13） *)
    RCON2_GwRun : BOOL;  (* RCON2 GW動作中（RUN/b15） *)
    RCON2_GwSystemStop : BOOL;  (* RCON2 システム停止状態（SEMG/b8・監視用） *)
    RCON2_GwWritten : BOOL;  (* RCON2 共通出力代入済み（RCON受付とは別） *)
    RCON2_IN : ARRAY[1..5] OF ST_RCON_Direct_IN_Axis;  (* RCON2 入力情報（RCON→PLC）; [1] 1軸目（No.0）入力情報; [2] 2軸目（No.1）入力情報; [3] 3軸目（No.2）入力情報; [4] 4軸目（No.3）入力情報; [5] 5軸目（No.4）入力情報 *)
    RCON2_LayoutConfirmed : BOOL;  (* RCON2 I/O配置確認済み（初期OFF） *)
    RCON2_MotionPermit : ARRAY[1..5] OF BOOL;  (* RCON2 軸別運転許可（外部判定・初期OFF）; [1] 1軸目（No.0）運転許可（外部判定）; [2] 2軸目（No.1）運転許可（外部判定）; [3] 3軸目（No.2）運転許可（外部判定）; [4] 4軸目（No.3）運転許可（外部判定）; [5] 5軸目（No.4）運転許可（外部判定） *)
    RCON2_OUT : ARRAY[1..5] OF ST_RCON_Direct_OUT_Axis;  (* RCON2 出力指令（PLC→RCON）; [1] 1軸目（No.0）出力指令; [2] 2軸目（No.1）出力指令; [3] 3軸目（No.2）出力指令; [4] 4軸目（No.3）出力指令; [5] 5軸目（No.4）出力指令 *)
    RCON2_PowerStateRaw : ARRAY[0..4] OF WORD;  (* RCON2 電源状態ワード（詳細未確認）; [0] IN02 電源状態0（詳細未確認）; [1] IN03 電源状態1（詳細未確認）; [2] IN04 電源状態2（詳細未確認）; [3] IN05 電源状態3（詳細未確認）; [4] IN06 電源状態4（詳細未確認） *)
    RCON2_RxRaw : ARRAY[0..55] OF UINT;  (* RCON2 受信値（バイト交換前）; [0] IN00 GW状態; [1] IN01 軸リンク状態; [2] IN02 電源状態0; [3] IN03 電源状態1; [4] IN04 電源状態2; [5] IN05 電源状態3; [6] IN06 電源状態4（構成依存）; [7] IN07 予約（使用禁止）; [8] IN08 1軸目 現在位置 下位 [0.01mm]; [9] IN09 1軸目 現在位置 上位 [0.01mm]; [10] IN10 1軸目 指令電流 下位 [mA]; [11] IN11 1軸目 指令電流 上位 [mA]; [12] IN12 1軸目 現在速度 [実機単位・符号付き]; [13] IN13 1軸目 予約（使用禁止）; [14] IN14 1軸目 軸異常コード; [15] IN15 1軸目 状態信号（PEND/SV等）; [16] IN16 2軸目 現在位置 下位 [0.01mm]; [17] IN17 2軸目 現在位置 上位 [0.01mm]; [18] IN18 2軸目 指令電流 下位 [mA]; [19] IN19 2軸目 指令電流 上位 [mA]; [20] IN20 2軸目 現在速度 [実機単位・符号付き]; [21] IN21 2軸目 予約（使用禁止）; [22] IN22 2軸目 軸異常コード; [23] IN23 2軸目 状態信号（PEND/SV等）; [24] IN24 3軸目 現在位置 下位 [0.01mm]; [25] IN25 3軸目 現在位置 上位 [0.01mm]; [26] IN26 3軸目 指令電流 下位 [mA]; [27] IN27 3軸目 指令電流 上位 [mA]; [28] IN28 3軸目 現在速度 [実機単位・符号付き]; [29] IN29 3軸目 予約（使用禁止）; [30] IN30 3軸目 軸異常コード; [31] IN31 3軸目 状態信号（PEND/SV等）; [32] IN32 4軸目 現在位置 下位 [0.01mm]; [33] IN33 4軸目 現在位置 上位 [0.01mm]; [34] IN34 4軸目 指令電流 下位 [mA]; [35] IN35 4軸目 指令電流 上位 [mA]; [36] IN36 4軸目 現在速度 [実機単位・符号付き]; [37] IN37 4軸目 予約（使用禁止）; [38] IN38 4軸目 軸異常コード; [39] IN39 4軸目 状態信号（PEND/SV等）; [40] IN40 5軸目 現在位置 下位 [0.01mm]; [41] IN41 5軸目 現在位置 上位 [0.01mm]; [42] IN42 5軸目 指令電流 下位 [mA]; [43] IN43 5軸目 指令電流 上位 [mA]; [44] IN44 5軸目 現在速度 [実機単位・符号付き]; [45] IN45 5軸目 予約（使用禁止）; [46] IN46 5軸目 軸異常コード; [47] IN47 5軸目 状態信号（PEND/SV等）; [48] IN48 用途未確認（今回未使用）; [49] IN49 用途未確認（今回未使用）; [50] IN50 用途未確認（今回未使用）; [51] IN51 用途未確認（今回未使用）; [52] IN52 用途未確認（今回未使用）; [53] IN53 用途未確認（今回未使用）; [54] IN54 用途未確認（今回未使用）; [55] IN55 用途未確認（今回未使用） *)
    RCON2_RxWord : ARRAY[0..55] OF WORD;  (* RCON2 受信ワード（正規化後）; [0] IN00 GW状態; [1] IN01 軸リンク状態; [2] IN02 電源状態0; [3] IN03 電源状態1; [4] IN04 電源状態2; [5] IN05 電源状態3; [6] IN06 電源状態4（構成依存）; [7] IN07 予約（使用禁止）; [8] IN08 1軸目 現在位置 下位 [0.01mm]; [9] IN09 1軸目 現在位置 上位 [0.01mm]; [10] IN10 1軸目 指令電流 下位 [mA]; [11] IN11 1軸目 指令電流 上位 [mA]; [12] IN12 1軸目 現在速度 [実機単位・符号付き]; [13] IN13 1軸目 予約（使用禁止）; [14] IN14 1軸目 軸異常コード; [15] IN15 1軸目 状態信号（PEND/SV等）; [16] IN16 2軸目 現在位置 下位 [0.01mm]; [17] IN17 2軸目 現在位置 上位 [0.01mm]; [18] IN18 2軸目 指令電流 下位 [mA]; [19] IN19 2軸目 指令電流 上位 [mA]; [20] IN20 2軸目 現在速度 [実機単位・符号付き]; [21] IN21 2軸目 予約（使用禁止）; [22] IN22 2軸目 軸異常コード; [23] IN23 2軸目 状態信号（PEND/SV等）; [24] IN24 3軸目 現在位置 下位 [0.01mm]; [25] IN25 3軸目 現在位置 上位 [0.01mm]; [26] IN26 3軸目 指令電流 下位 [mA]; [27] IN27 3軸目 指令電流 上位 [mA]; [28] IN28 3軸目 現在速度 [実機単位・符号付き]; [29] IN29 3軸目 予約（使用禁止）; [30] IN30 3軸目 軸異常コード; [31] IN31 3軸目 状態信号（PEND/SV等）; [32] IN32 4軸目 現在位置 下位 [0.01mm]; [33] IN33 4軸目 現在位置 上位 [0.01mm]; [34] IN34 4軸目 指令電流 下位 [mA]; [35] IN35 4軸目 指令電流 上位 [mA]; [36] IN36 4軸目 現在速度 [実機単位・符号付き]; [37] IN37 4軸目 予約（使用禁止）; [38] IN38 4軸目 軸異常コード; [39] IN39 4軸目 状態信号（PEND/SV等）; [40] IN40 5軸目 現在位置 下位 [0.01mm]; [41] IN41 5軸目 現在位置 上位 [0.01mm]; [42] IN42 5軸目 指令電流 下位 [mA]; [43] IN43 5軸目 指令電流 上位 [mA]; [44] IN44 5軸目 現在速度 [実機単位・符号付き]; [45] IN45 5軸目 予約（使用禁止）; [46] IN46 5軸目 軸異常コード; [47] IN47 5軸目 状態信号（PEND/SV等）; [48] IN48 用途未確認（今回未使用）; [49] IN49 用途未確認（今回未使用）; [50] IN50 用途未確認（今回未使用）; [51] IN51 用途未確認（今回未使用）; [52] IN52 用途未確認（今回未使用）; [53] IN53 用途未確認（今回未使用）; [54] IN54 用途未確認（今回未使用）; [55] IN55 用途未確認（今回未使用） *)
    RCON2_SpeedUnit_mm_s : LREAL;  (* RCON2 速度単位 [mm/s/カウント]（1.0/0.1） *)
    RCON2_SwapBytes : BOOL;  (* RCON2 上下バイト交換設定（ON=交換） *)
    RCON2_TxUInt : ARRAY[0..47] OF UINT;  (* RCON2 送信UINT候補（実I/Oではない）; [0] OUT00 共通制御（MON/RTE）; [1] OUT01 予約（書込禁止）; [2] OUT02 予約（書込禁止）; [3] OUT03 予約（書込禁止）; [4] OUT04 予約（書込禁止）; [5] OUT05 予約（書込禁止）; [6] OUT06 予約（書込禁止）; [7] OUT07 予約（書込禁止）; [8] OUT08 1軸目 目標位置 下位 [0.01mm]; [9] OUT09 1軸目 目標位置 上位 [0.01mm]; [10] OUT10 1軸目 位置決め幅 下位 [0.01mm]; [11] OUT11 1軸目 位置決め幅 上位 [0.01mm]; [12] OUT12 1軸目 速度指令 [実機単位]; [13] OUT13 1軸目 共通加減速 [0.01G]; [14] OUT14 1軸目 押付け制限 [255=100%]; [15] OUT15 1軸目 制御信号（DSTR/SON等）; [16] OUT16 2軸目 目標位置 下位 [0.01mm]; [17] OUT17 2軸目 目標位置 上位 [0.01mm]; [18] OUT18 2軸目 位置決め幅 下位 [0.01mm]; [19] OUT19 2軸目 位置決め幅 上位 [0.01mm]; [20] OUT20 2軸目 速度指令 [実機単位]; [21] OUT21 2軸目 共通加減速 [0.01G]; [22] OUT22 2軸目 押付け制限 [255=100%]; [23] OUT23 2軸目 制御信号（DSTR/SON等）; [24] OUT24 3軸目 目標位置 下位 [0.01mm]; [25] OUT25 3軸目 目標位置 上位 [0.01mm]; [26] OUT26 3軸目 位置決め幅 下位 [0.01mm]; [27] OUT27 3軸目 位置決め幅 上位 [0.01mm]; [28] OUT28 3軸目 速度指令 [実機単位]; [29] OUT29 3軸目 共通加減速 [0.01G]; [30] OUT30 3軸目 押付け制限 [255=100%]; [31] OUT31 3軸目 制御信号（DSTR/SON等）; [32] OUT32 4軸目 目標位置 下位 [0.01mm]; [33] OUT33 4軸目 目標位置 上位 [0.01mm]; [34] OUT34 4軸目 位置決め幅 下位 [0.01mm]; [35] OUT35 4軸目 位置決め幅 上位 [0.01mm]; [36] OUT36 4軸目 速度指令 [実機単位]; [37] OUT37 4軸目 共通加減速 [0.01G]; [38] OUT38 4軸目 押付け制限 [255=100%]; [39] OUT39 4軸目 制御信号（DSTR/SON等）; [40] OUT40 5軸目 目標位置 下位 [0.01mm]; [41] OUT41 5軸目 目標位置 上位 [0.01mm]; [42] OUT42 5軸目 位置決め幅 下位 [0.01mm]; [43] OUT43 5軸目 位置決め幅 上位 [0.01mm]; [44] OUT44 5軸目 速度指令 [実機単位]; [45] OUT45 5軸目 共通加減速 [0.01G]; [46] OUT46 5軸目 押付け制限 [255=100%]; [47] OUT47 5軸目 制御信号（DSTR/SON等） *)
    RCON2_TxWord : ARRAY[0..47] OF WORD;  (* RCON2 送信ワード候補; [0] OUT00 共通制御（MON/RTE）; [1] OUT01 予約（書込禁止）; [2] OUT02 予約（書込禁止）; [3] OUT03 予約（書込禁止）; [4] OUT04 予約（書込禁止）; [5] OUT05 予約（書込禁止）; [6] OUT06 予約（書込禁止）; [7] OUT07 予約（書込禁止）; [8] OUT08 1軸目 目標位置 下位 [0.01mm]; [9] OUT09 1軸目 目標位置 上位 [0.01mm]; [10] OUT10 1軸目 位置決め幅 下位 [0.01mm]; [11] OUT11 1軸目 位置決め幅 上位 [0.01mm]; [12] OUT12 1軸目 速度指令 [実機単位]; [13] OUT13 1軸目 共通加減速 [0.01G]; [14] OUT14 1軸目 押付け制限 [255=100%]; [15] OUT15 1軸目 制御信号（DSTR/SON等）; [16] OUT16 2軸目 目標位置 下位 [0.01mm]; [17] OUT17 2軸目 目標位置 上位 [0.01mm]; [18] OUT18 2軸目 位置決め幅 下位 [0.01mm]; [19] OUT19 2軸目 位置決め幅 上位 [0.01mm]; [20] OUT20 2軸目 速度指令 [実機単位]; [21] OUT21 2軸目 共通加減速 [0.01G]; [22] OUT22 2軸目 押付け制限 [255=100%]; [23] OUT23 2軸目 制御信号（DSTR/SON等）; [24] OUT24 3軸目 目標位置 下位 [0.01mm]; [25] OUT25 3軸目 目標位置 上位 [0.01mm]; [26] OUT26 3軸目 位置決め幅 下位 [0.01mm]; [27] OUT27 3軸目 位置決め幅 上位 [0.01mm]; [28] OUT28 3軸目 速度指令 [実機単位]; [29] OUT29 3軸目 共通加減速 [0.01G]; [30] OUT30 3軸目 押付け制限 [255=100%]; [31] OUT31 3軸目 制御信号（DSTR/SON等）; [32] OUT32 4軸目 目標位置 下位 [0.01mm]; [33] OUT33 4軸目 目標位置 上位 [0.01mm]; [34] OUT34 4軸目 位置決め幅 下位 [0.01mm]; [35] OUT35 4軸目 位置決め幅 上位 [0.01mm]; [36] OUT36 4軸目 速度指令 [実機単位]; [37] OUT37 4軸目 共通加減速 [0.01G]; [38] OUT38 4軸目 押付け制限 [255=100%]; [39] OUT39 4軸目 制御信号（DSTR/SON等）; [40] OUT40 5軸目 目標位置 下位 [0.01mm]; [41] OUT41 5軸目 目標位置 上位 [0.01mm]; [42] OUT42 5軸目 位置決め幅 下位 [0.01mm]; [43] OUT43 5軸目 位置決め幅 上位 [0.01mm]; [44] OUT44 5軸目 速度指令 [実機単位]; [45] OUT45 5軸目 共通加減速 [0.01G]; [46] OUT46 5軸目 押付け制限 [255=100%]; [47] OUT47 5軸目 制御信号（DSTR/SON等） *)
    RCON2_WriteEnable : BOOL;  (* RCON2 実出力書込み許可（OFF=前値保持・停止不可） *)
    RCON1_IAI_Auto : ARRAY[0..99] OF Bool;  (* A(左側) RCON1_1 NG1上下降 自動移動要求; [1] A(左側) RCON1_1 NG1上下降 原点位置移動; [2] A(左側) RCON1_1 NG1上下降 NG仕分け; [3] A(左側) RCON1_1 NG1上下降 動作完了後 原点位置移動 *)
    RCON1_OUT_PositionBand_mm : LREAL;  (* A(左側) RCON1_1 NG1上下降 位置決め幅 [mm] *)
    RCON1_OUT_TargetPos_mm : LREAL;  (* A(左側) RCON1_1 NG1上下降 目標位置 [mm] *)
    RCON1_OUT_Speed_mm_s : LREAL;  (* A(左側) RCON1_1 NG1上下降 指令速度 [mm/s] *)
    RCON1_OUT_AccDec_G : LREAL;  (* A(左側) RCON1_1 NG1上下降 共通加減速度 [G] *)
    RCON1_OUT_PushLimit_pct : LREAL;  (* A(左側) RCON1_1 NG1上下降 押付け制限 [%]（未使用） *)
    RCON1_ActualPos_mm : LREAL;  (* A(左側) RCON1_1 NG1上下降 現在位置 [mm] *)
    RCON1_Current_mA : DINT;  (* A(左側) RCON1_1 NG1上下降 指令電流 [mA]（監視値） *)
    RCON1_ActualSpeed_mm_s : LREAL;  (* A(左側) RCON1_1 NG1上下降 現在速度 [mm/s・符号付き] *)
    RCON1_AlarmCode : UINT;  (* A(左側) RCON1_1 NG1上下降 軸異常コード *)
    RCON1_DataValid : BOOL;  (* A(左側) RCON1_1 NG1上下降 入力有効（安全許可ではない） *)
    RCON1_1_IN_PositionDone : BOOL;  (* A(左側) RCON1_1 NG1上下降 位置決め完了 *)
    RCON1_1_IN_HomeDone : BOOL;  (* A(左側) RCON1_1 NG1上下降 原点復帰完了 *)
    RCON1_1_IN_Moving : BOOL;  (* A(左側) RCON1_1 NG1上下降 移動中 *)
    RCON1_1_IN_EmergencyStop : BOOL;  (* A(左側) RCON1_1 NG1上下降 非常停止状態（入力） *)
    RCON1_1_IN_ControllerReady : BOOL;  (* A(左側) RCON1_1 NG1上下降 コントローラ準備完了 *)
    RCON1_1_IN_Zone2 : BOOL;  (* A(左側) RCON1_1 NG1上下降 ゾーン2内 *)
    RCON1_1_IN_Zone1 : BOOL;  (* A(左側) RCON1_1 NG1上下降 ゾーン1内 *)
    RCON1_1_IN_CommandDone : BOOL;  (* A(左側) RCON1_1 NG1上下降 指令完了 *)
    RCON1_1_IN_OverloadWarning : BOOL;  (* A(左側) RCON1_1 NG1上下降 過負荷警告 *)
    RCON1_1_IN_PushMiss : BOOL;  (* A(左側) RCON1_1 NG1上下降 押付け空振り（未使用） *)
    RCON1_1_IN_ServoReady : BOOL;  (* A(左側) RCON1_1 NG1上下降 サーボON状態 *)
    RCON1_1_IN_Alarm : BOOL;  (* A(左側) RCON1_1 NG1上下降 軸異常 *)
    RCON1_1_Ready : BOOL;  (* A(左側) RCON1_1 NG1上下降 動作準備（安全許可とは別） *)
    RCON1_1_Error_Clear : BOOL;  (* A(左側) RCON1_1 NG1上下降 異常解除用予備（未接続） *)
    Error_M : ARRAY[0..99] OF Bool;  (* [3] FH A(左側) ST1; [9] FH A(左側) ST5; [10] FH B(右側) ST1; [11] FH B(右側) ST5; [12] A(左側) ST6 反転2 ワーク不一致 *)
    In_Sw_RESET : BOOL;
    RCON1_1_M : ARRAY[0..99] OF BOOL;  (* A(左側) RCON1_1 NG1上下降 開始・完了保持; [1] A(左側) RCON1_1 NG1上下降 開始指令保持; [2] A(左側) RCON1_1 NG1上下降 動作完了100ms *)
    TimerQ_In_SenCY_NG1_Pick_A_H : BOOL;
    Homing_Para_Stm : _sHOMING_REF;
END_VAR
VAR_EXTERNAL CONSTANT
    Stm_A_Rev_Axis000 : _sAXIS_REF;
END_VAR
VAR_EXTERNAL
    Stm_A_Rev_Axis000_OriginDone : BOOL;  (* A(左側) ST4 反転1 モータ原点復帰完了 *)
    Auto_A_Start : BOOL;
    HMI_Home_SW : BOOL;  (* HMI 原点復帰SW *)
    Stm_A_Rev_Axis000_Origin : BOOL;  (* A(左側) ST4 反転1 モータ原点復帰開始 *)
    Stm_A_Rev_Axis000_MovePos_Degree : LREAL;  (* A(左側)ステッピングモータ000 回転角度 *)
    Stm_A_Rev_Axis000_MoveAbsoluteDone : BOOL;  (* A(左側)ステッピング反転モータ1 絶対値位置決め 動作完了 *)
    Stm_A_Rev_Axis000_Auto : ARRAY[0..99] OF Bool;
    FH_A_ST5_Auto : BOOL;  (* A(左側) ST5 FH自動測定 *)
    FH_A_ST5_Manual : BOOL;  (* A(左側) ST5 FH手動測定 *)
    FH_A_ST5_Done : BOOL;  (* A(左側) ST5 画像検査完了 *)
    FH_Line1_Busy_1 : BOOL;  (* A(左側) 入力：ST5 処理実行中 *)
    FH_Line1_Command_Code_1 : DWORD;
    FH_Line1_Command_Completion_1 : BOOL;  (* A(左側) 入力：ST5 コマンド実行完了 *)
    FH_Line1_Command_Request_1 : BOOL;  (* A(左側) 出力：ST5 コマンド実行 *)
    FH_Line1_DINT_Result_Data_0_1 : DINT;  (* A(左側) 入力：ST5 判定0結果 *)
    FH_Line1_DINT_Result_Data_1_1 : DINT;  (* A(左側) 入力：ST5 判定1結果 *)
    FH_Line1_Error_Status_1 : BOOL;  (* A(左側) 入力：ST5 エラー信号 *)
    FH_Line1_Result_Notification_1 : BOOL;  (* A(左側) 入力：ST51 出力完了 *)
    FH_Line1_Trigger_1 : BOOL;  (* A(左側) 出力：ST5 測定トリガ *)
    FH_Line1_Trigger_Ready_1 : BOOL;  (* A(左側) 入力：ST5 測定準備完了 *)
    Homing_Para_Stm_Rev2 : _sHOMING_REF;  (* A(左側) ST6 反転2原点設定 *)
END_VAR
VAR_EXTERNAL CONSTANT
    Stm_A_Rev_Axis001 : _sAXIS_REF;
END_VAR
VAR_EXTERNAL
    Stm_A_Rev_Axis001_Auto : ARRAY[0..99] OF Bool;  (* A(左側) ST6 反転2自動指令; [1] A(左側) ST6 原点位置移動開始 *)
    Stm_A_Rev_Axis001_MoveAbsoluteDone : BOOL;  (* A(左側) ST6 反転2位置決め完了 *)
    Stm_A_Rev_Axis001_MovePos_Degree : LREAL;  (* A(左側) ST6 反転2指令角度 *)
    Stm_A_Rev_Axis001_Origin : BOOL;  (* A(左側) ST6 反転2 モータ原点復帰開始 *)
    Stm_A_Rev_Axis001_OriginDone : BOOL;  (* A(左側) ST6 反転2 モータ原点復帰完了 *)
    RCON1_2_IN_PositionDone : BOOL;  (* B(右側) RCON1_2 NG1上下降 位置決め完了 *)
    RCON1_2_IN_HomeDone : BOOL;  (* B(右側) RCON1_2 NG1上下降 原点復帰完了 *)
    RCON1_2_IN_Moving : BOOL;  (* B(右側) RCON1_2 NG1上下降 移動中 *)
    RCON1_2_IN_EmergencyStop : BOOL;  (* B(右側) RCON1_2 NG1上下降 非常停止状態（入力） *)
    RCON1_2_IN_ControllerReady : BOOL;  (* B(右側) RCON1_2 NG1上下降 コントローラ準備完了 *)
    RCON1_2_IN_Zone2 : BOOL;  (* B(右側) RCON1_2 NG1上下降 ゾーン2内 *)
    RCON1_2_IN_Zone1 : BOOL;  (* B(右側) RCON1_2 NG1上下降 ゾーン1内 *)
    RCON1_2_IN_CommandDone : BOOL;  (* B(右側) RCON1_2 NG1上下降 指令完了 *)
    RCON1_2_IN_OverloadWarning : BOOL;  (* B(右側) RCON1_2 NG1上下降 過負荷警告 *)
    RCON1_2_IN_PushMiss : BOOL;  (* B(右側) RCON1_2 NG1上下降 押付け空振り（未使用） *)
    RCON1_2_IN_ServoReady : BOOL;  (* B(右側) RCON1_2 NG1上下降 サーボON状態 *)
    RCON1_2_IN_Alarm : BOOL;  (* B(右側) RCON1_2 NG1上下降 軸異常 *)
    RCON1_2_Ready : BOOL;  (* B(右側) RCON1_2 NG1上下降 動作準備（安全許可とは別） *)
    RCON1_2_Error : BOOL;  (* B(右側) RCON1_2 NG1上下降 異常管理用予備（未接続） *)
    RCON1_2_Error_Clear : BOOL;  (* B(右側) RCON1_2 NG1上下降 異常解除用予備（未接続） *)
    RCON1_2_M : ARRAY[0..99] OF BOOL;  (* B(右側) RCON1_2 NG1上下降 開始・完了保持; [1] B(右側) RCON1_2 NG1上下降 開始指令保持; [2] B(右側) RCON1_2 NG1上下降 動作完了100ms *)
    RCON1_2_OUT_TargetPos_mm : LREAL;  (* B(右側) RCON1_2 NG1上下降 目標位置 [mm] *)
    RCON1_2_OUT_PositionBand_mm : LREAL;  (* B(右側) RCON1_2 NG1上下降 位置決め幅 [mm] *)
    RCON1_2_OUT_Speed_mm_s : LREAL;  (* B(右側) RCON1_2 NG1上下降 指令速度 [mm/s] *)
    RCON1_2_OUT_AccDec_G : LREAL;  (* B(右側) RCON1_2 NG1上下降 共通加減速度 [G] *)
    RCON1_2_OUT_PushLimit_pct : LREAL;  (* B(右側) RCON1_2 NG1上下降 押付け制限 [%]（未使用） *)
    RCON1_2_ActualPos_mm : LREAL;  (* B(右側) RCON1_2 NG1上下降 現在位置 [mm] *)
    RCON1_2_Current_mA : DINT;  (* B(右側) RCON1_2 NG1上下降 指令電流 [mA]（監視値） *)
    RCON1_2_ActualSpeed_mm_s : LREAL;  (* B(右側) RCON1_2 NG1上下降 現在速度 [mm/s・符号付き] *)
    RCON1_2_AlarmCode : UINT;  (* B(右側) RCON1_2 NG1上下降 軸異常コード *)
    RCON1_2_DataValid : BOOL;  (* B(右側) RCON1_2 NG1上下降 入力有効（安全許可ではない） *)
    RCON1_2_Auto : ARRAY[0..99] OF Bool;  (* B(右側) RCON1_2 NG1上下降 自動移動要求; [1] B(右側) RCON1_2 NG1上下降 自動要求1（外部接続用）; [2] B(右側) RCON1_2 NG1上下降 自動要求2（外部接続用）; [3] B(右側) RCON1_2 NG1上下降 自動要求3（外部接続用） *)
    RCON1_3_IN_PositionDone : BOOL;  (* A(左側) RCON1_3 SF/NG2送り 位置決め完了 *)
    RCON1_3_IN_HomeDone : BOOL;  (* A(左側) RCON1_3 SF/NG2送り 原点復帰完了 *)
    RCON1_3_IN_Moving : BOOL;  (* A(左側) RCON1_3 SF/NG2送り 移動中 *)
    RCON1_3_IN_EmergencyStop : BOOL;  (* A(左側) RCON1_3 SF/NG2送り 非常停止状態（入力） *)
    RCON1_3_IN_ControllerReady : BOOL;  (* A(左側) RCON1_3 SF/NG2送り コントローラ準備完了 *)
    RCON1_3_IN_Zone2 : BOOL;  (* A(左側) RCON1_3 SF/NG2送り ゾーン2内 *)
    RCON1_3_IN_Zone1 : BOOL;  (* A(左側) RCON1_3 SF/NG2送り ゾーン1内 *)
    RCON1_3_IN_CommandDone : BOOL;  (* A(左側) RCON1_3 SF/NG2送り 指令完了 *)
    RCON1_3_IN_OverloadWarning : BOOL;  (* A(左側) RCON1_3 SF/NG2送り 過負荷警告 *)
    RCON1_3_IN_PushMiss : BOOL;  (* A(左側) RCON1_3 SF/NG2送り 押付け空振り（未使用） *)
    RCON1_3_IN_ServoReady : BOOL;  (* A(左側) RCON1_3 SF/NG2送り サーボON状態 *)
    RCON1_3_IN_Alarm : BOOL;  (* A(左側) RCON1_3 SF/NG2送り 軸異常 *)
    RCON1_3_Ready : BOOL;  (* A(左側) RCON1_3 SF/NG2送り 動作準備（安全許可とは別） *)
    RCON1_3_Error : BOOL;  (* A(左側) RCON1_3 SF/NG2送り 異常管理用予備（未接続） *)
    RCON1_3_Error_Clear : BOOL;  (* A(左側) RCON1_3 SF/NG2送り 異常解除用予備（未接続） *)
    RCON1_3_M : ARRAY[0..99] OF BOOL;  (* A(左側) RCON1_3 SF/NG2送り 開始・完了保持; [1] A(左側) RCON1_3 SF/NG2送り 開始指令保持; [2] A(左側) RCON1_3 SF/NG2送り 動作完了100ms *)
    RCON1_3_OUT_TargetPos_mm : LREAL;  (* A(左側) RCON1_3 SF/NG2送り 目標位置 [mm] *)
    RCON1_3_OUT_PositionBand_mm : LREAL;  (* A(左側) RCON1_3 SF/NG2送り 位置決め幅 [mm] *)
    RCON1_3_OUT_Speed_mm_s : LREAL;  (* A(左側) RCON1_3 SF/NG2送り 指令速度 [mm/s] *)
    RCON1_3_OUT_AccDec_G : LREAL;  (* A(左側) RCON1_3 SF/NG2送り 共通加減速度 [G] *)
    RCON1_3_OUT_PushLimit_pct : LREAL;  (* A(左側) RCON1_3 SF/NG2送り 押付け制限 [%]（未使用） *)
    RCON1_3_ActualPos_mm : LREAL;  (* A(左側) RCON1_3 SF/NG2送り 現在位置 [mm] *)
    RCON1_3_Current_mA : DINT;  (* A(左側) RCON1_3 SF/NG2送り 指令電流 [mA]（監視値） *)
    RCON1_3_ActualSpeed_mm_s : LREAL;  (* A(左側) RCON1_3 SF/NG2送り 現在速度 [mm/s・符号付き] *)
    RCON1_3_AlarmCode : UINT;  (* A(左側) RCON1_3 SF/NG2送り 軸異常コード *)
    RCON1_3_DataValid : BOOL;  (* A(左側) RCON1_3 SF/NG2送り 入力有効（安全許可ではない） *)
    RCON1_3_Auto : ARRAY[0..99] OF Bool;  (* A(左側) RCON1_3 SF/NG2送り 自動移動要求; [1] A(左側) RCON1_3 SF/NG2送り 自動要求1（外部接続用）; [2] A(左側) RCON1_3 SF/NG2送り 自動要求2（外部接続用）; [3] A(左側) RCON1_3 SF/NG2送り 自動要求3（外部接続用） *)
    RCON1_4_IN_PositionDone : BOOL;  (* B(右側) RCON1_4 SF/NG2送り 位置決め完了 *)
    RCON1_4_IN_HomeDone : BOOL;  (* B(右側) RCON1_4 SF/NG2送り 原点復帰完了 *)
    RCON1_4_IN_Moving : BOOL;  (* B(右側) RCON1_4 SF/NG2送り 移動中 *)
    RCON1_4_IN_EmergencyStop : BOOL;  (* B(右側) RCON1_4 SF/NG2送り 非常停止状態（入力） *)
    RCON1_4_IN_ControllerReady : BOOL;  (* B(右側) RCON1_4 SF/NG2送り コントローラ準備完了 *)
    RCON1_4_IN_Zone2 : BOOL;  (* B(右側) RCON1_4 SF/NG2送り ゾーン2内 *)
    RCON1_4_IN_Zone1 : BOOL;  (* B(右側) RCON1_4 SF/NG2送り ゾーン1内 *)
    RCON1_4_IN_CommandDone : BOOL;  (* B(右側) RCON1_4 SF/NG2送り 指令完了 *)
    RCON1_4_IN_OverloadWarning : BOOL;  (* B(右側) RCON1_4 SF/NG2送り 過負荷警告 *)
    RCON1_4_IN_PushMiss : BOOL;  (* B(右側) RCON1_4 SF/NG2送り 押付け空振り（未使用） *)
    RCON1_4_IN_ServoReady : BOOL;  (* B(右側) RCON1_4 SF/NG2送り サーボON状態 *)
    RCON1_4_IN_Alarm : BOOL;  (* B(右側) RCON1_4 SF/NG2送り 軸異常 *)
    RCON1_4_Ready : BOOL;  (* B(右側) RCON1_4 SF/NG2送り 動作準備（安全許可とは別） *)
    RCON1_4_Error : BOOL;  (* B(右側) RCON1_4 SF/NG2送り 異常管理用予備（未接続） *)
    RCON1_4_Error_Clear : BOOL;  (* B(右側) RCON1_4 SF/NG2送り 異常解除用予備（未接続） *)
    RCON1_4_M : ARRAY[0..99] OF BOOL;  (* B(右側) RCON1_4 SF/NG2送り 開始・完了保持; [1] B(右側) RCON1_4 SF/NG2送り 開始指令保持; [2] B(右側) RCON1_4 SF/NG2送り 動作完了100ms *)
    RCON1_4_OUT_TargetPos_mm : LREAL;  (* B(右側) RCON1_4 SF/NG2送り 目標位置 [mm] *)
    RCON1_4_OUT_PositionBand_mm : LREAL;  (* B(右側) RCON1_4 SF/NG2送り 位置決め幅 [mm] *)
    RCON1_4_OUT_Speed_mm_s : LREAL;  (* B(右側) RCON1_4 SF/NG2送り 指令速度 [mm/s] *)
    RCON1_4_OUT_AccDec_G : LREAL;  (* B(右側) RCON1_4 SF/NG2送り 共通加減速度 [G] *)
    RCON1_4_OUT_PushLimit_pct : LREAL;  (* B(右側) RCON1_4 SF/NG2送り 押付け制限 [%]（未使用） *)
    RCON1_4_ActualPos_mm : LREAL;  (* B(右側) RCON1_4 SF/NG2送り 現在位置 [mm] *)
    RCON1_4_Current_mA : DINT;  (* B(右側) RCON1_4 SF/NG2送り 指令電流 [mA]（監視値） *)
    RCON1_4_ActualSpeed_mm_s : LREAL;  (* B(右側) RCON1_4 SF/NG2送り 現在速度 [mm/s・符号付き] *)
    RCON1_4_AlarmCode : UINT;  (* B(右側) RCON1_4 SF/NG2送り 軸異常コード *)
    RCON1_4_DataValid : BOOL;  (* B(右側) RCON1_4 SF/NG2送り 入力有効（安全許可ではない） *)
    RCON1_4_Auto : ARRAY[0..99] OF Bool;  (* B(右側) RCON1_4 SF/NG2送り 自動移動要求; [1] B(右側) RCON1_4 SF/NG2送り 自動要求1（外部接続用）; [2] B(右側) RCON1_4 SF/NG2送り 自動要求2（外部接続用）; [3] B(右側) RCON1_4 SF/NG2送り 自動要求3（外部接続用） *)
    RCON1_5_IN_PositionDone : BOOL;  (* A(左側) RCON1_5 SF/NG2上下降 位置決め完了 *)
    RCON1_5_IN_HomeDone : BOOL;  (* A(左側) RCON1_5 SF/NG2上下降 原点復帰完了 *)
    RCON1_5_IN_Moving : BOOL;  (* A(左側) RCON1_5 SF/NG2上下降 移動中 *)
    RCON1_5_IN_EmergencyStop : BOOL;  (* A(左側) RCON1_5 SF/NG2上下降 非常停止状態（入力） *)
    RCON1_5_IN_ControllerReady : BOOL;  (* A(左側) RCON1_5 SF/NG2上下降 コントローラ準備完了 *)
    RCON1_5_IN_Zone2 : BOOL;  (* A(左側) RCON1_5 SF/NG2上下降 ゾーン2内 *)
    RCON1_5_IN_Zone1 : BOOL;  (* A(左側) RCON1_5 SF/NG2上下降 ゾーン1内 *)
    RCON1_5_IN_CommandDone : BOOL;  (* A(左側) RCON1_5 SF/NG2上下降 指令完了 *)
    RCON1_5_IN_OverloadWarning : BOOL;  (* A(左側) RCON1_5 SF/NG2上下降 過負荷警告 *)
    RCON1_5_IN_PushMiss : BOOL;  (* A(左側) RCON1_5 SF/NG2上下降 押付け空振り（未使用） *)
    RCON1_5_IN_ServoReady : BOOL;  (* A(左側) RCON1_5 SF/NG2上下降 サーボON状態 *)
    RCON1_5_IN_Alarm : BOOL;  (* A(左側) RCON1_5 SF/NG2上下降 軸異常 *)
    RCON1_5_Ready : BOOL;  (* A(左側) RCON1_5 SF/NG2上下降 動作準備（安全許可とは別） *)
    RCON1_5_Error : BOOL;  (* A(左側) RCON1_5 SF/NG2上下降 異常管理用予備（未接続） *)
    RCON1_5_Error_Clear : BOOL;  (* A(左側) RCON1_5 SF/NG2上下降 異常解除用予備（未接続） *)
    RCON1_5_M : ARRAY[0..99] OF BOOL;  (* A(左側) RCON1_5 SF/NG2上下降 開始・完了保持; [1] A(左側) RCON1_5 SF/NG2上下降 開始指令保持; [2] A(左側) RCON1_5 SF/NG2上下降 動作完了100ms *)
    RCON1_5_OUT_TargetPos_mm : LREAL;  (* A(左側) RCON1_5 SF/NG2上下降 目標位置 [mm] *)
    RCON1_5_OUT_PositionBand_mm : LREAL;  (* A(左側) RCON1_5 SF/NG2上下降 位置決め幅 [mm] *)
    RCON1_5_OUT_Speed_mm_s : LREAL;  (* A(左側) RCON1_5 SF/NG2上下降 指令速度 [mm/s] *)
    RCON1_5_OUT_AccDec_G : LREAL;  (* A(左側) RCON1_5 SF/NG2上下降 共通加減速度 [G] *)
    RCON1_5_OUT_PushLimit_pct : LREAL;  (* A(左側) RCON1_5 SF/NG2上下降 押付け制限 [%]（未使用） *)
    RCON1_5_ActualPos_mm : LREAL;  (* A(左側) RCON1_5 SF/NG2上下降 現在位置 [mm] *)
    RCON1_5_Current_mA : DINT;  (* A(左側) RCON1_5 SF/NG2上下降 指令電流 [mA]（監視値） *)
    RCON1_5_ActualSpeed_mm_s : LREAL;  (* A(左側) RCON1_5 SF/NG2上下降 現在速度 [mm/s・符号付き] *)
    RCON1_5_AlarmCode : UINT;  (* A(左側) RCON1_5 SF/NG2上下降 軸異常コード *)
    RCON1_5_DataValid : BOOL;  (* A(左側) RCON1_5 SF/NG2上下降 入力有効（安全許可ではない） *)
    RCON1_5_Auto : ARRAY[0..99] OF Bool;  (* A(左側) RCON1_5 SF/NG2上下降 自動移動要求; [1] A(左側) RCON1_5 SF/NG2上下降 自動要求1（外部接続用）; [2] A(左側) RCON1_5 SF/NG2上下降 自動要求2（外部接続用）; [3] A(左側) RCON1_5 SF/NG2上下降 自動要求3（外部接続用） *)
    RCON1_6_IN_PositionDone : BOOL;  (* B(右側) RCON1_6 SF/NG2上下降 位置決め完了 *)
    RCON1_6_IN_HomeDone : BOOL;  (* B(右側) RCON1_6 SF/NG2上下降 原点復帰完了 *)
    RCON1_6_IN_Moving : BOOL;  (* B(右側) RCON1_6 SF/NG2上下降 移動中 *)
    RCON1_6_IN_EmergencyStop : BOOL;  (* B(右側) RCON1_6 SF/NG2上下降 非常停止状態（入力） *)
    RCON1_6_IN_ControllerReady : BOOL;  (* B(右側) RCON1_6 SF/NG2上下降 コントローラ準備完了 *)
    RCON1_6_IN_Zone2 : BOOL;  (* B(右側) RCON1_6 SF/NG2上下降 ゾーン2内 *)
    RCON1_6_IN_Zone1 : BOOL;  (* B(右側) RCON1_6 SF/NG2上下降 ゾーン1内 *)
    RCON1_6_IN_CommandDone : BOOL;  (* B(右側) RCON1_6 SF/NG2上下降 指令完了 *)
    RCON1_6_IN_OverloadWarning : BOOL;  (* B(右側) RCON1_6 SF/NG2上下降 過負荷警告 *)
    RCON1_6_IN_PushMiss : BOOL;  (* B(右側) RCON1_6 SF/NG2上下降 押付け空振り（未使用） *)
    RCON1_6_IN_ServoReady : BOOL;  (* B(右側) RCON1_6 SF/NG2上下降 サーボON状態 *)
    RCON1_6_IN_Alarm : BOOL;  (* B(右側) RCON1_6 SF/NG2上下降 軸異常 *)
    RCON1_6_Ready : BOOL;  (* B(右側) RCON1_6 SF/NG2上下降 動作準備（安全許可とは別） *)
    RCON1_6_Error : BOOL;  (* B(右側) RCON1_6 SF/NG2上下降 異常管理用予備（未接続） *)
    RCON1_6_Error_Clear : BOOL;  (* B(右側) RCON1_6 SF/NG2上下降 異常解除用予備（未接続） *)
    RCON1_6_M : ARRAY[0..99] OF BOOL;  (* B(右側) RCON1_6 SF/NG2上下降 開始・完了保持; [1] B(右側) RCON1_6 SF/NG2上下降 開始指令保持; [2] B(右側) RCON1_6 SF/NG2上下降 動作完了100ms *)
    RCON1_6_OUT_TargetPos_mm : LREAL;  (* B(右側) RCON1_6 SF/NG2上下降 目標位置 [mm] *)
    RCON1_6_OUT_PositionBand_mm : LREAL;  (* B(右側) RCON1_6 SF/NG2上下降 位置決め幅 [mm] *)
    RCON1_6_OUT_Speed_mm_s : LREAL;  (* B(右側) RCON1_6 SF/NG2上下降 指令速度 [mm/s] *)
    RCON1_6_OUT_AccDec_G : LREAL;  (* B(右側) RCON1_6 SF/NG2上下降 共通加減速度 [G] *)
    RCON1_6_OUT_PushLimit_pct : LREAL;  (* B(右側) RCON1_6 SF/NG2上下降 押付け制限 [%]（未使用） *)
    RCON1_6_ActualPos_mm : LREAL;  (* B(右側) RCON1_6 SF/NG2上下降 現在位置 [mm] *)
    RCON1_6_Current_mA : DINT;  (* B(右側) RCON1_6 SF/NG2上下降 指令電流 [mA]（監視値） *)
    RCON1_6_ActualSpeed_mm_s : LREAL;  (* B(右側) RCON1_6 SF/NG2上下降 現在速度 [mm/s・符号付き] *)
    RCON1_6_AlarmCode : UINT;  (* B(右側) RCON1_6 SF/NG2上下降 軸異常コード *)
    RCON1_6_DataValid : BOOL;  (* B(右側) RCON1_6 SF/NG2上下降 入力有効（安全許可ではない） *)
    RCON1_6_Auto : ARRAY[0..99] OF Bool;  (* B(右側) RCON1_6 SF/NG2上下降 自動移動要求; [1] B(右側) RCON1_6 SF/NG2上下降 自動要求1（外部接続用）; [2] B(右側) RCON1_6 SF/NG2上下降 自動要求2（外部接続用）; [3] B(右側) RCON1_6 SF/NG2上下降 自動要求3（外部接続用） *)
    TimerQ_In_SenCY_NG1_Pick_B_H : BOOL;  (* 【X428】B(右側) NG1ピックアップ戻 *)
END_VAR
VAR
    _e1 : R_TRIG;
    _e2 : R_TRIG;
    _e3 : R_TRIG;
    _p4 : BOOL;
    _e5 : R_TRIG;
    _e6 : R_TRIG;
    _e7 : R_TRIG;
    _p8 : BOOL;
    _e9 : R_TRIG;
    _e10 : R_TRIG;
    _e11 : R_TRIG;
    _p12 : BOOL;
    _e13 : R_TRIG;
    _e14 : R_TRIG;
    _e15 : R_TRIG;
    _p16 : BOOL;
    _e17 : R_TRIG;
    _e18 : R_TRIG;
    _e19 : R_TRIG;
    _p20 : BOOL;
    _e21 : R_TRIG;
    _e22 : R_TRIG;
    _e23 : R_TRIG;
    _p24 : BOOL;
    _e25 : R_TRIG;
    _p26 : BOOL;
    _e27 : R_TRIG;
    _p28 : BOOL;
    _e29 : R_TRIG;
    _p30 : BOOL;
    _e31 : R_TRIG;
    _e32 : R_TRIG;
    _p33 : BOOL;
    _e34 : R_TRIG;
    _e35 : R_TRIG;
    _p36 : BOOL;
    _p37 : BOOL;
    _e38 : R_TRIG;
    _p39 : BOOL;
    _e40 : R_TRIG;
    _p41 : BOOL;
    _e42 : R_TRIG;
    _p43 : BOOL;
    _e44 : R_TRIG;
    _e45 : R_TRIG;
    _p46 : BOOL;
    _e47 : R_TRIG;
    _e48 : R_TRIG;
    _p49 : BOOL;
    _p50 : BOOL;
    _p51 : BOOL;
    _p52 : BOOL;
END_VAR

(* Section RCON_IAI: ladder, written here as Structured Text *)

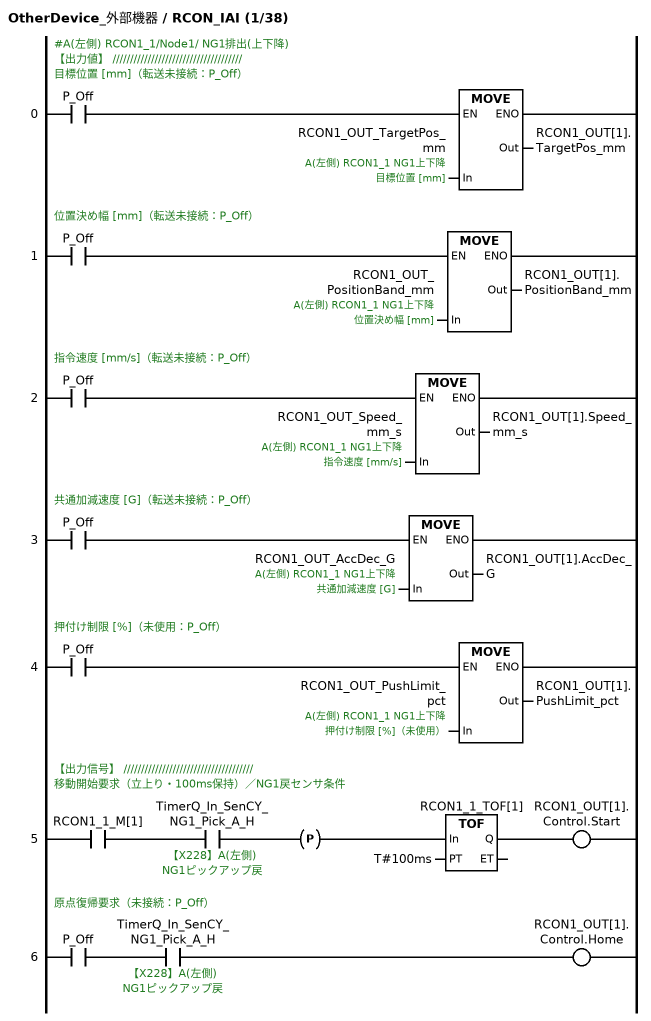
(* Rung 0: #A(左側) RCON1_1/Node1/ NG1排出(上下降) / 【出力値】 ///////////////////////////////////// / 目標位置 [mm]（転送未接続：P_Off） *)
IF P_Off THEN RCON1_OUT[1].TargetPos_mm := RCON1_OUT_TargetPos_mm; END_IF;
(* Rung 1: 位置決め幅 [mm]（転送未接続：P_Off） *)
IF P_Off THEN RCON1_OUT[1].PositionBand_mm := RCON1_OUT_PositionBand_mm; END_IF;
(* Rung 2: 指令速度 [mm/s]（転送未接続：P_Off） *)
IF P_Off THEN RCON1_OUT[1].Speed_mm_s := RCON1_OUT_Speed_mm_s; END_IF;
(* Rung 3: 共通加減速度 [G]（転送未接続：P_Off） *)
IF P_Off THEN RCON1_OUT[1].AccDec_G := RCON1_OUT_AccDec_G; END_IF;
(* Rung 4: 押付け制限 [%]（未使用：P_Off） *)
IF P_Off THEN RCON1_OUT[1].PushLimit_pct := RCON1_OUT_PushLimit_pct; END_IF;
(* Rung 5: 【出力信号】 ///////////////////////////////////// / 移動開始要求（立上り・100ms保持）／NG1戻センサ条件 *)
_e1(CLK := RCON1_1_M[1] AND TimerQ_In_SenCY_NG1_Pick_A_H);
RCON1_1_TOF[1](In := _e1.Q, PT := T#100ms);
RCON1_OUT[1].Control.Start := RCON1_1_TOF[1].Q;
(* Rung 6: 原点復帰要求（未接続：P_Off） *)
RCON1_OUT[1].Control.Home := P_Off AND TimerQ_In_SenCY_NG1_Pick_A_H;

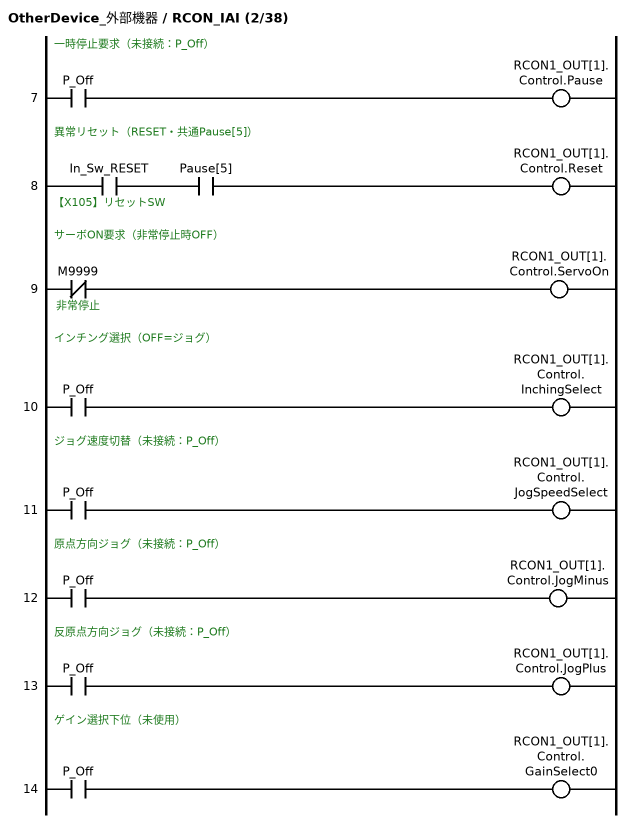
(* Rung 7: 一時停止要求（未接続：P_Off） *)
RCON1_OUT[1].Control.Pause := P_Off;
(* Rung 8: 異常リセット（RESET・共通Pause[5]） *)
RCON1_OUT[1].Control.Reset := In_Sw_RESET AND Pause[5];
(* Rung 9: サーボON要求（非常停止時OFF） *)
RCON1_OUT[1].Control.ServoOn := NOT M9999;
(* Rung 10: インチング選択（OFF=ジョグ） *)
RCON1_OUT[1].Control.InchingSelect := P_Off;
(* Rung 11: ジョグ速度切替（未接続：P_Off） *)
RCON1_OUT[1].Control.JogSpeedSelect := P_Off;
(* Rung 12: 原点方向ジョグ（未接続：P_Off） *)
RCON1_OUT[1].Control.JogMinus := P_Off;
(* Rung 13: 反原点方向ジョグ（未接続：P_Off） *)
RCON1_OUT[1].Control.JogPlus := P_Off;
(* Rung 14: ゲイン選択下位（未使用） *)
RCON1_OUT[1].Control.GainSelect0 := P_Off;

